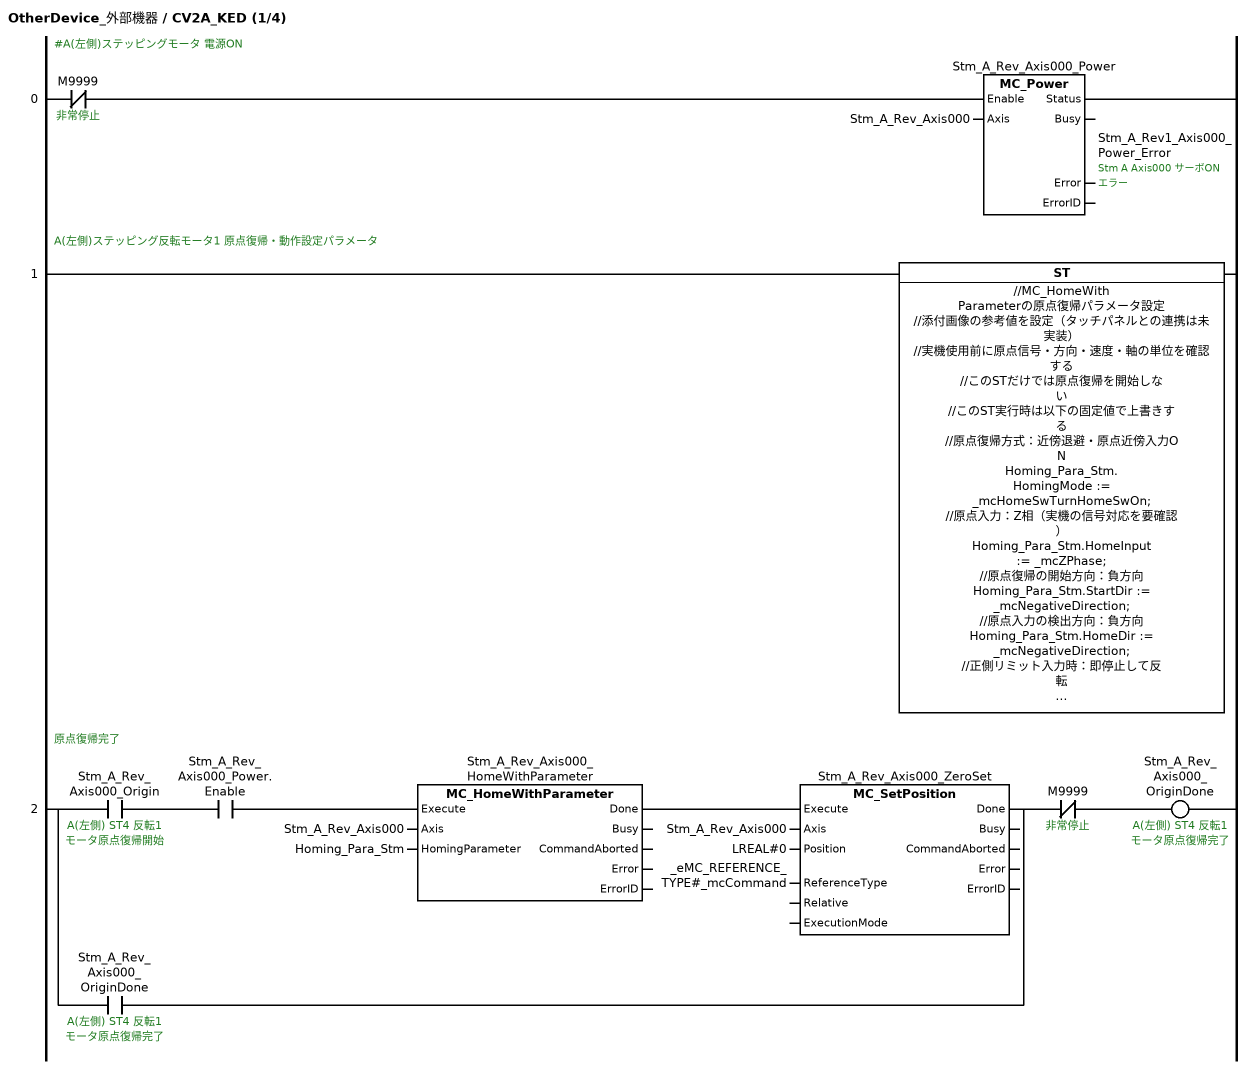
(* [picture p143: OtherDevice_外部機器 / CV2A_KED, rungs 0-2] *)
(* Rung 0: #A(左側)ステッピングモータ 電源ON *)
Stm_A_Rev_Axis000_Power(Enable := NOT M9999, Axis := Stm_A_Rev_Axis000, Error => Stm_A_Rev1_Axis000_Power_Error);
(* Rung 1: A(左側)ステッピング反転モータ1 原点復帰・動作設定パラメータ *)
//MC_HomeWithParameterの原点復帰パラメータ設定
//添付画像の参考値を設定（タッチパネルとの連携は未実装）
//実機使用前に原点信号・方向・速度・軸の単位を確認する
//このSTだけでは原点復帰を開始しない
//このST実行時は以下の固定値で上書きする

//原点復帰方式：近傍退避・原点近傍入力ON
Homing_Para_Stm.HomingMode := _mcHomeSwTurnHomeSwOn;
//原点入力：Z相（実機の信号対応を要確認）
Homing_Para_Stm.HomeInput := _mcZPhase;
//原点復帰の開始方向：負方向
Homing_Para_Stm.StartDir := _mcNegativeDirection;
//原点入力の検出方向：負方向
Homing_Para_Stm.HomeDir := _mcNegativeDirection;
//正側リミット入力時：即停止して反転
Homing_Para_Stm.PosiLmtMode := _mcRevImmediateStop;
//負側リミット入力時：即停止して反転
Homing_Para_Stm.NegaLmtMode := _mcRevImmediateStop;

//原点復帰速度 [指令単位/s]
Homing_Para_Stm.Vel := LREAL#40;
//原点近傍での接近速度 [指令単位/s]
Homing_Para_Stm.ApproachVel := LREAL#1;
//原点復帰の加速度 [指令単位/s^2]
Homing_Para_Stm.Acc := LREAL#100;
//原点復帰の減速度 [指令単位/s^2]
Homing_Para_Stm.Dec := LREAL#200;
//ジャーク [指令単位/s^3]：0はジャーク制御なし
Homing_Para_Stm.Jerk := LREAL#0;

//原点入力マスク距離 [指令単位]：今回の方式では未使用
Homing_Para_Stm.Mask := LREAL#0;
//原点確定後の現在位置 [指令単位]
Homing_Para_Stm.Offset := LREAL#0;
//押当て時間 [ms]：今回の方式では未使用
Homing_Para_Stm.PushTime := UINT#0;
//原点検出後の補正移動量 [指令単位]：0は補正移動なし
Homing_Para_Stm.Compensation := LREAL#0;
//原点補正移動時の速度 [指令単位/s]
Homing_Para_Stm.CompensationVel := LREAL#10;
(* Rung 2: 原点復帰完了 *)
Stm_A_Rev_Axis000_HomeWithParameter(Execute := Stm_A_Rev_Axis000_Origin AND Stm_A_Rev_Axis000_Power.Enable, Axis := Stm_A_Rev_Axis000, HomingParameter := Homing_Para_Stm);
Stm_A_Rev_Axis000_ZeroSet(Execute := Stm_A_Rev_Axis000_HomeWithParameter.Done, Axis := Stm_A_Rev_Axis000, Position := LREAL#0, ReferenceType := _eMC_REFERENCE_TYPE#_mcCommand);
Stm_A_Rev_Axis000_OriginDone := (Stm_A_Rev_Axis000_ZeroSet.Done OR Stm_A_Rev_Axis000_OriginDone) AND NOT M9999;

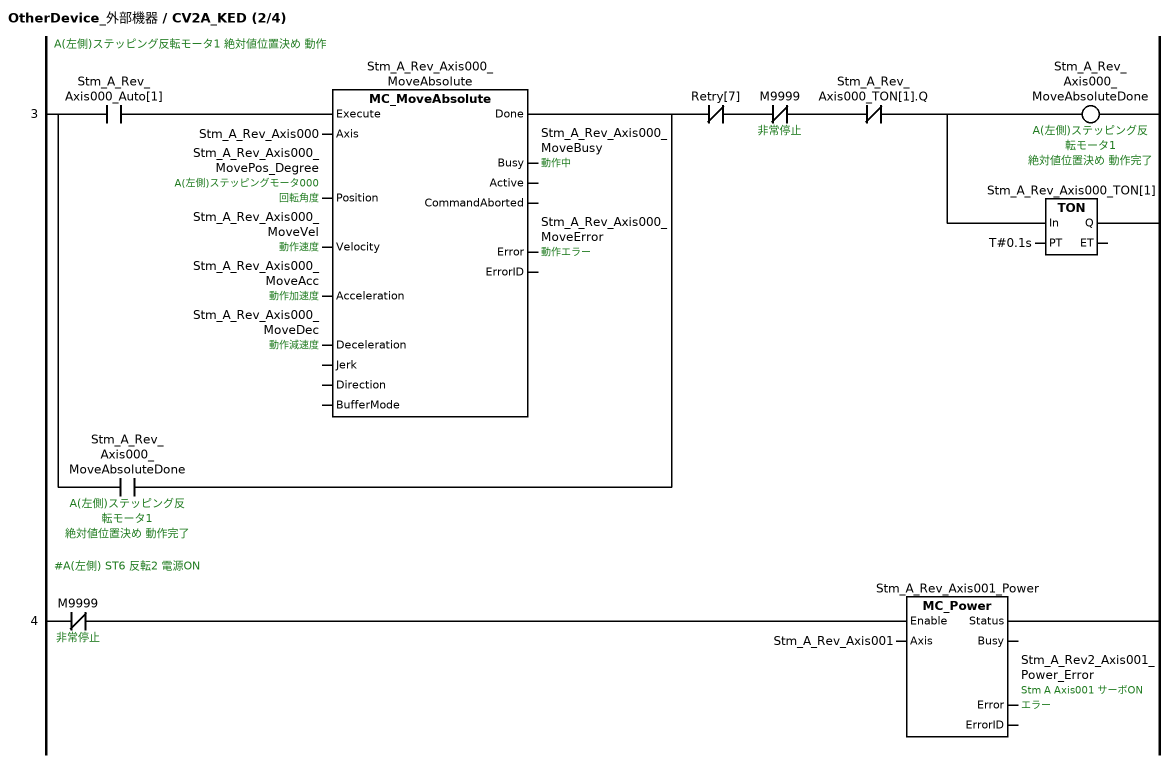
(* Rung 3: A(左側)ステッピング反転モータ1 絶対値位置決め 動作 *)
Stm_A_Rev_Axis000_MoveAbsolute(Execute := Stm_A_Rev_Axis000_Auto[1], Axis := Stm_A_Rev_Axis000, Position := Stm_A_Rev_Axis000_MovePos_Degree, Velocity := Stm_A_Rev_Axis000_MoveVel, Acceleration := Stm_A_Rev_Axis000_MoveAcc, Deceleration := Stm_A_Rev_Axis000_MoveDec, Busy => Stm_A_Rev_Axis000_MoveBusy, Error => Stm_A_Rev_Axis000_MoveError);
_p71 := (Stm_A_Rev_Axis000_MoveAbsolute.Done OR Stm_A_Rev_Axis000_MoveAbsoluteDone) AND NOT Retry[7] AND NOT M9999 AND NOT Stm_A_Rev_Axis000_TON[1].Q;
Stm_A_Rev_Axis000_MoveAbsoluteDone := _p71;
Stm_A_Rev_Axis000_TON[1](In := _p71, PT := T#0.1s);
(* Rung 4: #A(左側) ST6 反転2 電源ON *)
Stm_A_Rev_Axis001_Power(Enable := NOT M9999, Axis := Stm_A_Rev_Axis001, Error => Stm_A_Rev2_Axis001_Power_Error);

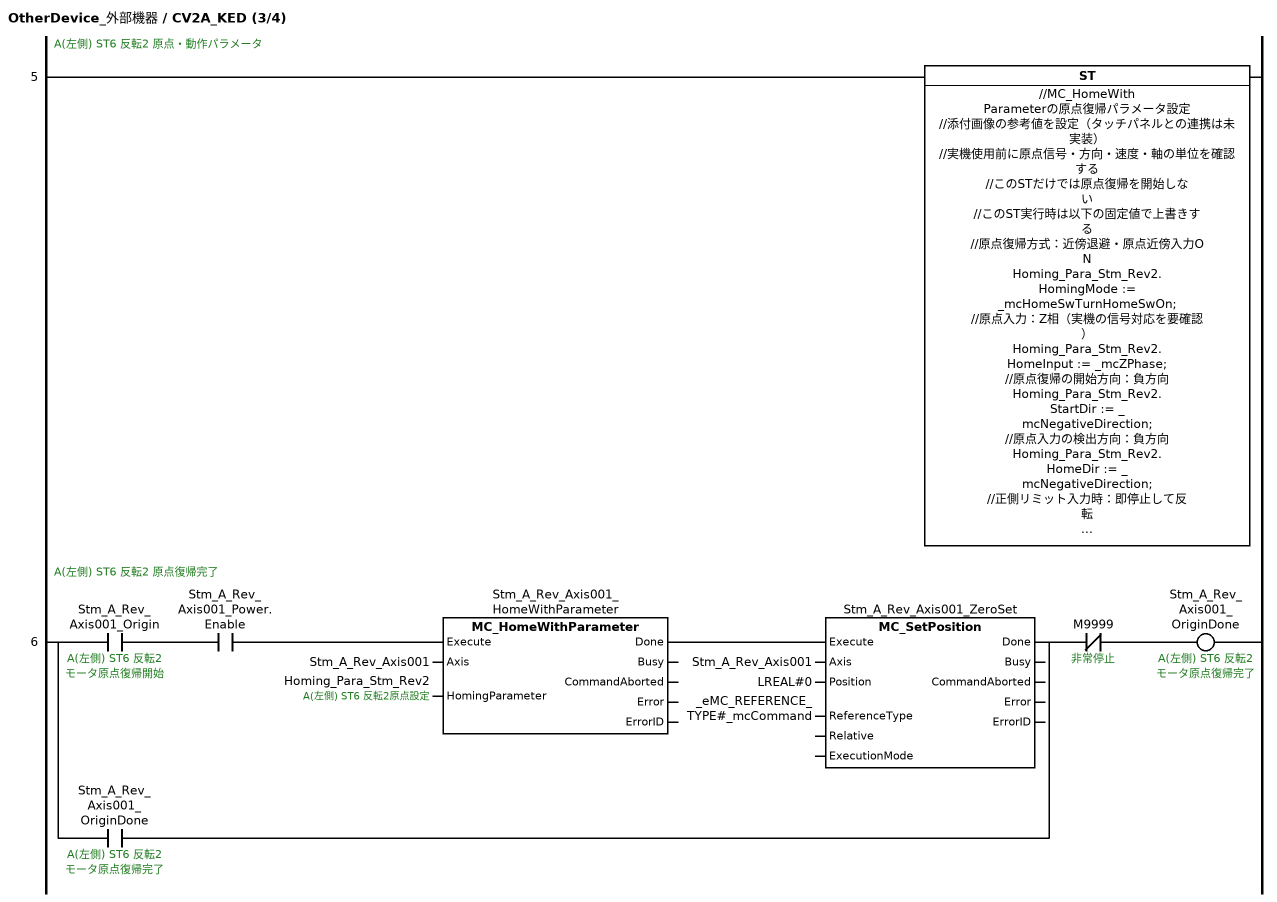
(* Rung 5: A(左側) ST6 反転2 原点・動作パラメータ *)
//MC_HomeWithParameterの原点復帰パラメータ設定
//添付画像の参考値を設定（タッチパネルとの連携は未実装）
//実機使用前に原点信号・方向・速度・軸の単位を確認する
//このSTだけでは原点復帰を開始しない
//このST実行時は以下の固定値で上書きする

//原点復帰方式：近傍退避・原点近傍入力ON
Homing_Para_Stm_Rev2.HomingMode := _mcHomeSwTurnHomeSwOn;
//原点入力：Z相（実機の信号対応を要確認）
Homing_Para_Stm_Rev2.HomeInput := _mcZPhase;
//原点復帰の開始方向：負方向
Homing_Para_Stm_Rev2.StartDir := _mcNegativeDirection;
//原点入力の検出方向：負方向
Homing_Para_Stm_Rev2.HomeDir := _mcNegativeDirection;
//正側リミット入力時：即停止して反転
Homing_Para_Stm_Rev2.PosiLmtMode := _mcRevImmediateStop;
//負側リミット入力時：即停止して反転
Homing_Para_Stm_Rev2.NegaLmtMode := _mcRevImmediateStop;

//原点復帰速度 [指令単位/s]
Homing_Para_Stm_Rev2.Vel := LREAL#40;
//原点近傍での接近速度 [指令単位/s]
Homing_Para_Stm_Rev2.ApproachVel := LREAL#1;
//原点復帰の加速度 [指令単位/s^2]
Homing_Para_Stm_Rev2.Acc := LREAL#100;
//原点復帰の減速度 [指令単位/s^2]
Homing_Para_Stm_Rev2.Dec := LREAL#200;
//ジャーク [指令単位/s^3]：0はジャーク制御なし
Homing_Para_Stm_Rev2.Jerk := LREAL#0;

//原点入力マスク距離 [指令単位]：今回の方式では未使用
Homing_Para_Stm_Rev2.Mask := LREAL#0;
//原点確定後の現在位置 [指令単位]
Homing_Para_Stm_Rev2.Offset := LREAL#0;
//押当て時間 [ms]：今回の方式では未使用
Homing_Para_Stm_Rev2.PushTime := UINT#0;
//原点検出後の補正移動量 [指令単位]：0は補正移動なし
Homing_Para_Stm_Rev2.Compensation := LREAL#0;
//原点補正移動時の速度 [指令単位/s]
Homing_Para_Stm_Rev2.CompensationVel := LREAL#10;
(* Rung 6: A(左側) ST6 反転2 原点復帰完了 *)
Stm_A_Rev_Axis001_HomeWithParameter(Execute := Stm_A_Rev_Axis001_Origin AND Stm_A_Rev_Axis001_Power.Enable, Axis := Stm_A_Rev_Axis001, HomingParameter := Homing_Para_Stm_Rev2);
Stm_A_Rev_Axis001_ZeroSet(Execute := Stm_A_Rev_Axis001_HomeWithParameter.Done, Axis := Stm_A_Rev_Axis001, Position := LREAL#0, ReferenceType := _eMC_REFERENCE_TYPE#_mcCommand);
Stm_A_Rev_Axis001_OriginDone := (Stm_A_Rev_Axis001_ZeroSet.Done OR Stm_A_Rev_Axis001_OriginDone) AND NOT M9999;

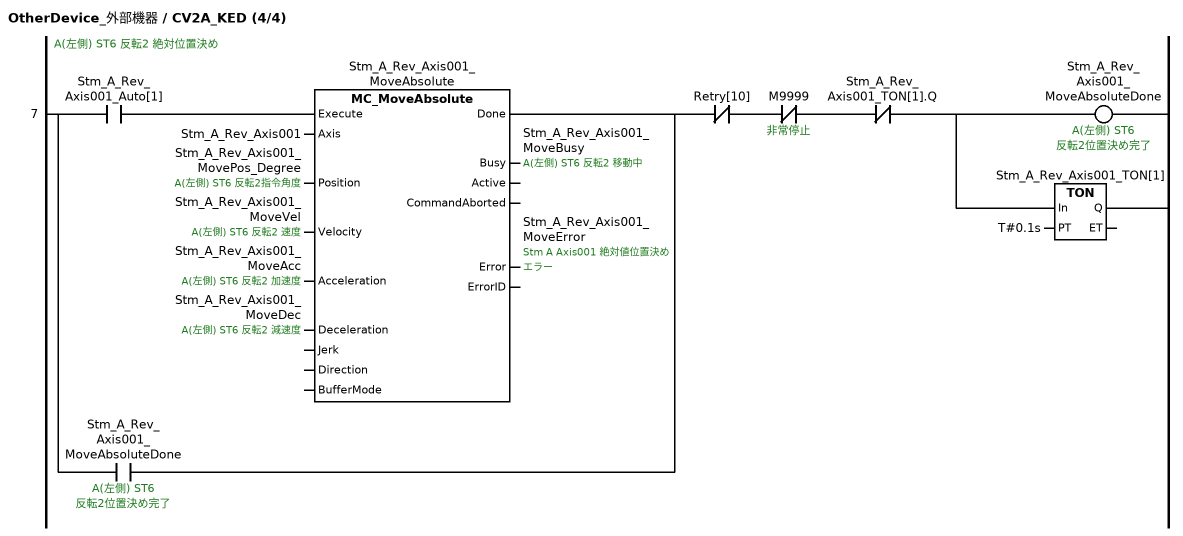
(* Rung 7: A(左側) ST6 反転2 絶対位置決め *)
Stm_A_Rev_Axis001_MoveAbsolute(Execute := Stm_A_Rev_Axis001_Auto[1], Axis := Stm_A_Rev_Axis001, Position := Stm_A_Rev_Axis001_MovePos_Degree, Velocity := Stm_A_Rev_Axis001_MoveVel, Acceleration := Stm_A_Rev_Axis001_MoveAcc, Deceleration := Stm_A_Rev_Axis001_MoveDec, Busy => Stm_A_Rev_Axis001_MoveBusy, Error => Stm_A_Rev_Axis001_MoveError);
_p72 := (Stm_A_Rev_Axis001_MoveAbsolute.Done OR Stm_A_Rev_Axis001_MoveAbsoluteDone) AND NOT Retry[10] AND NOT M9999 AND NOT Stm_A_Rev_Axis001_TON[1].Q;
Stm_A_Rev_Axis001_MoveAbsoluteDone := _p72;
Stm_A_Rev_Axis001_TON[1](In := _p72, PT := T#0.1s);

(* Section HMI: ladder, written here as Structured Text *)

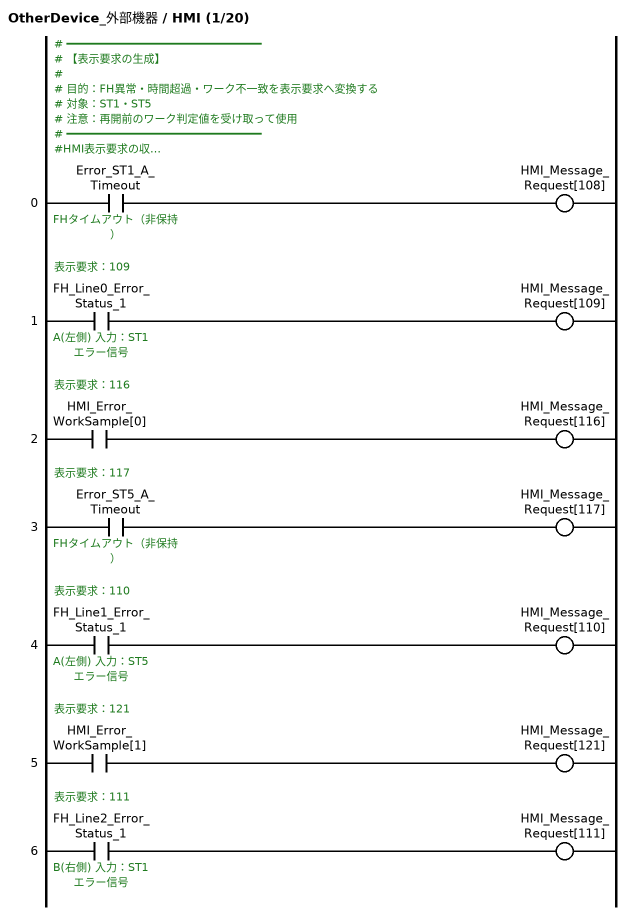
(* Rung 0: # ━━━━━━━━━━━━━━━━━━━━━━━━━━━━━━ / # 【表示要求の生成】 / # / # 目的：FH異常・時間超過・ワーク不一致を表示要求へ変換する / # 対象：ST1・ST5 / # 注意：再開前のワーク判定値を受け取って使用 / # ━━━━━━━━━━━━━━━━━━━━━━━━━━━━━━ / #HMI表示要求の収集 / 実行順維持のため、異常判定後・再開処理前 / 表示要求：108 *)
HMI_Message_Request[108] := Error_ST1_A_Timeout;
(* Rung 1: 表示要求：109 *)
HMI_Message_Request[109] := FH_Line0_Error_Status_1;
(* Rung 2: 表示要求：116 *)
HMI_Message_Request[116] := HMI_Error_WorkSample[0];
(* Rung 3: 表示要求：117 *)
HMI_Message_Request[117] := Error_ST5_A_Timeout;
(* Rung 4: 表示要求：110 *)
HMI_Message_Request[110] := FH_Line1_Error_Status_1;
(* Rung 5: 表示要求：121 *)
HMI_Message_Request[121] := HMI_Error_WorkSample[1];
(* Rung 6: 表示要求：111 *)
HMI_Message_Request[111] := FH_Line2_Error_Status_1;

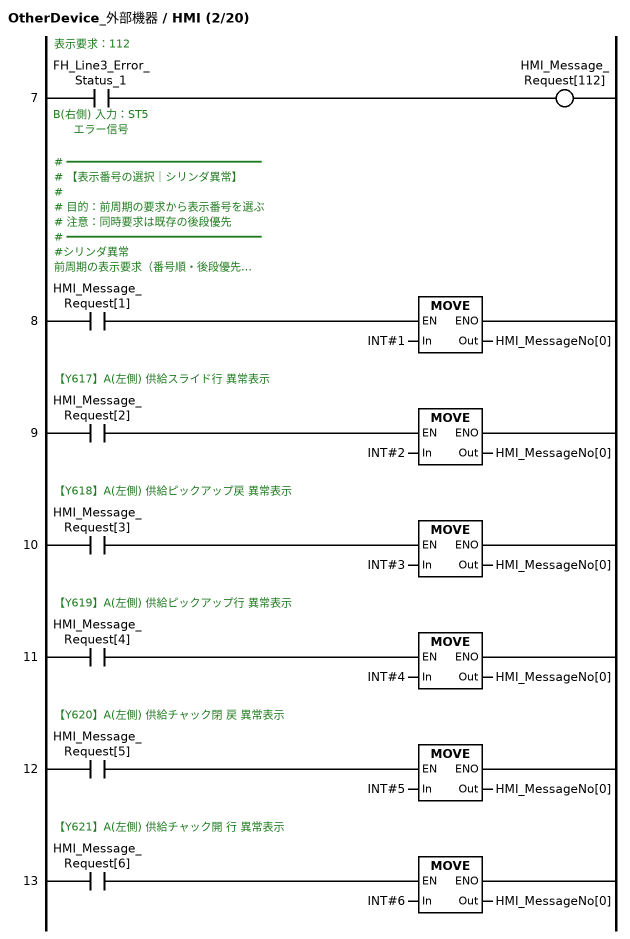
(* Rung 7: 表示要求：112 *)
HMI_Message_Request[112] := FH_Line3_Error_Status_1;
(* Rung 8: # ━━━━━━━━━━━━━━━━━━━━━━━━━━━━━━ / # 【表示番号の選択｜シリンダ異常】 / # / # 目的：前周期の要求から表示番号を選ぶ / # 注意：同時要求は既存の後段優先 / # ━━━━━━━━━━━━━━━━━━━━━━━━━━━━━━ / #シリンダ異常 / 前周期の表示要求（番号順・後段優先） / 【Y616】A(左側) 供給スライド戻 異常表示 *)
IF HMI_Message_Request[1] THEN HMI_MessageNo[0] := INT#1; END_IF;
(* Rung 9: 【Y617】A(左側) 供給スライド行 異常表示 *)
IF HMI_Message_Request[2] THEN HMI_MessageNo[0] := INT#2; END_IF;
(* Rung 10: 【Y618】A(左側) 供給ピックアップ戻 異常表示 *)
IF HMI_Message_Request[3] THEN HMI_MessageNo[0] := INT#3; END_IF;
(* Rung 11: 【Y619】A(左側) 供給ピックアップ行 異常表示 *)
IF HMI_Message_Request[4] THEN HMI_MessageNo[0] := INT#4; END_IF;
(* Rung 12: 【Y620】A(左側) 供給チャック閉 戻 異常表示 *)
IF HMI_Message_Request[5] THEN HMI_MessageNo[0] := INT#5; END_IF;
(* Rung 13: 【Y621】A(左側) 供給チャック開 行 異常表示 *)
IF HMI_Message_Request[6] THEN HMI_MessageNo[0] := INT#6; END_IF;

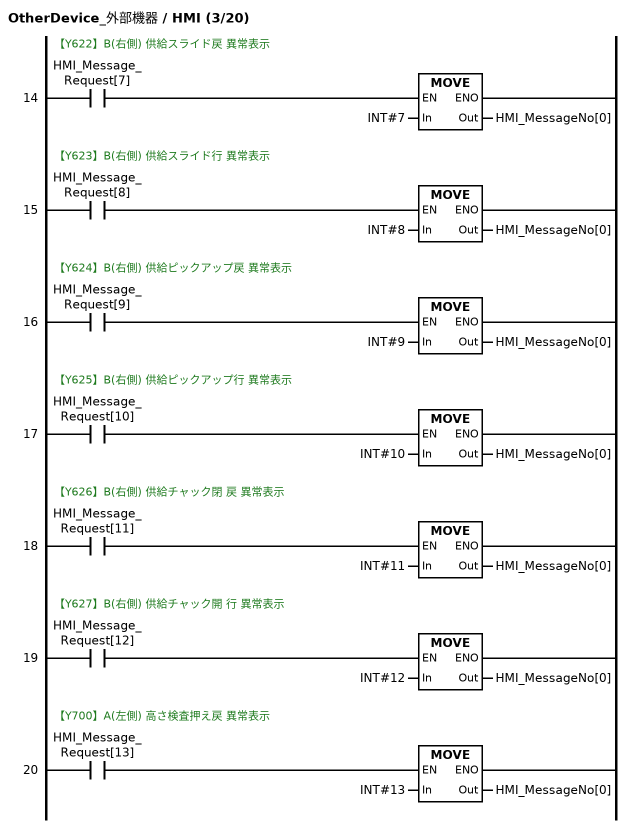
(* Rung 14: 【Y622】B(右側) 供給スライド戻 異常表示 *)
IF HMI_Message_Request[7] THEN HMI_MessageNo[0] := INT#7; END_IF;
(* Rung 15: 【Y623】B(右側) 供給スライド行 異常表示 *)
IF HMI_Message_Request[8] THEN HMI_MessageNo[0] := INT#8; END_IF;
(* Rung 16: 【Y624】B(右側) 供給ピックアップ戻 異常表示 *)
IF HMI_Message_Request[9] THEN HMI_MessageNo[0] := INT#9; END_IF;
(* Rung 17: 【Y625】B(右側) 供給ピックアップ行 異常表示 *)
IF HMI_Message_Request[10] THEN HMI_MessageNo[0] := INT#10; END_IF;
(* Rung 18: 【Y626】B(右側) 供給チャック閉 戻 異常表示 *)
IF HMI_Message_Request[11] THEN HMI_MessageNo[0] := INT#11; END_IF;
(* Rung 19: 【Y627】B(右側) 供給チャック開 行 異常表示 *)
IF HMI_Message_Request[12] THEN HMI_MessageNo[0] := INT#12; END_IF;
(* Rung 20: 【Y700】A(左側) 高さ検査押え戻 異常表示 *)
IF HMI_Message_Request[13] THEN HMI_MessageNo[0] := INT#13; END_IF;

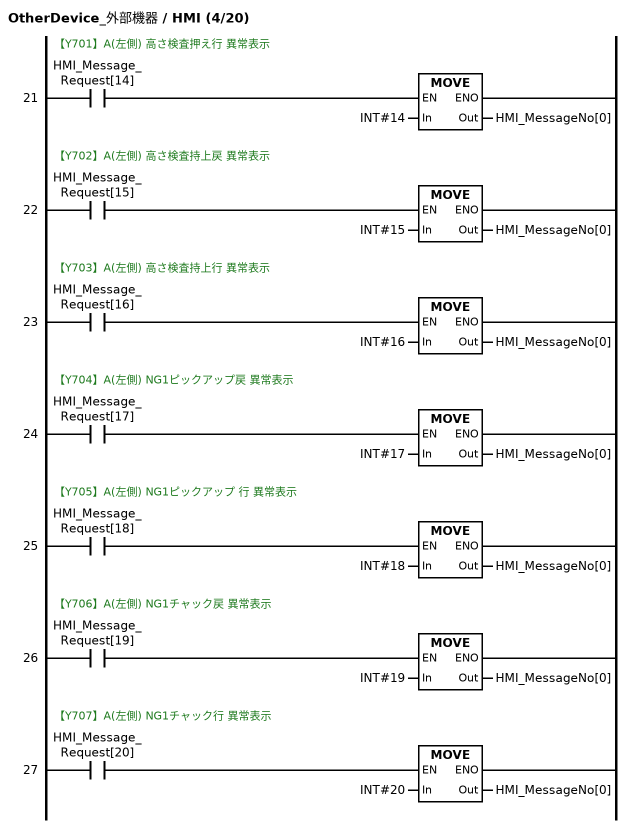
(* Rung 21: 【Y701】A(左側) 高さ検査押え行 異常表示 *)
IF HMI_Message_Request[14] THEN HMI_MessageNo[0] := INT#14; END_IF;
(* Rung 22: 【Y702】A(左側) 高さ検査持上戻 異常表示 *)
IF HMI_Message_Request[15] THEN HMI_MessageNo[0] := INT#15; END_IF;
(* Rung 23: 【Y703】A(左側) 高さ検査持上行 異常表示 *)
IF HMI_Message_Request[16] THEN HMI_MessageNo[0] := INT#16; END_IF;
(* Rung 24: 【Y704】A(左側) NG1ピックアップ戻 異常表示 *)
IF HMI_Message_Request[17] THEN HMI_MessageNo[0] := INT#17; END_IF;
(* Rung 25: 【Y705】A(左側) NG1ピックアップ 行 異常表示 *)
IF HMI_Message_Request[18] THEN HMI_MessageNo[0] := INT#18; END_IF;
(* Rung 26: 【Y706】A(左側) NG1チャック戻 異常表示 *)
IF HMI_Message_Request[19] THEN HMI_MessageNo[0] := INT#19; END_IF;
(* Rung 27: 【Y707】A(左側) NG1チャック行 異常表示 *)
IF HMI_Message_Request[20] THEN HMI_MessageNo[0] := INT#20; END_IF;

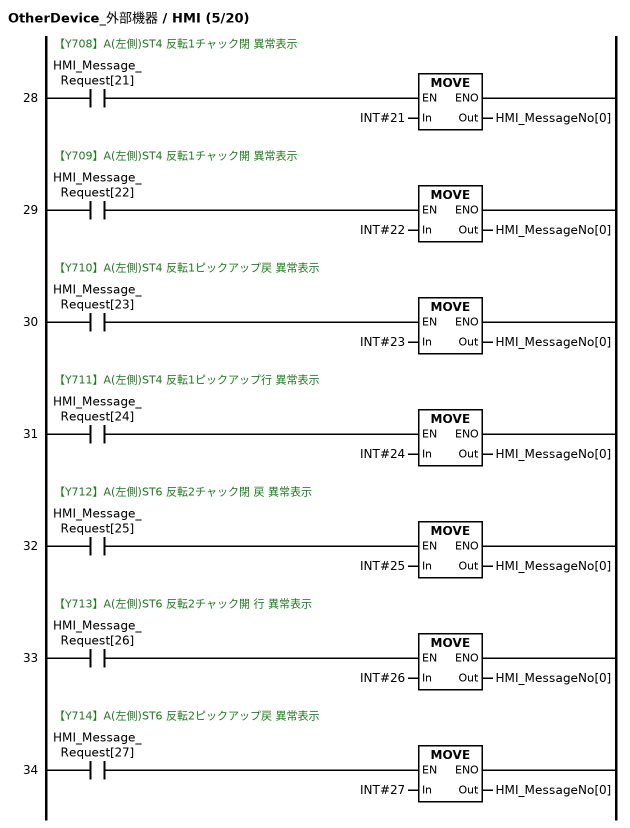
(* Rung 28: 【Y708】A(左側)ST4 反転1チャック閉 異常表示 *)
IF HMI_Message_Request[21] THEN HMI_MessageNo[0] := INT#21; END_IF;
(* Rung 29: 【Y709】A(左側)ST4 反転1チャック開 異常表示 *)
IF HMI_Message_Request[22] THEN HMI_MessageNo[0] := INT#22; END_IF;
(* Rung 30: 【Y710】A(左側)ST4 反転1ピックアップ戻 異常表示 *)
IF HMI_Message_Request[23] THEN HMI_MessageNo[0] := INT#23; END_IF;
(* Rung 31: 【Y711】A(左側)ST4 反転1ピックアップ行 異常表示 *)
IF HMI_Message_Request[24] THEN HMI_MessageNo[0] := INT#24; END_IF;
(* Rung 32: 【Y712】A(左側)ST6 反転2チャック閉 戻 異常表示 *)
IF HMI_Message_Request[25] THEN HMI_MessageNo[0] := INT#25; END_IF;
(* Rung 33: 【Y713】A(左側)ST6 反転2チャック開 行 異常表示 *)
IF HMI_Message_Request[26] THEN HMI_MessageNo[0] := INT#26; END_IF;
(* Rung 34: 【Y714】A(左側)ST6 反転2ピックアップ戻 異常表示 *)
IF HMI_Message_Request[27] THEN HMI_MessageNo[0] := INT#27; END_IF;

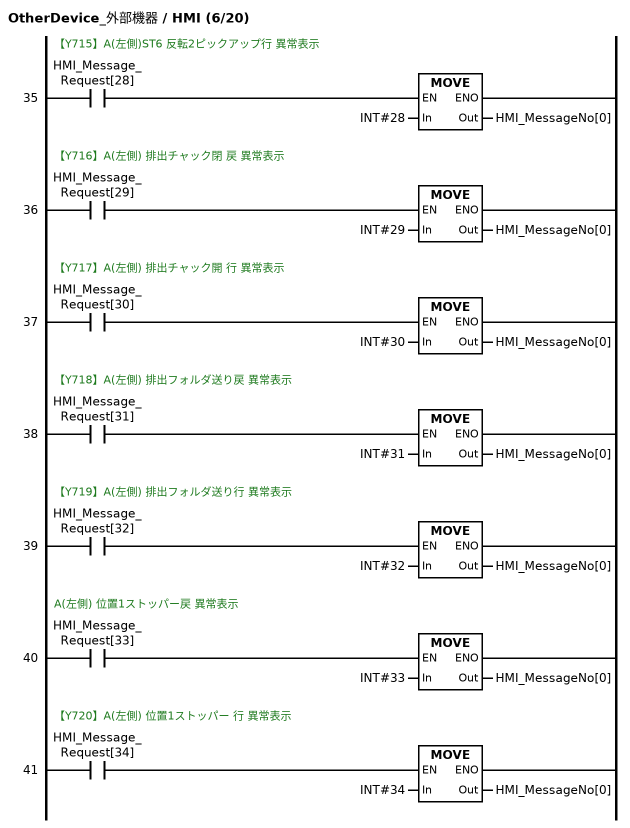
(* Rung 35: 【Y715】A(左側)ST6 反転2ピックアップ行 異常表示 *)
IF HMI_Message_Request[28] THEN HMI_MessageNo[0] := INT#28; END_IF;
(* Rung 36: 【Y716】A(左側) 排出チャック閉 戻 異常表示 *)
IF HMI_Message_Request[29] THEN HMI_MessageNo[0] := INT#29; END_IF;
(* Rung 37: 【Y717】A(左側) 排出チャック開 行 異常表示 *)
IF HMI_Message_Request[30] THEN HMI_MessageNo[0] := INT#30; END_IF;
(* Rung 38: 【Y718】A(左側) 排出フォルダ送り戻 異常表示 *)
IF HMI_Message_Request[31] THEN HMI_MessageNo[0] := INT#31; END_IF;
(* Rung 39: 【Y719】A(左側) 排出フォルダ送り行 異常表示 *)
IF HMI_Message_Request[32] THEN HMI_MessageNo[0] := INT#32; END_IF;
(* Rung 40: A(左側) 位置1ストッパー戻 異常表示 *)
IF HMI_Message_Request[33] THEN HMI_MessageNo[0] := INT#33; END_IF;
(* Rung 41: 【Y720】A(左側) 位置1ストッパー 行 異常表示 *)
IF HMI_Message_Request[34] THEN HMI_MessageNo[0] := INT#34; END_IF;

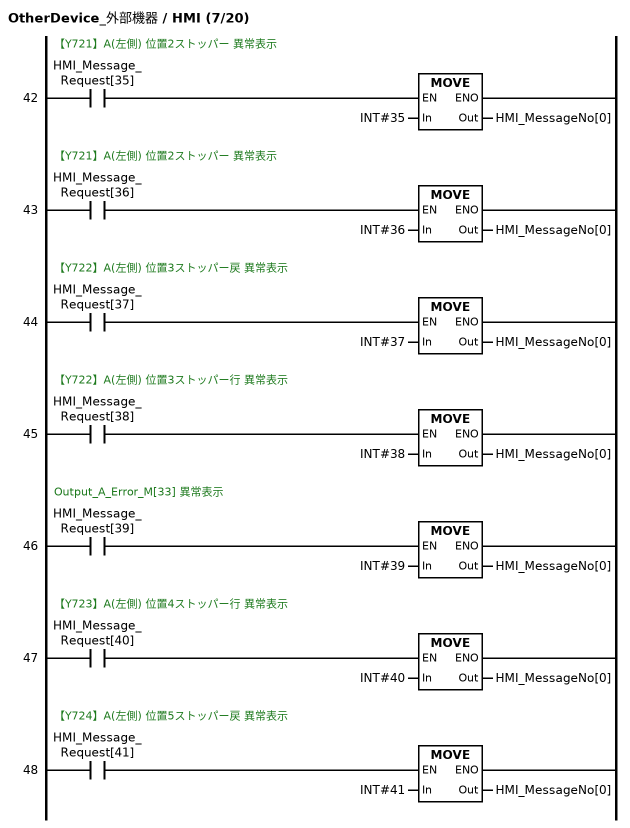
(* Rung 42: 【Y721】A(左側) 位置2ストッパー 異常表示 *)
IF HMI_Message_Request[35] THEN HMI_MessageNo[0] := INT#35; END_IF;
(* Rung 43: 【Y721】A(左側) 位置2ストッパー 異常表示 *)
IF HMI_Message_Request[36] THEN HMI_MessageNo[0] := INT#36; END_IF;
(* Rung 44: 【Y722】A(左側) 位置3ストッパー戻 異常表示 *)
IF HMI_Message_Request[37] THEN HMI_MessageNo[0] := INT#37; END_IF;
(* Rung 45: 【Y722】A(左側) 位置3ストッパー行 異常表示 *)
IF HMI_Message_Request[38] THEN HMI_MessageNo[0] := INT#38; END_IF;
(* Rung 46: Output_A_Error_M[33] 異常表示 *)
IF HMI_Message_Request[39] THEN HMI_MessageNo[0] := INT#39; END_IF;
(* Rung 47: 【Y723】A(左側) 位置4ストッパー行 異常表示 *)
IF HMI_Message_Request[40] THEN HMI_MessageNo[0] := INT#40; END_IF;
(* Rung 48: 【Y724】A(左側) 位置5ストッパー戻 異常表示 *)
IF HMI_Message_Request[41] THEN HMI_MessageNo[0] := INT#41; END_IF;

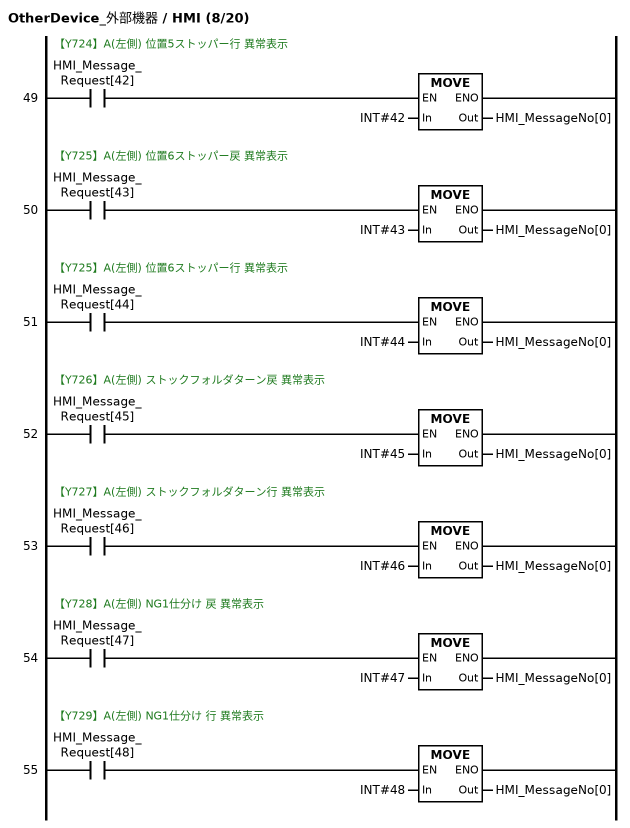
(* Rung 49: 【Y724】A(左側) 位置5ストッパー行 異常表示 *)
IF HMI_Message_Request[42] THEN HMI_MessageNo[0] := INT#42; END_IF;
(* Rung 50: 【Y725】A(左側) 位置6ストッパー戻 異常表示 *)
IF HMI_Message_Request[43] THEN HMI_MessageNo[0] := INT#43; END_IF;
(* Rung 51: 【Y725】A(左側) 位置6ストッパー行 異常表示 *)
IF HMI_Message_Request[44] THEN HMI_MessageNo[0] := INT#44; END_IF;
(* Rung 52: 【Y726】A(左側) ストックフォルダターン戻 異常表示 *)
IF HMI_Message_Request[45] THEN HMI_MessageNo[0] := INT#45; END_IF;
(* Rung 53: 【Y727】A(左側) ストックフォルダターン行 異常表示 *)
IF HMI_Message_Request[46] THEN HMI_MessageNo[0] := INT#46; END_IF;
(* Rung 54: 【Y728】A(左側) NG1仕分け 戻 異常表示 *)
IF HMI_Message_Request[47] THEN HMI_MessageNo[0] := INT#47; END_IF;
(* Rung 55: 【Y729】A(左側) NG1仕分け 行 異常表示 *)
IF HMI_Message_Request[48] THEN HMI_MessageNo[0] := INT#48; END_IF;

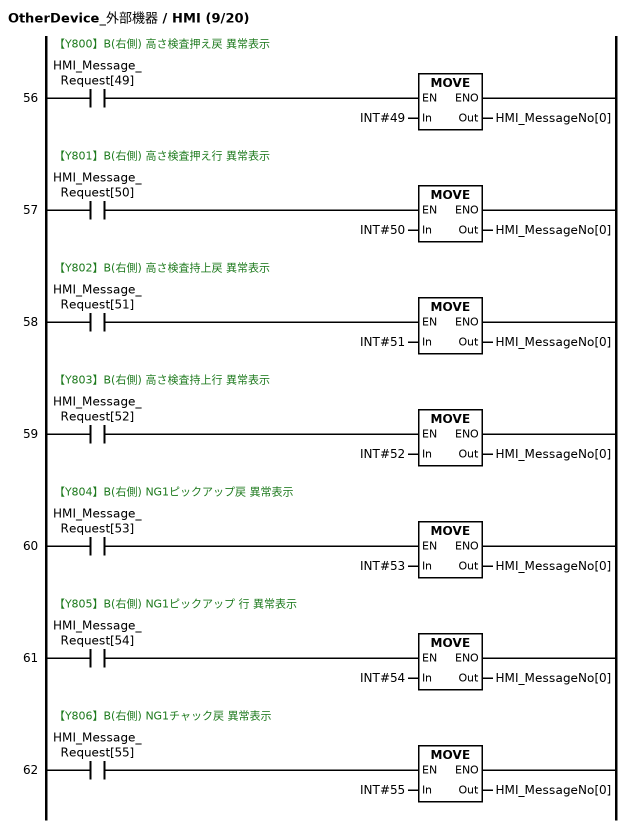
(* Rung 56: 【Y800】B(右側) 高さ検査押え戻 異常表示 *)
IF HMI_Message_Request[49] THEN HMI_MessageNo[0] := INT#49; END_IF;
(* Rung 57: 【Y801】B(右側) 高さ検査押え行 異常表示 *)
IF HMI_Message_Request[50] THEN HMI_MessageNo[0] := INT#50; END_IF;
(* Rung 58: 【Y802】B(右側) 高さ検査持上戻 異常表示 *)
IF HMI_Message_Request[51] THEN HMI_MessageNo[0] := INT#51; END_IF;
(* Rung 59: 【Y803】B(右側) 高さ検査持上行 異常表示 *)
IF HMI_Message_Request[52] THEN HMI_MessageNo[0] := INT#52; END_IF;
(* Rung 60: 【Y804】B(右側) NG1ピックアップ戻 異常表示 *)
IF HMI_Message_Request[53] THEN HMI_MessageNo[0] := INT#53; END_IF;
(* Rung 61: 【Y805】B(右側) NG1ピックアップ 行 異常表示 *)
IF HMI_Message_Request[54] THEN HMI_MessageNo[0] := INT#54; END_IF;
(* Rung 62: 【Y806】B(右側) NG1チャック戻 異常表示 *)
IF HMI_Message_Request[55] THEN HMI_MessageNo[0] := INT#55; END_IF;

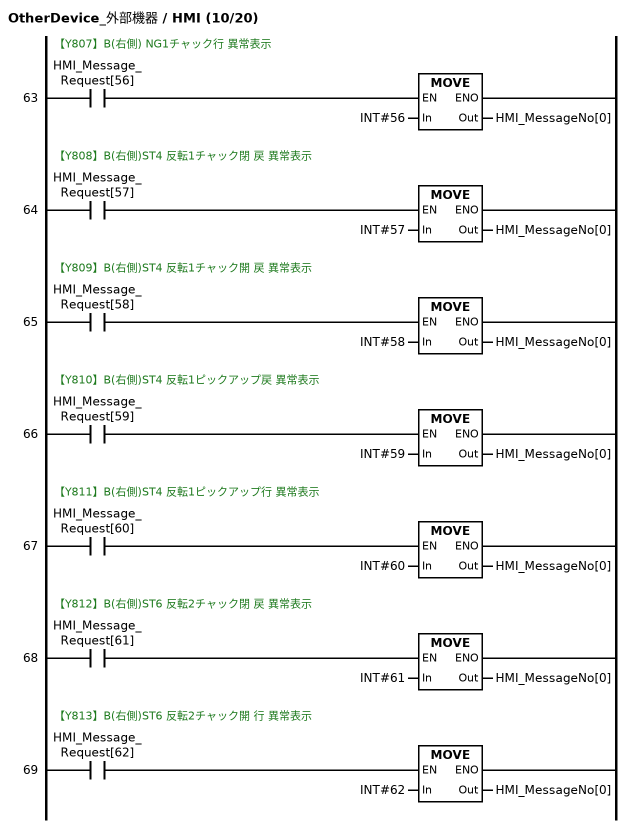
(* Rung 63: 【Y807】B(右側) NG1チャック行 異常表示 *)
IF HMI_Message_Request[56] THEN HMI_MessageNo[0] := INT#56; END_IF;
(* Rung 64: 【Y808】B(右側)ST4 反転1チャック閉 戻 異常表示 *)
IF HMI_Message_Request[57] THEN HMI_MessageNo[0] := INT#57; END_IF;
(* Rung 65: 【Y809】B(右側)ST4 反転1チャック開 戻 異常表示 *)
IF HMI_Message_Request[58] THEN HMI_MessageNo[0] := INT#58; END_IF;
(* Rung 66: 【Y810】B(右側)ST4 反転1ピックアップ戻 異常表示 *)
IF HMI_Message_Request[59] THEN HMI_MessageNo[0] := INT#59; END_IF;
(* Rung 67: 【Y811】B(右側)ST4 反転1ピックアップ行 異常表示 *)
IF HMI_Message_Request[60] THEN HMI_MessageNo[0] := INT#60; END_IF;
(* Rung 68: 【Y812】B(右側)ST6 反転2チャック閉 戻 異常表示 *)
IF HMI_Message_Request[61] THEN HMI_MessageNo[0] := INT#61; END_IF;
(* Rung 69: 【Y813】B(右側)ST6 反転2チャック開 行 異常表示 *)
IF HMI_Message_Request[62] THEN HMI_MessageNo[0] := INT#62; END_IF;

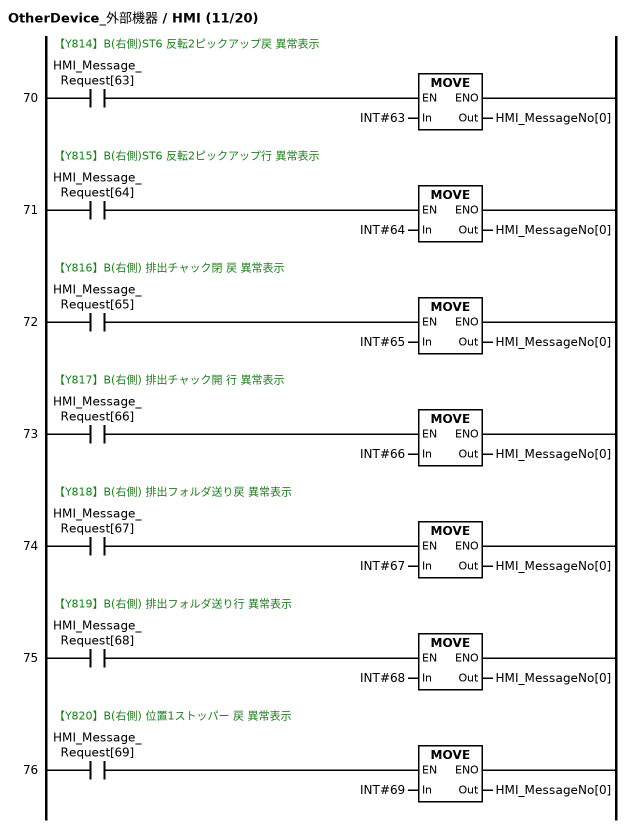
(* Rung 70: 【Y814】B(右側)ST6 反転2ピックアップ戻 異常表示 *)
IF HMI_Message_Request[63] THEN HMI_MessageNo[0] := INT#63; END_IF;
(* Rung 71: 【Y815】B(右側)ST6 反転2ピックアップ行 異常表示 *)
IF HMI_Message_Request[64] THEN HMI_MessageNo[0] := INT#64; END_IF;
(* Rung 72: 【Y816】B(右側) 排出チャック閉 戻 異常表示 *)
IF HMI_Message_Request[65] THEN HMI_MessageNo[0] := INT#65; END_IF;
(* Rung 73: 【Y817】B(右側) 排出チャック開 行 異常表示 *)
IF HMI_Message_Request[66] THEN HMI_MessageNo[0] := INT#66; END_IF;
(* Rung 74: 【Y818】B(右側) 排出フォルダ送り戻 異常表示 *)
IF HMI_Message_Request[67] THEN HMI_MessageNo[0] := INT#67; END_IF;
(* Rung 75: 【Y819】B(右側) 排出フォルダ送り行 異常表示 *)
IF HMI_Message_Request[68] THEN HMI_MessageNo[0] := INT#68; END_IF;
(* Rung 76: 【Y820】B(右側) 位置1ストッパー 戻 異常表示 *)
IF HMI_Message_Request[69] THEN HMI_MessageNo[0] := INT#69; END_IF;

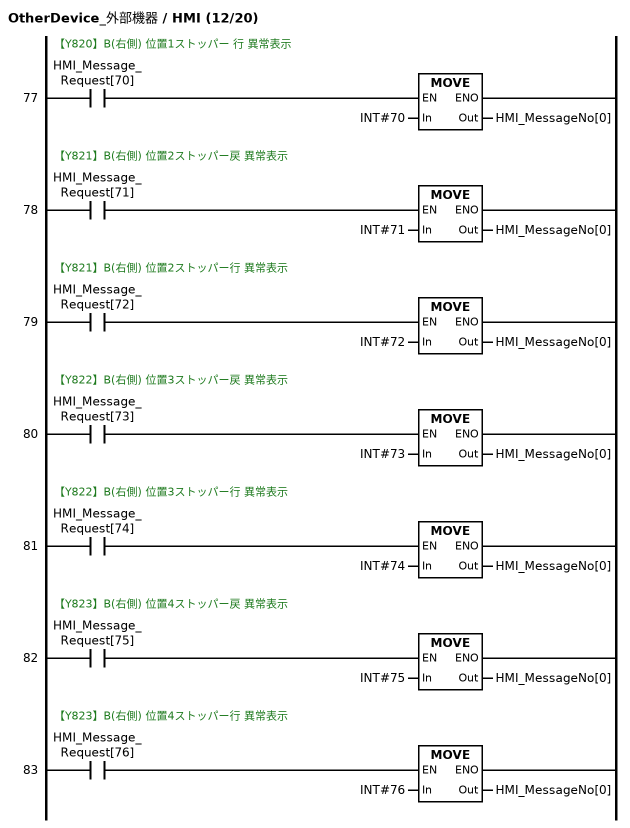
(* Rung 77: 【Y820】B(右側) 位置1ストッパー 行 異常表示 *)
IF HMI_Message_Request[70] THEN HMI_MessageNo[0] := INT#70; END_IF;
(* Rung 78: 【Y821】B(右側) 位置2ストッパー戻 異常表示 *)
IF HMI_Message_Request[71] THEN HMI_MessageNo[0] := INT#71; END_IF;
(* Rung 79: 【Y821】B(右側) 位置2ストッパー行 異常表示 *)
IF HMI_Message_Request[72] THEN HMI_MessageNo[0] := INT#72; END_IF;
(* Rung 80: 【Y822】B(右側) 位置3ストッパー戻 異常表示 *)
IF HMI_Message_Request[73] THEN HMI_MessageNo[0] := INT#73; END_IF;
(* Rung 81: 【Y822】B(右側) 位置3ストッパー行 異常表示 *)
IF HMI_Message_Request[74] THEN HMI_MessageNo[0] := INT#74; END_IF;
(* Rung 82: 【Y823】B(右側) 位置4ストッパー戻 異常表示 *)
IF HMI_Message_Request[75] THEN HMI_MessageNo[0] := INT#75; END_IF;
(* Rung 83: 【Y823】B(右側) 位置4ストッパー行 異常表示 *)
IF HMI_Message_Request[76] THEN HMI_MessageNo[0] := INT#76; END_IF;

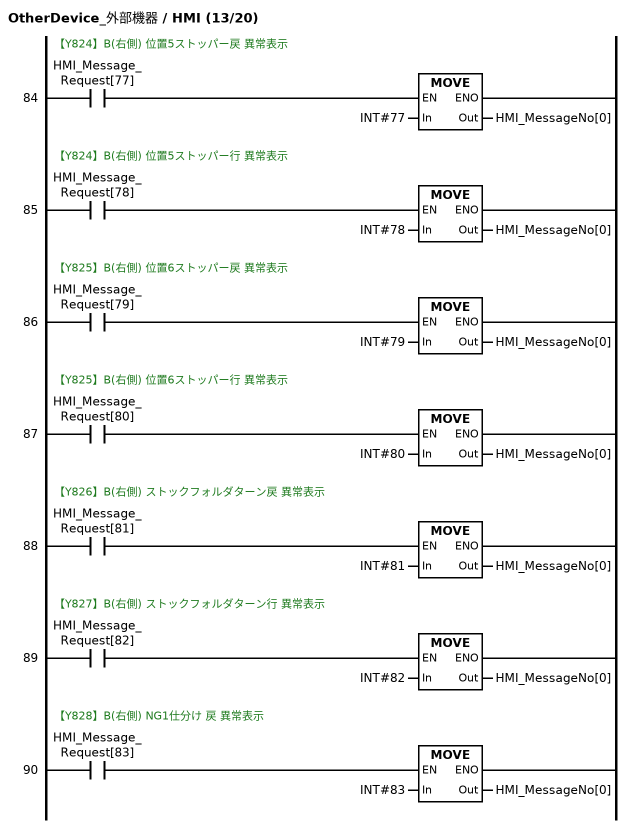
(* Rung 84: 【Y824】B(右側) 位置5ストッパー戻 異常表示 *)
IF HMI_Message_Request[77] THEN HMI_MessageNo[0] := INT#77; END_IF;
(* Rung 85: 【Y824】B(右側) 位置5ストッパー行 異常表示 *)
IF HMI_Message_Request[78] THEN HMI_MessageNo[0] := INT#78; END_IF;
(* Rung 86: 【Y825】B(右側) 位置6ストッパー戻 異常表示 *)
IF HMI_Message_Request[79] THEN HMI_MessageNo[0] := INT#79; END_IF;
(* Rung 87: 【Y825】B(右側) 位置6ストッパー行 異常表示 *)
IF HMI_Message_Request[80] THEN HMI_MessageNo[0] := INT#80; END_IF;
(* Rung 88: 【Y826】B(右側) ストックフォルダターン戻 異常表示 *)
IF HMI_Message_Request[81] THEN HMI_MessageNo[0] := INT#81; END_IF;
(* Rung 89: 【Y827】B(右側) ストックフォルダターン行 異常表示 *)
IF HMI_Message_Request[82] THEN HMI_MessageNo[0] := INT#82; END_IF;
(* Rung 90: 【Y828】B(右側) NG1仕分け 戻 異常表示 *)
IF HMI_Message_Request[83] THEN HMI_MessageNo[0] := INT#83; END_IF;

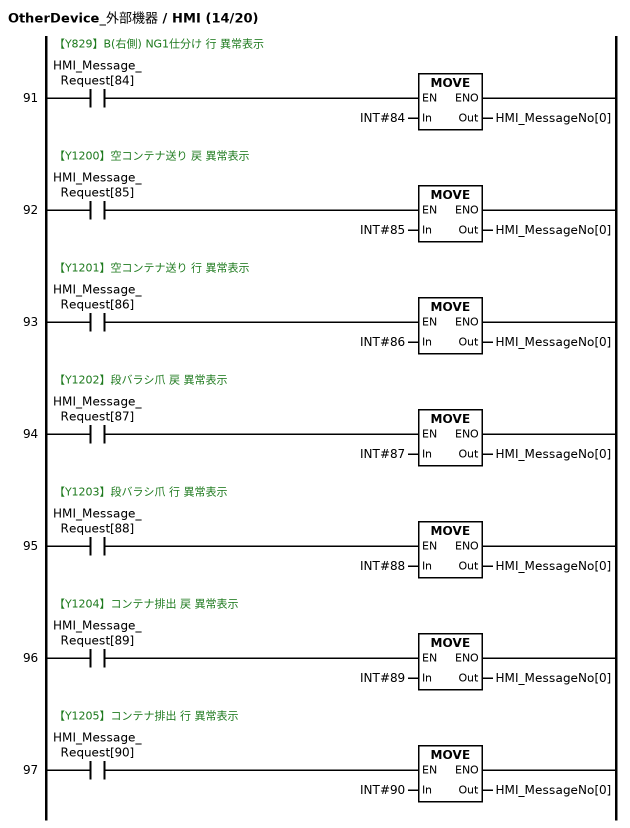
(* Rung 91: 【Y829】B(右側) NG1仕分け 行 異常表示 *)
IF HMI_Message_Request[84] THEN HMI_MessageNo[0] := INT#84; END_IF;
(* Rung 92: 【Y1200】空コンテナ送り 戻 異常表示 *)
IF HMI_Message_Request[85] THEN HMI_MessageNo[0] := INT#85; END_IF;
(* Rung 93: 【Y1201】空コンテナ送り 行 異常表示 *)
IF HMI_Message_Request[86] THEN HMI_MessageNo[0] := INT#86; END_IF;
(* Rung 94: 【Y1202】段バラシ爪 戻 異常表示 *)
IF HMI_Message_Request[87] THEN HMI_MessageNo[0] := INT#87; END_IF;
(* Rung 95: 【Y1203】段バラシ爪 行 異常表示 *)
IF HMI_Message_Request[88] THEN HMI_MessageNo[0] := INT#88; END_IF;
(* Rung 96: 【Y1204】コンテナ排出 戻 異常表示 *)
IF HMI_Message_Request[89] THEN HMI_MessageNo[0] := INT#89; END_IF;
(* Rung 97: 【Y1205】コンテナ排出 行 異常表示 *)
IF HMI_Message_Request[90] THEN HMI_MessageNo[0] := INT#90; END_IF;

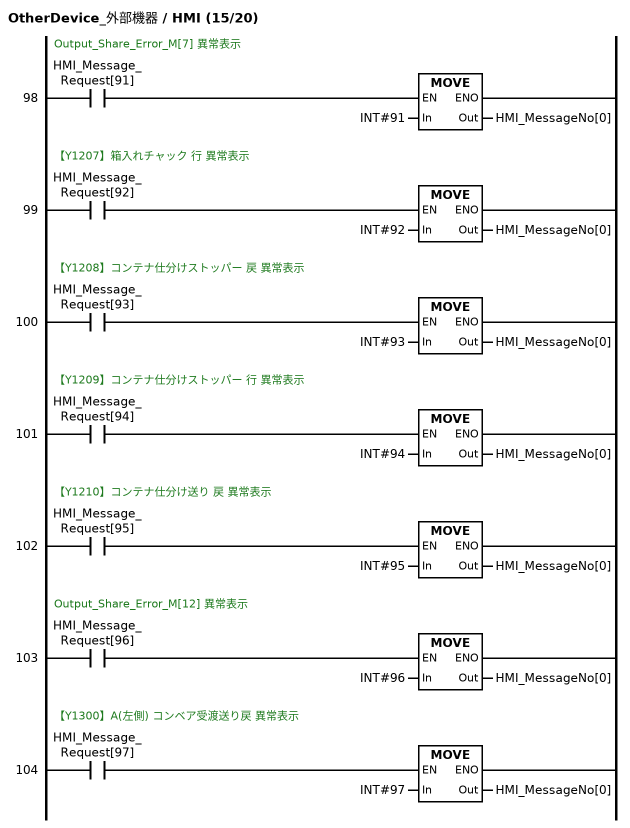
(* Rung 98: Output_Share_Error_M[7] 異常表示 *)
IF HMI_Message_Request[91] THEN HMI_MessageNo[0] := INT#91; END_IF;
(* Rung 99: 【Y1207】箱入れチャック 行 異常表示 *)
IF HMI_Message_Request[92] THEN HMI_MessageNo[0] := INT#92; END_IF;
(* Rung 100: 【Y1208】コンテナ仕分けストッパー 戻 異常表示 *)
IF HMI_Message_Request[93] THEN HMI_MessageNo[0] := INT#93; END_IF;
(* Rung 101: 【Y1209】コンテナ仕分けストッパー 行 異常表示 *)
IF HMI_Message_Request[94] THEN HMI_MessageNo[0] := INT#94; END_IF;
(* Rung 102: 【Y1210】コンテナ仕分け送り 戻 異常表示 *)
IF HMI_Message_Request[95] THEN HMI_MessageNo[0] := INT#95; END_IF;
(* Rung 103: Output_Share_Error_M[12] 異常表示 *)
IF HMI_Message_Request[96] THEN HMI_MessageNo[0] := INT#96; END_IF;
(* Rung 104: 【Y1300】A(左側) コンベア受渡送り戻 異常表示 *)
IF HMI_Message_Request[97] THEN HMI_MessageNo[0] := INT#97; END_IF;

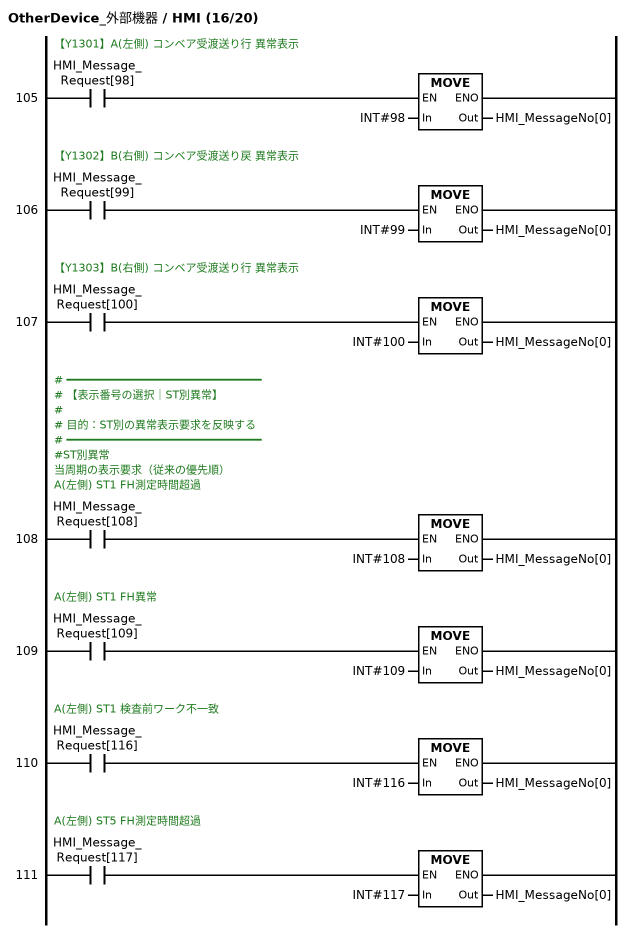
(* Rung 105: 【Y1301】A(左側) コンベア受渡送り行 異常表示 *)
IF HMI_Message_Request[98] THEN HMI_MessageNo[0] := INT#98; END_IF;
(* Rung 106: 【Y1302】B(右側) コンベア受渡送り戻 異常表示 *)
IF HMI_Message_Request[99] THEN HMI_MessageNo[0] := INT#99; END_IF;
(* Rung 107: 【Y1303】B(右側) コンベア受渡送り行 異常表示 *)
IF HMI_Message_Request[100] THEN HMI_MessageNo[0] := INT#100; END_IF;
(* Rung 108: # ━━━━━━━━━━━━━━━━━━━━━━━━━━━━━━ / # 【表示番号の選択｜ST別異常】 / # / # 目的：ST別の異常表示要求を反映する / # ━━━━━━━━━━━━━━━━━━━━━━━━━━━━━━ / #ST別異常 / 当周期の表示要求（従来の優先順） / A(左側) ST1 FH測定時間超過 *)
IF HMI_Message_Request[108] THEN HMI_MessageNo[0] := INT#108; END_IF;
(* Rung 109: A(左側) ST1 FH異常 *)
IF HMI_Message_Request[109] THEN HMI_MessageNo[0] := INT#109; END_IF;
(* Rung 110: A(左側) ST1 検査前ワーク不一致 *)
IF HMI_Message_Request[116] THEN HMI_MessageNo[0] := INT#116; END_IF;
(* Rung 111: A(左側) ST5 FH測定時間超過 *)
IF HMI_Message_Request[117] THEN HMI_MessageNo[0] := INT#117; END_IF;

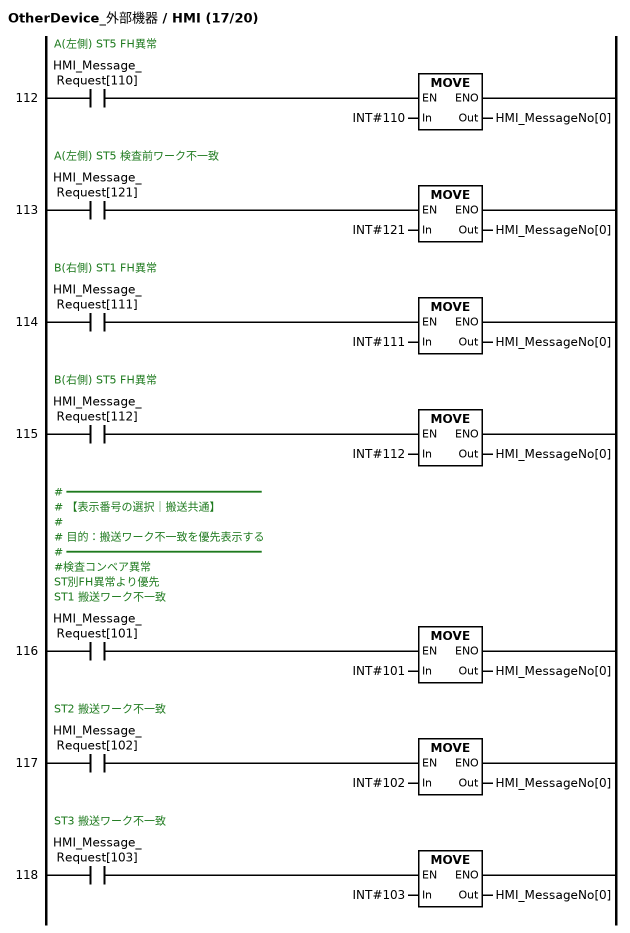
(* Rung 112: A(左側) ST5 FH異常 *)
IF HMI_Message_Request[110] THEN HMI_MessageNo[0] := INT#110; END_IF;
(* Rung 113: A(左側) ST5 検査前ワーク不一致 *)
IF HMI_Message_Request[121] THEN HMI_MessageNo[0] := INT#121; END_IF;
(* Rung 114: B(右側) ST1 FH異常 *)
IF HMI_Message_Request[111] THEN HMI_MessageNo[0] := INT#111; END_IF;
(* Rung 115: B(右側) ST5 FH異常 *)
IF HMI_Message_Request[112] THEN HMI_MessageNo[0] := INT#112; END_IF;
(* Rung 116: # ━━━━━━━━━━━━━━━━━━━━━━━━━━━━━━ / # 【表示番号の選択｜搬送共通】 / # / # 目的：搬送ワーク不一致を優先表示する / # ━━━━━━━━━━━━━━━━━━━━━━━━━━━━━━ / #検査コンベア異常 / ST別FH異常より優先 / ST1 搬送ワーク不一致 *)
IF HMI_Message_Request[101] THEN HMI_MessageNo[0] := INT#101; END_IF;
(* Rung 117: ST2 搬送ワーク不一致 *)
IF HMI_Message_Request[102] THEN HMI_MessageNo[0] := INT#102; END_IF;
(* Rung 118: ST3 搬送ワーク不一致 *)
IF HMI_Message_Request[103] THEN HMI_MessageNo[0] := INT#103; END_IF;

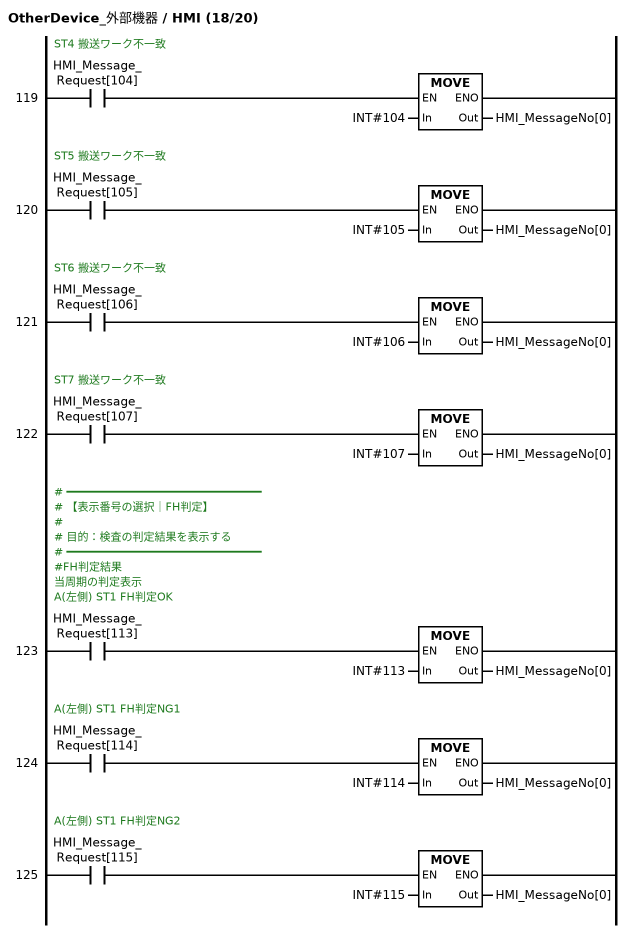
(* Rung 119: ST4 搬送ワーク不一致 *)
IF HMI_Message_Request[104] THEN HMI_MessageNo[0] := INT#104; END_IF;
(* Rung 120: ST5 搬送ワーク不一致 *)
IF HMI_Message_Request[105] THEN HMI_MessageNo[0] := INT#105; END_IF;
(* Rung 121: ST6 搬送ワーク不一致 *)
IF HMI_Message_Request[106] THEN HMI_MessageNo[0] := INT#106; END_IF;
(* Rung 122: ST7 搬送ワーク不一致 *)
IF HMI_Message_Request[107] THEN HMI_MessageNo[0] := INT#107; END_IF;
(* Rung 123: # ━━━━━━━━━━━━━━━━━━━━━━━━━━━━━━ / # 【表示番号の選択｜FH判定】 / # / # 目的：検査の判定結果を表示する / # ━━━━━━━━━━━━━━━━━━━━━━━━━━━━━━ / #FH判定結果 / 当周期の判定表示 / A(左側) ST1 FH判定OK *)
IF HMI_Message_Request[113] THEN HMI_MessageNo[0] := INT#113; END_IF;
(* Rung 124: A(左側) ST1 FH判定NG1 *)
IF HMI_Message_Request[114] THEN HMI_MessageNo[0] := INT#114; END_IF;
(* Rung 125: A(左側) ST1 FH判定NG2 *)
IF HMI_Message_Request[115] THEN HMI_MessageNo[0] := INT#115; END_IF;

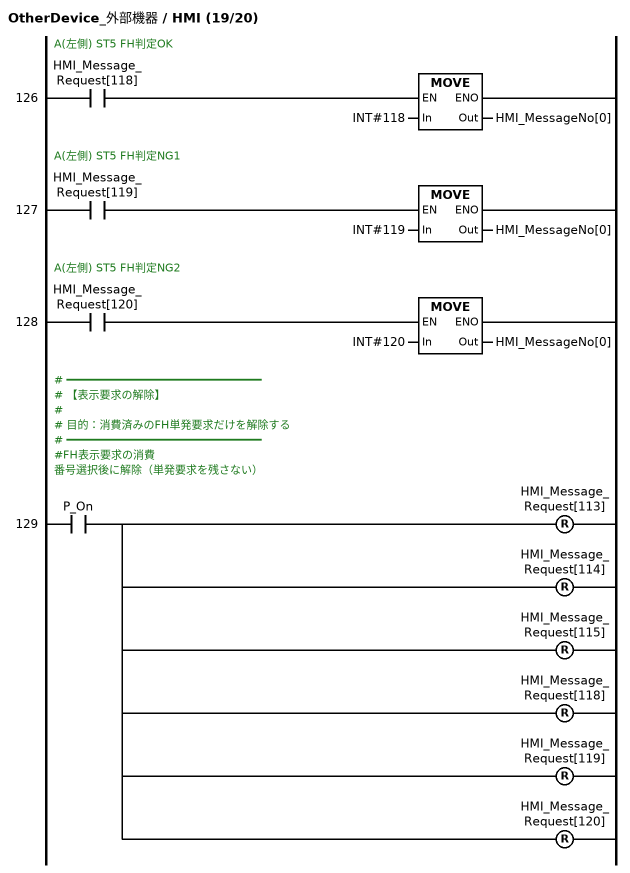
(* Rung 126: A(左側) ST5 FH判定OK *)
IF HMI_Message_Request[118] THEN HMI_MessageNo[0] := INT#118; END_IF;
(* Rung 127: A(左側) ST5 FH判定NG1 *)
IF HMI_Message_Request[119] THEN HMI_MessageNo[0] := INT#119; END_IF;
(* Rung 128: A(左側) ST5 FH判定NG2 *)
IF HMI_Message_Request[120] THEN HMI_MessageNo[0] := INT#120; END_IF;
(* Rung 129: # ━━━━━━━━━━━━━━━━━━━━━━━━━━━━━━ / # 【表示要求の解除】 / # / # 目的：消費済みのFH単発要求だけを解除する / # ━━━━━━━━━━━━━━━━━━━━━━━━━━━━━━ / #FH表示要求の消費 / 番号選択後に解除（単発要求を残さない） *)
IF P_On THEN
    HMI_Message_Request[113] := FALSE;
    HMI_Message_Request[114] := FALSE;
    HMI_Message_Request[115] := FALSE;
    HMI_Message_Request[118] := FALSE;
    HMI_Message_Request[119] := FALSE;
    HMI_Message_Request[120] := FALSE;
END_IF;

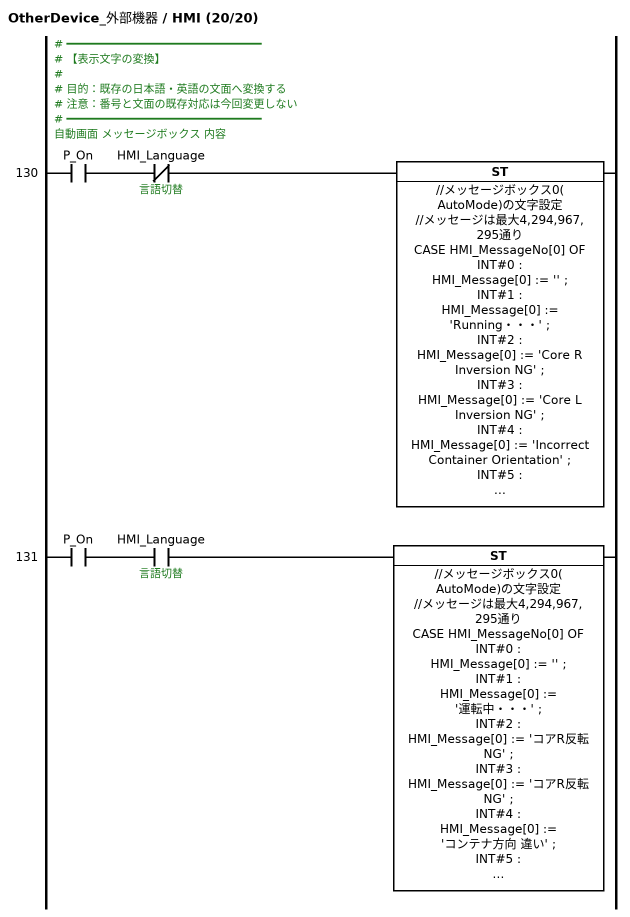
(* Rung 130: # ━━━━━━━━━━━━━━━━━━━━━━━━━━━━━━ / # 【表示文字の変換】 / # / # 目的：既存の日本語・英語の文面へ変換する / # 注意：番号と文面の既存対応は今回変更しない / # ━━━━━━━━━━━━━━━━━━━━━━━━━━━━━━ / 自動画面 メッセージボックス 内容 *)
IF P_On AND NOT HMI_Language THEN
    //メッセージボックス0(AutoMode)の文字設定
    //メッセージは最大4,294,967,295通り
    	
    	CASE HMI_MessageNo[0] OF
    	
    	INT#0 :
    	HMI_Message[0] := '' ;
        INT#1 :
    	HMI_Message[0] := 'Running・・・' ;
    	INT#2 :
    	HMI_Message[0] := 'Core R Inversion NG' ;
    	INT#3 :
    	HMI_Message[0] := 'Core L Inversion NG' ;
    	INT#4 :
    	HMI_Message[0] := 'Incorrect Container Orientation' ;
    	INT#5 :
    	HMI_Message[0] := 'Packed Container Full' ;
         INT#6 :
    	HMI_Message[0] := 'No Container Added' ;
    	INT#7 :
    	HMI_Message[0] := 'Paused・・・' ;
        INT#8 :
    	HMI_Message[0] := 'R Stock Holder Qty Error' ;
    	INT#9 :
    	HMI_Message[0] := 'L Stock Holder Qty Error' ;
        INT#10 :
    	HMI_Message[0] := 'Step Running・・・' ;
    	INT#11 :
    	HMI_Message[0] := 'Work Discharge Complete' ;
    	INT#12 :
    	HMI_Message[0] := 'SD Error' ;
    	END_CASE;		
    	
END_IF;
(* Rung 131 *)
IF P_On AND HMI_Language THEN
    //メッセージボックス0(AutoMode)の文字設定
    //メッセージは最大4,294,967,295通り
    	
    	CASE HMI_MessageNo[0] OF
    	
    	INT#0 :
    	HMI_Message[0] := '' ;
    	INT#1 :
    	HMI_Message[0] := '運転中・・・' ;	
    	INT#2 :
    	HMI_Message[0] := 'コアR反転 NG' ;	
        INT#3 :
    	HMI_Message[0] := 'コアR反転 NG' ;
    	INT#4 :
    	HMI_Message[0] := 'コンテナ方向 違い' ;
    	INT#5 :
    	HMI_Message[0] := '梱包済みコンテナ 満杯 or 排出詰まり' ;
        INT#6 :
    	HMI_Message[0] := 'コンテナ 無 追加してください' ;
        INT#7 :
    	HMI_Message[0] := '一時停止中・・・' ;
        INT#8 :
    	HMI_Message[0] := '右ストックフォルダ 入数ミス 取り除いて 再スタート' ;
        INT#9 :
    	HMI_Message[0] := '左ストックフォルダ 入数ミス 取り除いて 再スタート' ;
    	INT#10 :
    	HMI_Message[0] := 'ステップ運転中・・・' ;
    	INT#11 :
    	HMI_Message[0] := 'ワーク排出完了' ;
    	INT#12 :
    	HMI_Message[0] := 'SDカードエラー' ;
    	END_CASE;		
    	
END_IF;
END_PROGRAM

PROGRAM IO_入出力
VAR
    Timer_In_Sen_Accum_CV_A_Full : TON;
    Timer_In_Sen_Accum_CV_A_Arrival : TON;
    Timer_In_Sen_Work_A_Pos_00 : TON;
    Timer_In_Sen_Work_A_Pos_01 : TON;
    Timer_In_Sen_Work_A_Pos_02 : TON;
    Timer_In_Sen_Work_A_Pos_03 : TON;
    Timer_In_Sen_Work_A_Pos_04 : TON;
    Timer_In_Sen_Work_A_Pos_05 : TON;
    Timer_In_Sen_Work_A_Pos_06 : TON;
    Timer_In_Sen_Work_A_Pos_07 : TON;
    Timer_In_Sen_NG1_Tray_A_Full : TON;
    Timer_In_Sen_NG1_Tray_A_Full_Warn : TON;
    Timer_In_Sen_NG2_Tray_A_Full : TON;
    Timer_In_Sen_NG2_Tray_A_Full_Warn : TON;
    Timer_In_Sen_SH_A_Ent : TON;
    Timer_In_Sen_SH_A_Ext : TON;
    Timer_In_Sen_SH_A_Type_Ent : TON;
    Timer_In_Sen_SH_A_Type_Ext : TON;
    Timer_In_SenCY_Sply_Slide_A_H : TON;
    Timer_In_SenCY_Sply_Slide_A_F : TON;
    Timer_In_SenCY_Sply_Pick_A_H : TON;
    Timer_In_SenCY_Sply_Pick_A_F : TON;
    Timer_In_SenCY_Sply_Chk_A_H : TON;
    Timer_In_SenCY_Sply_Chk_A_F : TON;
    Timer_In_SenCY_HgtInsp_Clp_A_H : TON;
    Timer_In_SenCY_HgtInsp_Clp_A_F : TON;
    Timer_In_SenCY_HgtInsp_Lf_A_H : TON;
    Timer_In_SenCY_HgtInsp_Lf_A_F : TON;
    Timer_In_SenCY_NG1_Pick_A_H : TON;
    Timer_In_SenCY_NG1_Pick_A_F : TON;
    Timer_In_SenCY_NG1_Chk_A_H : TON;
    Timer_In_SenCY_NG1_Chk_A_F : TON;
    Timer_In_SenCY_Rev_01_Chk_A_H : TON;
    Timer_In_SenCY_Rev_01_Chk_A_F : TON;
    Timer_In_SenCY_Rev_01_Pick_A_H : TON;
    Timer_In_SenCY_Rev_01_Pick_A_F : TON;
    Timer_In_SenCY_Rev_02_Chk_A_H : TON;
    Timer_In_SenCY_Rev_02_Chk_A_F : TON;
    Timer_In_SenCY_Rev_02_Pick_A_H : TON;
    Timer_In_SenCY_Rev_02_Pick_A_F : TON;
    Timer_In_SenCY_Disc_Chk_A_H : TON;
    Timer_In_SenCY_Disc_Chk_A_F : TON;
    Timer_In_SenCY_Ejc_SH_Feed_A_F : TON;
    Timer_In_SenCY_Ejc_SH_Feed_A_H : TON;
    Timer_In_SenCY_Pos_01_Stopper_A_H : TON;
    Timer_In_SenCY_Pos_01_Stopper_A_F : TON;
    Timer_In_SenCY_Pos_02_Stopper_A_H : TON;
    Timer_In_SenCY_Pos_02_Stopper_A_F : TON;
    Timer_In_SenCY_Pos_03_Stopper_A_H : TON;
    Timer_In_SenCY_Pos_03_Stopper_A_F : TON;
    Timer_In_SenCY_Pos_04_Stopper_A_H : TON;
    Timer_In_SenCY_Pos_04_Stopper_A_F : TON;
    Timer_In_SenCY_Pos_05_Stopper_A_H : TON;
    Timer_In_SenCY_Pos_05_Stopper_A_F : TON;
    Timer_In_SenCY_Pos_06_Stopper_A_H : TON;
    Timer_In_SenCY_Pos_06_Stopper_A_F : TON;
    Timer_In_SenCY_SH_A_Turn_H : TON;
    Timer_In_SenCY_SH_A_Turn_F : TON;
    Timer_In_SenCY_NG1_Srt_A_H : TON;
    Timer_In_SenCY_NG1_Srt_A_F : TON;
    Timer_In_Sen_Accum_CV_B_Full : TON;
    Timer_In_Sen_Accum_CV_B_Arrival : TON;
    Timer_In_Sen_Work_B_Pos_00 : TON;
    Timer_In_Sen_Work_B_Pos_01 : TON;
    Timer_In_Sen_Work_B_Pos_02 : TON;
    Timer_In_Sen_Work_B_Pos_03 : TON;
    Timer_In_Sen_Work_B_Pos_04 : TON;
    Timer_In_Sen_Work_B_Pos_05 : TON;
    Timer_In_Sen_Work_B_Pos_06 : TON;
    Timer_In_Sen_Work_B_Pos_07 : TON;
    Timer_In_Sen_NG1_Tray_B_Full : TON;
    Timer_In_Sen_NG1_Tray_B_Full_Warn : TON;
    Timer_In_Sen_NG2_Tray_B_Full : TON;
    Timer_In_Sen_NG2_Tray_B_Full_Warn : TON;
    Timer_In_Sen_SH_B_Ent : TON;
    Timer_In_Sen_SH_B_Ext : TON;
    Timer_In_Sen_SH_B_Type_Ent : TON;
    Timer_In_Sen_SH_B_Type_Ext : TON;
    Timer_In_SenCY_Sply_Slide_B_H : TON;
    Timer_In_SenCY_Sply_Slide_B_F : TON;
    Timer_In_SenCY_Sply_Pick_B_H : TON;
    Timer_In_SenCY_Sply_Pick_B_F : TON;
    Timer_In_SenCY_Sply_Chk_B_H : TON;
    Timer_In_SenCY_HgtInsp_Clp_B_H : TON;
    Timer_In_SenCY_Sply_Chk_B_F : TON;
    Timer_In_SenCY_HgtInsp_Clp_B_F : TON;
    Timer_In_SenCY_HgtInsp_Lf_B_H : TON;
    Timer_In_SenCY_HgtInsp_Lf_B_F : TON;
    Timer_In_SenCY_NG1_Pick_B_H : TON;
    Timer_In_SenCY_NG1_Pick_B_F : TON;
    Timer_In_SenCY_NG1_Chk_B_H : TON;
    Timer_In_SenCY_NG1_Chk_B_F : TON;
    Timer_In_SenCY_Rev_01_Chk_B_H : TON;
    Timer_In_SenCY_Rev_01_Chk_B_F : TON;
    Timer_In_SenCY_Rev_01_Pick_B_H : TON;
    Timer_In_SenCY_Rev_01_Pick_B_F : TON;
    Timer_In_SenCY_Rev_02_Chk_B_H : TON;
    Timer_In_SenCY_Rev_02_Chk_B_F : TON;
    Timer_In_SenCY_Rev_02_Pick_B_H : TON;
    Timer_In_SenCY_Rev_02_Pick_B_F : TON;
    Timer_In_SenCY_Disc_Chk_B_H : TON;
    Timer_In_SenCY_Disc_Chk_B_F : TON;
    Timer_In_SenCY_Ejc_SH_Feed_B_F : TON;
    Timer_In_SenCY_Ejc_SH_Feed_B_H : TON;
    Timer_In_SenCY_Pos_01_Stopper_B_H : TON;
    Timer_In_SenCY_Pos_01_Stopper_B_F : TON;
    Timer_In_SenCY_Pos_02_Stopper_B_H : TON;
    Timer_In_SenCY_Pos_02_Stopper_B_F : TON;
    Timer_In_SenCY_Pos_03_Stopper_B_H : TON;
    Timer_In_SenCY_Pos_03_Stopper_B_F : TON;
    Timer_In_SenCY_Pos_04_Stopper_B_H : TON;
    Timer_In_SenCY_Pos_04_Stopper_B_F : TON;
    Timer_In_SenCY_Pos_05_Stopper_B_H : TON;
    Timer_In_SenCY_Pos_05_Stopper_B_F : TON;
    Timer_In_SenCY_Pos_06_Stopper_B_H : TON;
    Timer_In_SenCY_Pos_06_Stopper_B_F : TON;
    Timer_In_SenCY_SH_B_Turn_H : TON;
    Timer_In_SenCY_SH_B_Turn_F : TON;
    Timer_In_SenCY_NG1_Srt_B_H : TON;
    Timer_In_SenCY_NG1_Srt_B_F : TON;
    Timer_In_Sen_Supply_Container_Exist : TON;
    Timer_In_Sen_Destacker_Stage_01_Exist : TON;
    Timer_In_Sen_Destacker_Stage_02_Exist : TON;
    Timer_In_Sen_Container_Arrival : TON;
    Timer_In_Sen_Container_Direction_Check : TON;
    Timer_In_Sen_Container_Pass : TON;
    Timer_In_Sen_Container_Full : TON;
    Timer_In_Sen_Container_Sorting : TON;
    Timer_In_SenCY_Empty_Container_CY_H : TON;
    Timer_In_SenCY_Empty_Container_CY_F : TON;
    Timer_In_SenCY_Sep_Claw1_H : TON;
    Timer_In_SenCY_Sep_Claw1_F : TON;
    Timer_In_SenCY_Sep_Claw2_F : TON;
    Timer_In_SenCY_Sep_Claw2_H : TON;
    Timer_In_SenCY_Ejc_Cont1_H : TON;
    Timer_In_SenCY_Ejc_Cont1_F : TON;
    Timer_In_SenCY_Ejc_Cont2_H : TON;
    Timer_In_SenCY_Ejc_Cont2_F : TON;
    Timer_In_SenCY_Box_Chk_H : TON;
    Timer_In_SenCY_Box_Chk_F : TON;
    Timer_In_SenCY_Srt_Stopper_H : TON;
    Timer_In_SenCY_Srt_Stopper_F : TON;
    Timer_In_SenCY_Srt_Feed_H : TON;
    Timer_In_SenCY_Srt_Feed_F : TON;
    Timer_In_Sen_Unl_Conv_A_Pass : TON;
    Timer_In_Sen_Unl_Conv_B_Pass : TON;
    Timer_In_Sen_Trs_Conv_A_Arv : TON;
    Timer_In_Sen_Trs_Conv_A_Arrival : TON;
    Timer_In_Sen_Trs_Conv_B_Arrival : TON;
    Timer_In_SenCY_Hnd_Feed_A_H : TON;
    Timer_In_SenCY_Hnd_Feed_A_F : TON;
    Timer_In_SenCY_Hnd_Feed_B_H : TON;
    Timer_In_SenCY_Hnd_Feed_B_F : TON;
    Output_A_Error_TON : ARRAY[0..999] OF TON;  (* A(左側)出力タイムオーバーエラー： *)
    Output_A_M : ARRAY[0..999] OF Bool;  (* A(左側)出力補助コイル：; [1] 【Y616】A(左側) 供給スライド戻; [2] 【Y617】A(左側) 供給スライド行; [3] 【Y618】A(左側) 供給ピックアップ戻; [4] 【Y619】A(左側) 供給ピックアップ行; [5] 【Y620】A(左側) 供給チャック閉 戻; [6] 【Y621】A(左側) 供給チャック開 行; [7] 【Y700】A(左側) 高さ検査押え戻; [8] 【Y701】A(左側) 高さ検査押え行; [9] 【Y702】A(左側) 高さ検査持上戻; [10] 【Y703】A(左側) 高さ検査持上行; [11] 【Y704】A(左側) NG1ピックアップ戻; [12] 【Y705】A(左側) NG1ピックアップ 行; [13] 【Y706】A(左側) NG1チャック戻; [14] 【Y707】A(左側) NG1チャック行; [15] 【Y708】A(左側)ST4 反転1チャック閉; [16] 【Y709】A(左側)ST4 反転1チャック開; [17] 【Y710】A(左側)ST4 反転1ピックアップ戻; [18] 【Y711】A(左側)ST4 反転1ピックアップ行; [19] 【Y712】A(左側)ST6 反転2チャック閉 戻; [20] 【Y713】A(左側)ST6 反転2チャック開 行; [21] 【Y714】A(左側)ST6 反転2ピックアップ戻; [22] 【Y715】A(左側)ST6 反転2ピックアップ行; [23] 【Y716】A(左側) 排出チャック閉 戻; [24] 【Y717】A(左側) 排出チャック開 行; [25] 【Y718】A(左側) 排出フォルダ送り戻; [26] 【Y719】A(左側) 排出フォルダ送り行; [27] 【Y720】A(左側) 位置1ストッパー 戻; [28] 【Y720】A(左側) 位置1ストッパー 行; [29] 【Y721】A(左側) 位置2ストッパー; [30] 【Y721】A(左側) 位置2ストッパー; [32] 【Y722】A(左側) 位置3ストッパー行; [34] 【Y723】A(左側) 位置4ストッパー行; [35] 【Y724】A(左側) 位置5ストッパー戻; [36] 【Y724】A(左側) 位置5ストッパー行; [37] 【Y725】A(左側) 位置6ストッパー戻; [38] 【Y725】A(左側) 位置6ストッパー行; [39] 【Y726】A(左側) ストックフォルダターン戻; [40] 【Y727】A(左側) ストックフォルダターン行; [41] 【Y728】A(左側) NG1仕分け 戻; [42] 【Y729】A(左側) NG1仕分け 行; [43] 【Y1300】A(左側) コンベア受渡送り戻; [44] 【Y1301】A(左側) コンベア受渡送り行 *)
    Output_B_Error_TON : ARRAY[0..999] OF TON;  (* B(右側)出力タイムオーバーエラー *)
    Output_B_M : ARRAY[0..999] OF Bool;  (* B(右側)出力補助コイル：; [1] 【Y622】B(右側) 供給スライド戻; [2] 【Y623】B(右側) 供給スライド行; [3] 【Y624】B(右側) 供給ピックアップ戻; [4] 【Y625】B(右側) 供給ピックアップ行; [5] 【Y626】B(右側) 供給チャック閉 戻; [6] 【Y627】B(右側) 供給チャック開 行; [7] 【Y800】B(右側) 高さ検査押え戻; [9] 【Y802】B(右側) 高さ検査持上戻; [11] 【Y804】B(右側) NG1ピックアップ戻; [14] 【Y807】B(右側) NG1チャック行; [18] 【Y811】B(右側)ST4 反転1ピックアップ行; [42] 【Y829】B(右側) NG1仕分け 行; [41] 【Y828】B(右側) NG1仕分け 戻; [40] 【Y827】B(右側) ストックフォルダターン行; [39] 【Y826】B(右側) ストックフォルダターン戻; [38] 【Y825】B(右側) 位置6ストッパー行; [37] 【Y825】B(右側) 位置6ストッパー戻; [36] 【Y824】B(右側) 位置5ストッパー行; [35] 【Y824】B(右側) 位置5ストッパー戻; [34] 【Y823】B(右側) 位置4ストッパー行; [33] 【Y823】B(右側) 位置4ストッパー戻; [32] 【Y822】B(右側) 位置3ストッパー行; [31] 【Y822】B(右側) 位置3ストッパー戻; [30] 【Y821】B(右側) 位置2ストッパー行; [29] 【Y821】B(右側) 位置2ストッパー戻; [28] 【Y820】B(右側) 位置1ストッパー 行; [27] 【Y820】B(右側) 位置1ストッパー 戻; [26] 【Y819】B(右側) 排出フォルダ送り行; [25] 【Y818】B(右側) 排出フォルダ送り戻; [24] 【Y817】B(右側) 排出チャック開 行; [23] 【Y816】B(右側) 排出チャック閉 戻; [22] 【Y815】B(右側)ST6 反転2ピックアップ行; [21] 【Y814】B(右側)ST6 反転2ピックアップ戻; [20] 【Y813】B(右側)ST6 反転2チャック開 行; [19] 【Y812】B(右側)ST6 反転2チャック閉 戻; [17] 【Y810】B(右側)ST4 反転1ピックアップ戻; [16] 【Y809】B(右側)ST4 反転1チャック開 戻; [15] 【Y808】B(右側)ST4 反転1チャック閉 戻; [13] 【Y806】B(右側) NG1チャック戻; [12] 【Y805】B(右側) NG1ピックアップ 行; [10] 【Y803】B(右側) 高さ検査持上行; [8] 【Y801】B(右側) 高さ検査押え行; [43] 【Y1302】B(右側) コンベア受渡送り戻; [44] 【Y1303】B(右側) コンベア受渡送り行 *)
    Mtr_Flip_02_Busy : BOOL;  (* A(左側)反転 オリエンタルモータ2 動作中 *)
    Output_A_Reset_TON : ARRAY[0..99] OF TON;  (* A(左側)出力リセット ：; [34] 【Y723】A(左側) 位置4ストッパー行 *)
    Output_B_Reset_TON : ARRAY[0..99] OF TON;  (* B(右側)出力リセット ： *)
    Output_Share_M : ARRAY[0..99] OF Bool;  (* 共有出力補助コイル：; [1] 【Y1200】空コンテナ送り 戻; [2] 【Y1201】空コンテナ送り 行; [3] 【Y1202】段バラシ爪 戻; [4] 【Y1203】段バラシ爪 行; [5] 【Y1204】コンテナ排出 戻; [6] 【Y1205】コンテナ排出 行; [7] 【Y1206】箱入れチャック 戻; [8] 【Y1207】箱入れチャック 行; [9] 【Y1208】コンテナ仕分けストッパー 戻; [10] 【Y1209】コンテナ仕分けストッパー 行; [11] 【Y1210】コンテナ仕分け送り 戻 *)
    Output_Share_Reset_TON : ARRAY[0..99] OF TON;  (* 共有出力リセット:; [7] 【Y1206】箱入れチャック 戻 *)
    Output_Share_Error_TON : ARRAY[0..99] OF TON;  (* 共有出力タイムオーバーエラー *)
    IAI_In_Sample_Busy_MOVE : BOOL;
    Input_T : ARRAY[0..99] OF TON;
    Timer_In_Sen_Tray_Direction_Check : TON;
END_VAR
VAR_EXTERNAL
    In_Sw_EMS1 : BOOL;
    In_Sen_Accum_CV_A_Full : BOOL;
    TimerQ_In_Sen_Accum_CV_A_Full : BOOL;  (* 【X200】A(左側) アキュームCV満 *)
    In_Sen_Accum_CV_A_Arrival : BOOL;
    TimerQ_In_Sen_Accum_CV_A_Arrival : BOOL;  (* 【X201】A(左側) アキュームCV着 *)
    In_Sen_Work_A_Pos_00 : BOOL;
    TimerQ_In_Sen_Work_A_Pos_00 : BOOL;  (* 【X202】A(左側)ワーク位置0 *)
    In_Sen_Work_A_Pos_01 : BOOL;
    TimerQ_In_Sen_Work_A_Pos_01 : BOOL;  (* 【X203】A(左側)ワーク位置1 *)
    In_Sen_Work_A_Pos_02 : BOOL;
    TimerQ_In_Sen_Work_A_Pos_02 : BOOL;  (* 【X204】A(左側)ワーク位置2 *)
    In_Sen_Work_A_Pos_03 : BOOL;
    TimerQ_In_Sen_Work_A_Pos_03 : BOOL;  (* 【X205】A(左側)ワーク位置3 *)
    In_Sen_Work_A_Pos_04 : BOOL;
    TimerQ_In_Sen_Work_A_Pos_04 : BOOL;  (* 【X206】A(左側)ワーク位置4 *)
    In_Sen_Work_A_Pos_05 : BOOL;
    TimerQ_In_Sen_Work_A_Pos_05 : BOOL;  (* 【X207】A(左側)ワーク位置5 *)
    In_Sen_Work_A_Pos_06 : BOOL;
    TimerQ_In_Sen_Work_A_Pos_06 : BOOL;  (* 【X208】A(左側)ワーク位置6 *)
    In_Sen_Work_A_Pos_07 : BOOL;
    TimerQ_In_Sen_Work_A_Pos_07 : BOOL;  (* 【X209】A(左側)ワーク位置7 *)
    In_Sen_NG1_Tray_A_Full : BOOL;
    TimerQ_In_Sen_NG1_Tray_A_Full : BOOL;  (* 【X210】A(左側) NG1トレイ満杯停止 *)
    In_Sen_NG1_Tray_A_Full_Warn : BOOL;
    TimerQ_In_Sen_NG1_Tray_A_Full_Warn : BOOL;  (* 【X211】A(左側) NG1トレイ満杯警告 *)
    In_Sen_NG2_Tray_A_Full : BOOL;
    TimerQ_In_Sen_NG2_Tray_A_Full : BOOL;  (* 【X212】A(左側) NG2トレイ満杯停止 *)
    In_Sen_NG2_Tray_A_Full_Warn : BOOL;
    TimerQ_In_Sen_NG2_Tray_A_Full_Warn : BOOL;  (* 【X213】A(左側) NG2トレイ満杯警告 *)
    In_Sen_SH_A_Ent : BOOL;
    TimerQ_In_Sen_SH_A_Ent : BOOL;  (* 【X214】A(左側) ストックフォルダIN *)
    In_Sen_SH_A_Ext : BOOL;
    TimerQ_In_Sen_SH_A_Ext : BOOL;  (* 【X215】A(左側) ストックフォルダOut *)
    In_Sen_SH_A_Type_Ent : BOOL;
    TimerQ_In_Sen_SH_A_Type_Ent : BOOL;  (* 【X216】A(左側) ストック機種判別IN *)
    In_Sen_SH_A_Type_Ext : BOOL;
    TimerQ_In_Sen_SH_A_Type_Ext : BOOL;  (* 【X217】A(左側) ストック機種判別OUT *)
    In_SenCY_Sply_Slide_A_H : BOOL;
    In_SenCY_Sply_Slide_A_F : BOOL;
    TimerQ_In_SenCY_Sply_Slide_A_H : BOOL;  (* 【X218】A(左側) 供給スライド戻 *)
    TimerQ_In_SenCY_Sply_Slide_A_F : BOOL;  (* 【X219】A(左側) 供給スライド行 *)
    In_SenCY_Sply_Pick_A_H : BOOL;
    TimerQ_In_SenCY_Sply_Pick_A_H : BOOL;  (* 【X220】A(左側) 供給ピックアップ戻 *)
    In_SenCY_Sply_Pick_A_F : BOOL;
    TimerQ_In_SenCY_Sply_Pick_A_F : BOOL;  (* 【X221】A(左側) 供給ピックアップ行 *)
    In_SenCY_Sply_Chk_A_H : BOOL;
    TimerQ_In_SenCY_Sply_Chk_A_H : BOOL;  (* 【X222】A(左側) 供給チャック戻 *)
    In_SenCY_Sply_Chk_A_F : BOOL;
    TimerQ_In_SenCY_Sply_Chk_A_F : BOOL;  (* 【X223】A(左側) 供給チャック行 *)
    In_SenCY_HgtInsp_Clp_A_H : BOOL;
    TimerQ_In_SenCY_HgtInsp_Clp_A_H : BOOL;  (* 【X224】A(左側) 高さ検査押え戻 *)
    In_SenCY_HgtInsp_Clp_A_F : BOOL;
    TimerQ_In_SenCY_HgtInsp_Clp_A_F : BOOL;  (* 【X225】A(左側) 高さ検査押え行 *)
    In_SenCY_HgtInsp_Lf_A_H : BOOL;
    TimerQ_In_SenCY_HgtInsp_Lf_A_H : BOOL;  (* 【X226】A(左側) 高さ検査持上戻 *)
    In_SenCY_HgtInsp_Lf_A_F : BOOL;
    TimerQ_In_SenCY_HgtInsp_Lf_A_F : BOOL;  (* 【X227】A(左側) 高さ検査持上行 *)
    In_SenCY_NG1_Pick_A_H : BOOL;
    In_SenCY_NG1_Pick_A_F : BOOL;
    In_SenCY_NG1_Chk_A_H : BOOL;
    TimerQ_In_SenCY_NG1_Pick_A_H : BOOL;  (* 【X228】A(左側) NG1ピックアップ戻 *)
    TimerQ_In_SenCY_NG1_Pick_A_F : BOOL;  (* 【X229】A(左側) NG1ピックアップ行 *)
    TimerQ_In_SenCY_NG1_Chk_A_H : BOOL;  (* 【X230】A(左側) NG1チャック戻 *)
    In_SenCY_NG1_Chk_A_F : BOOL;
    In_SenCY_Rev_01_Chk_A_H : BOOL;  (* 【X300】A(左側)ST4 反転1チャック戻 *)
    In_SenCY_Rev_01_Chk_A_F : BOOL;  (* 【X301】A(左側)ST4 反転1チャック行 *)
    In_SenCY_Rev_01_Pick_A_H : BOOL;  (* 【X302】A(左側)ST4 反転1ピックアップ戻 *)
    In_SenCY_Rev_01_Pick_A_F : BOOL;  (* 【X303】A(左側)ST4 反転1ピックアップ行 *)
    In_SenCY_Rev_02_Chk_A_H : BOOL;  (* 【X304】A(左側)ST6 反転2チャック戻 *)
    In_SenCY_Rev_02_Chk_A_F : BOOL;  (* 【X305】A(左側)ST6 反転2チャック行 *)
    In_SenCY_Rev_02_Pick_A_H : BOOL;  (* 【X306】A(左側)ST6 反転2ピックアップ戻 *)
    TimerQ_In_SenCY_NG1_Chk_A_F : BOOL;  (* 【X231】A(左側) NG1チャック行 *)
    TimerQ_In_SenCY_Rev_01_Chk_A_H : BOOL;  (* 【X300】A(左側)ST4 反転1チャック戻 *)
    TimerQ_In_SenCY_Rev_01_Chk_A_F : BOOL;  (* 【X301】A(左側)ST4 反転1チャック行 *)
    TimerQ_In_SenCY_Rev_01_Pick_A_H : BOOL;  (* 【X302】A(左側)ST4 反転1ピックアップ戻 *)
    TimerQ_In_SenCY_Rev_01_Pick_A_F : BOOL;  (* 【X303】A(左側)ST4 反転1ピックアップ行 *)
    TimerQ_In_SenCY_Rev_02_Chk_A_H : BOOL;  (* 【X304】A(左側)ST6 反転2チャック戻 *)
    TimerQ_In_SenCY_Rev_02_Chk_A_F : BOOL;  (* 【X305】A(左側)ST6 反転2チャック行 *)
    TimerQ_In_SenCY_Rev_02_Pick_A_H : BOOL;  (* 【X306】A(左側)ST6 反転2ピックアップ戻 *)
    In_SenCY_Rev_02_Pick_A_F : BOOL;  (* 【X307】A(左側)ST6 反転2ピックアップ行 *)
    TimerQ_In_SenCY_Rev_02_Pick_A_F : BOOL;  (* 【X307】A(左側)ST6 反転2ピックアップ行 *)
    In_SenCY_Disc_Chk_A_H : BOOL;
    TimerQ_In_SenCY_Disc_Chk_A_H : BOOL;  (* 【X308】A(左側) 排出チャック戻 *)
    In_SenCY_Disc_Chk_A_F : BOOL;
    TimerQ_In_SenCY_Disc_Chk_A_F : BOOL;  (* 【X309】A(左側) 排出チャック行 *)
    In_SenCY_Ejc_SH_Feed_A_H : BOOL;
    In_SenCY_Ejc_SH_Feed_A_F : BOOL;
    TimerQ_In_SenCY_Ejc_SH_Feed_A_H : BOOL;  (* 【X310】A(左側) 排出フォルダ送り戻 *)
    TimerQ_In_SenCY_Ejc_SH_Feed_A_F : BOOL;  (* 【X311】A(左側) 排出フォルダ送り行 *)
    In_SenCY_Pos_01_Stopper_A_H : BOOL;
    TimerQ_In_SenCY_Pos_01_Stopper_A_H : BOOL;  (* 【X312】A(左側) 位置1ストッパー戻 *)
    In_SenCY_Pos_01_Stopper_A_F : BOOL;
    TimerQ_In_SenCY_Pos_01_Stopper_A_F : BOOL;  (* 【X313】位置1ストッパー行 *)
    In_SenCY_Pos_02_Stopper_A_H : BOOL;
    TimerQ_In_SenCY_Pos_02_Stopper_A_H : BOOL;  (* 【X314】A(左側) 位置2ストッパー戻 *)
    In_SenCY_Pos_02_Stopper_A_F : BOOL;
    TimerQ_In_SenCY_Pos_02_Stopper_A_F : BOOL;  (* 【X315】A(左側) 位置2ストッパー行 *)
    In_SenCY_Pos_03_Stopper_A_H : BOOL;
    In_SenCY_Pos_03_Stopper_A_F : BOOL;
    TimerQ_In_SenCY_Pos_03_Stopper_A_H : BOOL;  (* 【X316】A(左側) 位置3ストッパー戻 *)
    TimerQ_In_SenCY_Pos_03_Stopper_A_F : BOOL;  (* 【X317】A(左側) 位置3ストッパー行 *)
    In_SenCY_Pos_04_Stopper_A_H : BOOL;
    In_SenCY_Pos_04_Stopper_A_F : BOOL;
    TimerQ_In_SenCY_Pos_04_Stopper_A_H : BOOL;  (* 【X318】A(左側) 位置4ストッパー戻 *)
    TimerQ_In_SenCY_Pos_04_Stopper_A_F : BOOL;  (* 【X319】A(左側) 位置4ストッパー行 *)
    In_SenCY_Pos_05_Stopper_A_H : BOOL;
    In_SenCY_Pos_05_Stopper_A_F : BOOL;
    TimerQ_In_SenCY_Pos_05_Stopper_A_H : BOOL;  (* 【X320】A(左側) 位置5ストッパー戻 *)
    TimerQ_In_SenCY_Pos_05_Stopper_A_F : BOOL;  (* 【X321】A(左側) 位置5ストッパー行 *)
    In_SenCY_Pos_06_Stopper_A_H : BOOL;
    In_SenCY_Pos_06_Stopper_A_F : BOOL;
    TimerQ_In_SenCY_Pos_06_Stopper_A_H : BOOL;  (* 【X322】A(左側) 位置6ストッパー戻 *)
    TimerQ_In_SenCY_Pos_06_Stopper_A_F : BOOL;  (* 【X323】A(左側) 位置6ストッパー行 *)
    In_SenCY_SH_A_Turn_H : BOOL;
    TimerQ_In_SenCY_SH_A_Turn_H : BOOL;  (* 【X324】A(左側) ストックフォルダターン戻 *)
    In_SenCY_SH_A_Turn_F : BOOL;
    TimerQ_In_SenCY_SH_A_Turn_F : BOOL;  (* 【X325】A(左側) ストックフォルダターン行 *)
    In_SenCY_NG1_Srt_A_H : BOOL;
    TimerQ_In_SenCY_NG1_Srt_A_H : BOOL;  (* 【X330】NG1仕分け 戻 *)
    In_SenCY_NG1_Srt_A_F : BOOL;
    TimerQ_In_SenCY_NG1_Srt_A_F : BOOL;  (* 【X331】NG1仕分け 行 *)
    TimerQ_In_Sen_Accum_CV_B_Full : BOOL;  (* 【X400】B(右側) アキュームCV満 *)
    In_Sen_Accum_CV_B_Arrival : BOOL;
    TimerQ_In_Sen_Accum_CV_B_Arrival : BOOL;  (* 【X401】B(右側) アキュームCV着 *)
    In_Sen_Work_B_Pos_00 : BOOL;
    TimerQ_In_Sen_Work_B_Pos_00 : BOOL;  (* 【X402】B(右側)ワーク位置0 *)
    In_Sen_Work_B_Pos_01 : BOOL;
    In_Sen_Work_B_Pos_02 : BOOL;
    In_Sen_Work_B_Pos_03 : BOOL;
    In_Sen_Work_B_Pos_04 : BOOL;
    In_Sen_Work_B_Pos_05 : BOOL;
    In_Sen_Work_B_Pos_06 : BOOL;
    In_Sen_Work_B_Pos_07 : BOOL;
    In_Sen_NG1_Tray_B_Full : BOOL;
    In_Sen_NG1_Tray_B_Full_Warn : BOOL;
    In_Sen_NG2_Tray_B_Full : BOOL;
    In_Sen_NG2_Tray_B_Full_Warn : BOOL;
    In_Sen_SH_B_Ent : BOOL;
    In_Sen_SH_B_Ext : BOOL;
    In_Sen_SH_B_Type_Ent : BOOL;
    In_Sen_SH_B_Type_Ext : BOOL;
    In_SenCY_Sply_Slide_B_H : BOOL;
    In_SenCY_Sply_Slide_B_F : BOOL;
    In_SenCY_Sply_Pick_B_H : BOOL;
    In_SenCY_Sply_Pick_B_F : BOOL;
    In_SenCY_Sply_Chk_B_H : BOOL;
    In_SenCY_HgtInsp_Clp_B_H : BOOL;
    In_SenCY_Sply_Chk_B_F : BOOL;
    In_SenCY_HgtInsp_Clp_B_F : BOOL;
    In_SenCY_HgtInsp_Lf_B_H : BOOL;
    In_SenCY_HgtInsp_Lf_B_F : BOOL;
    In_SenCY_NG1_Pick_B_H : BOOL;
    In_SenCY_NG1_Pick_B_F : BOOL;
    In_SenCY_NG1_Chk_B_H : BOOL;
    In_SenCY_NG1_Chk_B_F : BOOL;
    In_SenCY_Rev_01_Chk_B_H : BOOL;  (* 【X500】B(右側)ST4 反転1チャック閉 戻 *)
    In_SenCY_Rev_01_Chk_B_F : BOOL;  (* 【X501】B(右側)ST4 反転1チャック開 行 *)
    In_SenCY_Rev_01_Pick_B_H : BOOL;  (* 【X502】B(右側)ST4 反転1ピックアップ戻 *)
    In_SenCY_Rev_01_Pick_B_F : BOOL;  (* 【X503】B(右側)ST4 反転1ピックアップ行 *)
    In_SenCY_Rev_02_Chk_B_H : BOOL;  (* 【X504】B(右側)ST6 反転2チャック閉 戻 *)
    In_SenCY_Rev_02_Chk_B_F : BOOL;  (* 【X505】B(右側)ST6 反転2チャック開 行 *)
    In_SenCY_Rev_02_Pick_B_H : BOOL;  (* 【X506】B(右側)ST6 反転2ピックアップ戻 *)
    In_SenCY_Rev_02_Pick_B_F : BOOL;  (* 【X507】B(右側)ST6 反転2ピックアップ行 *)
    In_SenCY_Disc_Chk_B_H : BOOL;
    In_SenCY_Disc_Chk_B_F : BOOL;
    In_SenCY_Ejc_SH_Feed_B_H : BOOL;
    In_SenCY_Ejc_SH_Feed_B_F : BOOL;
    In_SenCY_Pos_01_Stopper_B_H : BOOL;
    In_SenCY_Pos_01_Stopper_B_F : BOOL;
    In_SenCY_Pos_02_Stopper_B_H : BOOL;
    In_SenCY_Pos_02_Stopper_B_F : BOOL;
    In_SenCY_Pos_03_Stopper_B_H : BOOL;
    In_SenCY_Pos_03_Stopper_B_F : BOOL;
    In_SenCY_Pos_04_Stopper_B_H : BOOL;
    In_SenCY_Pos_04_Stopper_B_F : BOOL;
    In_SenCY_Pos_05_Stopper_B_H : BOOL;
    In_SenCY_Pos_05_Stopper_B_F : BOOL;
    In_SenCY_Pos_06_Stopper_B_H : BOOL;
    In_SenCY_Pos_06_Stopper_B_F : BOOL;
    In_SenCY_SH_B_Turn_H : BOOL;
    In_SenCY_SH_B_Turn_F : BOOL;
    In_SenCY_NG1_Srt_B_H : BOOL;
    In_SenCY_NG1_Srt_B_F : BOOL;
    TimerQ_In_Sen_Work_B_Pos_01 : BOOL;  (* 【X403】B(右側)ワーク位置1 *)
    TimerQ_In_Sen_Work_B_Pos_02 : BOOL;  (* 【X404】B(右側)ワーク位置2 *)
    TimerQ_In_Sen_Work_B_Pos_03 : BOOL;  (* 【X405】B(右側)ワーク位置3 *)
    TimerQ_In_Sen_Work_B_Pos_04 : BOOL;  (* 【X406】B(右側)ワーク位置4 *)
    TimerQ_In_Sen_Work_B_Pos_05 : BOOL;  (* 【X407】B(右側)ワーク位置5 *)
    TimerQ_In_Sen_Work_B_Pos_06 : BOOL;  (* 【X408】B(右側)ワーク位置6 *)
    TimerQ_In_Sen_Work_B_Pos_07 : BOOL;  (* 【X409】B(右側)ワーク位置7 *)
    TimerQ_In_Sen_NG1_Tray_B_Full : BOOL;  (* 【X410】B(右側) NG1トレイ満杯停止 *)
    TimerQ_In_Sen_NG1_Tray_B_Full_Warn : BOOL;  (* 【X411】B(右側) NG1トレイ満杯警告 *)
    TimerQ_In_Sen_NG2_Tray_B_Full : BOOL;  (* 【X412】B(右側) NG2トレイ満杯停止 *)
    TimerQ_In_Sen_NG2_Tray_B_Full_Warn : BOOL;  (* 【X413】B(右側) NG2トレイ満杯警告 *)
    TimerQ_In_Sen_SH_B_Ent : BOOL;  (* 【X414】B(右側) ストックフォルダIN *)
    TimerQ_In_Sen_SH_B_Ext : BOOL;  (* 【X415】B(右側) ストックフォルダOut *)
    TimerQ_In_Sen_SH_B_Type_Ent : BOOL;  (* 【X416】B(右側) ストック機種判別IN *)
    TimerQ_In_Sen_SH_B_Type_Ext : BOOL;  (* 【X417】B(右側) ストック機種判別OUT *)
    TimerQ_In_SenCY_Sply_Slide_B_H : BOOL;  (* 【X418】B(右側) 供給スライド戻 *)
    TimerQ_In_SenCY_Sply_Slide_B_F : BOOL;  (* 【X419】B(右側) 供給スライド行 *)
    TimerQ_In_SenCY_Sply_Pick_B_H : BOOL;  (* 【X420】B(右側) 供給ピックアップ戻 *)
    TimerQ_In_SenCY_Sply_Pick_B_F : BOOL;  (* 【X421】B(右側) 供給ピックアップ行 *)
    TimerQ_In_SenCY_Sply_Chk_B_H : BOOL;  (* 【X422】B(右側) 供給チャック閉 戻 *)
    TimerQ_In_SenCY_HgtInsp_Clp_B_H : BOOL;  (* 【X424】B(右側) 高さ検査押え戻 *)
    TimerQ_In_SenCY_Sply_Chk_B_F : BOOL;  (* 【X423】B(右側) 供給チャック開 行 *)
    TimerQ_In_SenCY_HgtInsp_Clp_B_F : BOOL;  (* 【X425】B(右側) 高さ検査押え行 *)
    TimerQ_In_SenCY_HgtInsp_Lf_B_H : BOOL;  (* 【X426】B(右側) 高さ検査持上戻 *)
    TimerQ_In_SenCY_HgtInsp_Lf_B_F : BOOL;  (* 【X427】 B(右側) 高さ検査持上行 *)
    TimerQ_In_SenCY_NG1_Pick_B_H : BOOL;  (* 【X428】B(右側) NG1ピックアップ戻 *)
    TimerQ_In_SenCY_NG1_Pick_B_F : BOOL;  (* 【X429】B(右側) NG1ピックアップ行 *)
    TimerQ_In_SenCY_NG1_Chk_B_H : BOOL;  (* 【X430】 B(右側) NG1チャック閉 戻 *)
    TimerQ_In_SenCY_NG1_Chk_B_F : BOOL;  (* 【X431】B(右側) NG1チャック開 行 *)
    TimerQ_In_SenCY_Rev_01_Chk_B_H : BOOL;  (* 【X500】B(右側)ST4 反転1チャック閉 戻 *)
    TimerQ_In_SenCY_Rev_01_Pick_B_H : BOOL;  (* 【X502】B(右側)ST4 反転1ピックアップ戻 *)
    TimerQ_In_SenCY_Rev_01_Pick_B_F : BOOL;  (* 【X503】B(右側)ST4 反転1ピックアップ行 *)
    TimerQ_In_SenCY_Rev_02_Chk_B_H : BOOL;  (* 【X504】B(右側)ST6 反転2チャック閉 戻 *)
    TimerQ_In_SenCY_Rev_02_Chk_B_F : BOOL;  (* 【X505】B(右側)ST6 反転2チャック開 行 *)
    TimerQ_In_SenCY_Rev_02_Pick_B_H : BOOL;  (* 【X506】B(右側)ST6 反転2ピックアップ戻 *)
    TimerQ_In_SenCY_Rev_02_Pick_B_F : BOOL;  (* 【X507】B(右側)ST6 反転2ピックアップ行 *)
    TimerQ_In_SenCY_Disc_Chk_B_H : BOOL;  (* 【X508】B(右側) 排出チャック閉 戻 *)
    TimerQ_In_SenCY_Disc_Chk_B_F : BOOL;  (* 【X509】B(右側) 排出チャック開 行 *)
    TimerQ_In_SenCY_Ejc_SH_Feed_B_H : BOOL;  (* 【X511】B(右側) 排出フォルダ送り行 *)
    TimerQ_In_SenCY_Ejc_SH_Feed_B_F : BOOL;  (* 【X510】B(右側) 排出フォルダ送り戻 *)
    TimerQ_In_SenCY_Pos_01_Stopper_B_H : BOOL;  (* 【X512】B(右側) 位置1ストッパー戻 *)
    TimerQ_In_SenCY_Pos_01_Stopper_B_F : BOOL;  (* 【X513】B(右側) 位置1ストッパー行 *)
    TimerQ_In_SenCY_Pos_02_Stopper_B_H : BOOL;  (* 【X514】B(右側) 位置2ストッパー戻 *)
    TimerQ_In_SenCY_Pos_02_Stopper_B_F : BOOL;  (* 【X515】B(右側) 位置2ストッパー行 *)
    TimerQ_In_SenCY_Pos_03_Stopper_B_H : BOOL;  (* 【X516】B(右側) 位置3ストッパー戻 *)
    TimerQ_In_SenCY_Pos_03_Stopper_B_F : BOOL;  (* 【X517】B(右側) 位置3ストッパー行 *)
    TimerQ_In_SenCY_Pos_04_Stopper_B_H : BOOL;  (* 【X518】B(右側) 位置4ストッパー戻 *)
    TimerQ_In_SenCY_Pos_04_Stopper_B_F : BOOL;  (* 【X519】B(右側) 位置4ストッパー行 *)
    TimerQ_In_SenCY_Pos_05_Stopper_B_H : BOOL;  (* 【X520】B(右側) 位置5ストッパー戻 *)
    TimerQ_In_SenCY_Pos_05_Stopper_B_F : BOOL;  (* 【X521】B(右側) 位置5ストッパー行 *)
    TimerQ_In_SenCY_Pos_06_Stopper_B_H : BOOL;  (* 【X522】B(右側) 位置6ストッパー戻 *)
    TimerQ_In_SenCY_Pos_06_Stopper_B_F : BOOL;  (* 【X523】B(右側) 位置6ストッパー行 *)
    TimerQ_In_SenCY_SH_B_Turn_H : BOOL;  (* 【X524】B(右側) ストックフォルダターン戻 *)
    TimerQ_In_SenCY_SH_B_Turn_F : BOOL;  (* 【X525】B(右側) ストックフォルダターン行 *)
    TimerQ_In_SenCY_NG1_Srt_B_H : BOOL;  (* 【X530】B(右側) NG1仕分け 戻 *)
    TimerQ_In_SenCY_NG1_Srt_B_F : BOOL;  (* 【X531】B(右側) NG1仕分け 行 *)
    In_Sen_Supply_Container_Exist : BOOL;
    In_Sen_Destacker_Stage_01_Exist : BOOL;
    In_Sen_Destacker_Stage_02_Exist : BOOL;
    In_Sen_Container_Arrival : BOOL;
    In_Sen_Container_Direction_Check : BOOL;
    In_Sen_Container_Pass : BOOL;
    In_Sen_Container_Full : BOOL;
    In_SenCY_Empty_Container_CY_H : BOOL;
    In_SenCY_Empty_Container_CY_F : BOOL;
    In_SenCY_Sep_Claw1_H : BOOL;
    In_SenCY_Sep_Claw1_F : BOOL;
    In_SenCY_Sep_Claw2_F : BOOL;
    In_SenCY_Sep_Claw2_H : BOOL;
    In_SenCY_Ejc_Cont1_H : BOOL;
    In_SenCY_Ejc_Cont1_F : BOOL;
    In_SenCY_Ejc_Cont2_F : BOOL;
    In_SenCY_Ejc_Cont2_H : BOOL;
    In_SenCY_Box_Chk_H : BOOL;
    In_SenCY_Box_Chk_F : BOOL;
    In_SenCY_Srt_Stopper_H : BOOL;
    In_SenCY_Srt_Stopper_F : BOOL;
    In_SenCY_Srt_Feed_H : BOOL;
    In_SenCY_Srt_Feed_F : BOOL;
    In_Sen_Unl_Conv_A_Pass : BOOL;
    In_Sen_Unl_Conv_B_Pass : BOOL;
    In_Sen_Trs_Conv_A_Arrival : BOOL;
    In_Sen_Trs_Conv_B_Arrival : BOOL;
    In_SenCY_Hnd_Feed_A_H : BOOL;
    In_SenCY_Hnd_Feed_A_F : BOOL;
    In_SenCY_Hnd_Feed_B_H : BOOL;
    In_SenCY_Hnd_Feed_B_F : BOOL;
    TimerQ_In_Sen_Supply_Container_Exist : BOOL;  (* 【X1000】供給部コンテナ有 *)
    TimerQ_In_Sen_Destacker_Stage_01_Exist : BOOL;  (* 【X1001】段バラシ1段目有 *)
    TimerQ_In_Sen_Destacker_Stage_02_Exist : BOOL;  (* 【X1002】段バラシ2段目有 *)
    TimerQ_In_Sen_Container_Arrival : BOOL;  (* 【X1003】コンテナ到着 *)
    TimerQ_In_Sen_Container_Direction_Check : BOOL;  (* 【X1004】コンテナ方向確認 *)
    TimerQ_In_Sen_Container_Pass : BOOL;  (* 【X1005】コンテナ通過 *)
    TimerQ_In_Sen_Container_Full : BOOL;  (* 【X1006】コンテナ満杯 *)
    TimerQ_In_Sen_Container_Sorting : BOOL;  (* 【X1007】コンテナ仕分け *)
    TimerQ_In_SenCY_Empty_Container_CY_H : BOOL;  (* 【X1010】空コンテナ送り 戻 *)
    TimerQ_In_SenCY_Empty_Container_CY_F : BOOL;  (* 【X1011】空コンテナ送り 行 *)
    TimerQ_In_SenCY_Sep_Claw1_H : BOOL;  (* 【X1012】段バラシ爪1 戻 *)
    TimerQ_In_SenCY_Sep_Claw1_F : BOOL;  (* 【X1013】段バラシ爪1 行 *)
    TimerQ_In_SenCY_Sep_Claw2_F : BOOL;  (* 【X1015】段バラシ爪2 行 *)
    TimerQ_In_SenCY_Sep_Claw2_H : BOOL;  (* 【X1014】段バラシ爪2 戻 *)
    TimerQ_In_SenCY_Ejc_Cont1_H : BOOL;  (* 【X1016】コンテナ排出1 戻 *)
    TimerQ_In_SenCY_Ejc_Cont1_F : BOOL;  (* 【X1017】コンテナ排出1 行 *)
    TimerQ_In_SenCY_Ejc_Cont2_H : BOOL;  (* 【X1018】コンテナ排出2 戻 *)
    TimerQ_In_SenCY_Ejc_Cont2_F : BOOL;  (* 【X1019】コンテナ排出2 行 *)
    TimerQ_In_SenCY_Box_Chk_H : BOOL;  (* 【X1020】箱入れチャック 戻 *)
    TimerQ_In_SenCY_Box_Chk_F : BOOL;  (* 【X1021】箱入れチャック 行 *)
    TimerQ_In_SenCY_Srt_Stopper_H : BOOL;  (* 【X1022】コンテナ仕分けストッパー 戻 *)
    TimerQ_In_SenCY_Srt_Stopper_F : BOOL;  (* 【X1023】コンテナ仕分けストッパー 行 *)
    TimerQ_In_SenCY_Srt_Feed_H : BOOL;  (* 【X1024】コンテナ仕分け送り 戻 *)
    TimerQ_In_SenCY_Srt_Feed_F : BOOL;  (* 【X1025】コンテナ仕分け送り 行 *)
    TimerQ_In_Sen_Unl_Conv_A_Pass : BOOL;  (* 【X1100】A(左側) 取出しコンベア 通過 *)
    TimerQ_In_Sen_Unl_Conv_B_Pass : BOOL;  (* 【X1101】B(右側) 取出しコンベア 通過 *)
    TimerQ_In_Sen_Trs_Conv_B_Arrival : BOOL;  (* 【X1103】B(右側) 搬送コンベア到着 *)
    TimerQ_In_Sen_Trs_Conv_A_Arrival : BOOL;  (* 【X1102】A(左側) 搬送コンベア到着 *)
    TimerQ_In_SenCY_Hnd_Feed_A_H : BOOL;  (* 【X1104】A(左側) コンベア受渡送り戻 *)
    TimerQ_In_SenCY_Hnd_Feed_A_F : BOOL;  (* 【X1105】A(左側) コンベア受渡送り行 *)
    TimerQ_In_SenCY_Hnd_Feed_B_H : BOOL;  (* 【X1106】B(右側) コンベア受渡送り戻 *)
    TimerQ_In_SenCY_Hnd_Feed_B_F : BOOL;  (* 【X1107】B(右側) コンベア受渡送り行 *)
    TimerQ_In_SenCY_Rev_01_Chk_B_F : BOOL;  (* 【X501】B(右側)ST4 反転1チャック開 行 *)
    Out_SW_Start_LP_GREEN : BOOL;
    Out_SW_Stop_LP_RED : BOOL;
    Out_SW_Reset_LP_Orange : BOOL;
    Out_Sg_LP_GREEN : BOOL;
    Out_Sg_LP_RED : BOOL;
    Out_Sg_LP_ORANGE : BOOL;
    Out_Sg_BUZZER : BOOL;
    Out_Accum_Cv_RESET : BOOL;
    Out_Acc_Conv_Run : BOOL;
    Out_Accum_Cv_PowerOn : BOOL;
    Out_Insp_Cv_A_Run : BOOL;
    Out_Insp_Cv_A_RESET : BOOL;
    Out_Insp_Cv_A_PowerOn : BOOL;
    Out_Insp_Cv_B_Run : BOOL;
    Out_Insp_Cv_B_RESET : BOOL;
    Out_Insp_Cv_B_PowerOn : BOOL;
    Out_CYw_Sply_Slide_A_H : BOOL;
    AutoMode : BOOL;  (* 自動運転 *)
    ManualMode : BOOL;  (* 手動運転 *)
    M9999 : BOOL;  (* 非常停止 *)
    Out_CYw_Sply_Slide_A_H_Done : BOOL;  (* 【Y616】A(左側) 供給スライド戻 動作完了 *)
    Output_A_Error_M : ARRAY[0..99] OF Bool;  (* Output一時停止：; [1] 【Y616】A(左側) 供給スライド戻 *)
    Output_A_Restart_M : ARRAY[0..99] OF Bool;  (* Output再スタート： *)
    Out_SW_Start_LP_GREEN_Auto : ARRAY[0..10] OF Bool;  (* 自動 【Y600】SWスタートランプ緑：; [1] 1 *)
    Out_SW_Start_LP_GREEN_Manual : ARRAY[0..10] OF Bool;  (* 手動 【Y600】SWスタートランプ緑： *)
    Out_SW_Stop_LP_RED_Auto : ARRAY[0..10] OF Bool;  (* 【Y601】SWストップランプ赤： *)
    Out_SW_Stop_LP_RED_Manual : ARRAY[0..10] OF Bool;  (* 【Y601】SWストップランプ赤： *)
    Out_SW_Reset_LP_Orange_Auto : ARRAY[0..10] OF Bool;  (* 【Y602】SW リセットランプ橙： *)
    Out_SW_Reset_LP_Orange_Manual : ARRAY[0..10] OF Bool;  (* 【Y602】SW リセットランプ橙： *)
    Out_Sg_LP_GREEN_Auto : ARRAY[0..10] OF Bool;  (* 【Y603】シグナルタワー緑： *)
    Out_Sg_LP_GREEN_Manual : ARRAY[0..10] OF Bool;  (* 【Y603】シグナルタワー緑： *)
    Out_Sg_LP_RED_Auto : ARRAY[0..10] OF Bool;  (* 【Y604】シグナルタワー赤： *)
    Out_Sg_LP_RED_Manual : ARRAY[0..10] OF Bool;  (* 【Y604】シグナルタワー赤： *)
    Out_Sg_LP_ORANGE_Auto : ARRAY[0..10] OF Bool;  (* 【Y605】シグナルタワー橙： *)
    Out_Sg_LP_ORANGE_Manual : ARRAY[0..10] OF Bool;  (* 【Y605】シグナルタワー橙： *)
    Out_Sg_BUZZER_Auto : ARRAY[0..10] OF Bool;  (* 【Y606】シグナルタワーブザー： *)
    Out_Sg_BUZZER_Manual : ARRAY[0..10] OF Bool;  (* 【Y606】シグナルタワーブザー： *)
    Out_Accum_Cv_RESET_Manual : ARRAY[0..10] OF Bool;  (* 【Y608】アキューム コンベア リセット： *)
    Out_Accum_Cv_RESET_Auto : ARRAY[0..10] OF Bool;  (* 【Y608】アキューム コンベア リセット： *)
    Out_Acc_Conv_Run_Manual : ARRAY[0..10] OF Bool;  (* 【Y607】アキューム コンベア運転ON： *)
    Out_Acc_Conv_Run_Auto : ARRAY[0..10] OF Bool;  (* 【Y607】アキューム コンベア運転ON： *)
    Out_Accum_Cv_PowerOn_Auto : ARRAY[0..10] OF Bool;  (* 【Y609】アキューム コンベア電源ON： *)
    Out_Accum_Cv_PowerOn_Manual : ARRAY[0..10] OF Bool;  (* 【Y609】アキューム コンベア電源ON： *)
    Out_Insp_Cv_A_Run_Auto : ARRAY[0..10] OF Bool;  (* 【Y610】A(左側) 検査 コンベア運転ON： *)
    Out_Insp_Cv_A_Run_Manual : ARRAY[0..10] OF Bool;  (* 【Y610】A(左側) 検査 コンベア運転ON： *)
    Out_Insp_Cv_A_RESET_Auto : ARRAY[0..10] OF Bool;  (* 【Y611】A(左側) 検査 コンベア リセット： *)
    Out_Insp_Cv_A_RESET_Manual : ARRAY[0..10] OF Bool;  (* 【Y611】A(左側) 検査 コンベア リセット： *)
    Out_Insp_Cv_A_PowerOn_Auto : ARRAY[0..10] OF Bool;
    Out_Insp_Cv_A_PowerOn_Manual : ARRAY[0..10] OF Bool;
    Out_Insp_Cv_B_RESET_Auto : ARRAY[0..10] OF Bool;  (* 【Y614】B(右側) 検査 コンベア リセット： *)
    Out_Insp_Cv_B_RESET_Manual : ARRAY[0..10] OF Bool;  (* 【Y614】B(右側) 検査 コンベア リセット： *)
    Out_Insp_Cv_B_Run_Manual : ARRAY[0..10] OF Bool;  (* 【Y613】B(右側) 検査 コンベア運転ON： *)
    Out_Insp_Cv_B_Run_Auto : ARRAY[0..10] OF Bool;  (* 【Y613】B(右側) 検査 コンベア運転ON： *)
    Out_CYw_Sply_Slide_A_H_Manual : ARRAY[0..10] OF Bool;  (* 【Y616】A(左側) 供給スライド戻： *)
    Out_CYw_Sply_Slide_A_H_Auto : ARRAY[0..10] OF Bool;  (* 【Y616】A(左側) 供給スライド戻： *)
    HMI_MessageNo : ARRAY[0..9] OF UINT;
    Out_CYw_Sply_Slide_A_F : BOOL;
    Out_CYw_Sply_Pick_A_H : BOOL;
    Out_CYw_Sply_Slide_A_F_Done : BOOL;  (* 【Y617】A(左側) 供給スライド行動作完了 *)
    Pause : ARRAY[0..99] OF Bool;  (* 一時停止; [3] FH A(左側) ST1; [9] FH A(左側) ST5; [10] FH B(右側) ST1; [11] FH B(右側) ST5; [12] A(左側) ST6 反転2 ワーク不一致 *)
    Out_CYw_Sply_Pick_A_F : BOOL;
    Out_CYw_Sup_Chuck_A_Cl_H : BOOL;
    Out_CYw_Sup_Chuck_A_Op_F : BOOL;
    Out_CYw_Sply_Slide_B_H : BOOL;
    Output_B_Restart_M : ARRAY[0..99] OF Bool;
    Output_B_Error_M : ARRAY[0..99] OF Bool;
    Out_CYw_Sply_Slide_B_F : BOOL;
    Out_CYw_Sply_Pick_B_H : BOOL;
    Out_CYw_Sply_Pick_B_F : BOOL;
    Out_CYw_Sup_Chuck_B_Cl_H : BOOL;
    Out_CYw_Sup_Chuck_B_Op_F : BOOL;
    Out_CYw_HgtInsp_Clp_A_H : BOOL;
    Out_CYw_HgtInsp_Clp_A_F : BOOL;
    Out_CYw_HgtInsp_Lf_A_H : BOOL;
    Out_CYw_HgtInsp_Lf_A_F : BOOL;
    Out_CYw_NG1_Pick_A_H : BOOL;
    Out_CYw_NG1_Pick_A_F : BOOL;
    Out_CYw_NG1_Chk_A_H : BOOL;
    Out_CYw_NG1_Chk_A_F : BOOL;
    Out_CYw_Rev_01_Chk_A_H : BOOL;  (* 【Y708】A(左側)ST4 反転1チャック閉 *)
    Out_CYw_Rev_01_Chk_A_F : BOOL;  (* 【Y709】A(左側)ST4 反転1チャック開 *)
    Out_CYw_Rev_01_Pick_A_H : BOOL;  (* 【Y710】A(左側)ST4 反転1ピックアップ戻 *)
    Out_CYw_Rev_01_Pick_A_F : BOOL;  (* 【Y711】A(左側)ST4 反転1ピックアップ行 *)
    Out_CYw_Rev_02_Chk_A_H : BOOL;  (* 【Y712】A(左側)ST6 反転2チャック閉 戻 *)
    Out_CYw_Rev_02_Chk_A_F : BOOL;  (* 【Y713】A(左側)ST6 反転2チャック開 行 *)
    Out_CYw_Rev_02_Pick_A_H : BOOL;  (* 【Y714】A(左側)ST6 反転2ピックアップ戻 *)
    Out_CYw_Rev_02_Pick_A_F : BOOL;  (* 【Y715】A(左側)ST6 反転2ピックアップ行 *)
    Out_CYw_Disc_Chk_A_H : BOOL;
    Out_CYw_Disc_Chk_A_F : BOOL;
    Out_CYw_Ejc_Hldr_Feed_A_F : BOOL;
    Out_CYw_Ejc_Hldr_Feed_A_H : BOOL;
    Out_CYS_Pos_01_Stopper_A : BOOL;
    Out_CYS_Pos_02_Stopper_A : BOOL;
    Out_CYS_Pos_03_Stopper_A : BOOL;
    Out_CYS_Pos_04_Stopper_A : BOOL;
    Out_CYS_Pos_05_Stopper_A : BOOL;
    Out_CYS_Pos_06_Stopper_A : BOOL;
    Out_CYw_SH_A_Turn_H : BOOL;
    Out_CYw_SH_A_Turn_F : BOOL;
    Out_CYw_NG1_Srt_A_H : BOOL;
    Out_CYw_NG1_Srt_A_F : BOOL;
    Out_CYw_HgtInsp_Clp_B_H : BOOL;
    Out_CYw_HgtInsp_Clp_B_F : BOOL;
    Out_CYw_HgtInsp_Lf_B_H : BOOL;
    Out_CYw_HgtInsp_Lf_B_F : BOOL;
    Out_CYw_NG1_Pick_B_H : BOOL;
    Out_CYw_NG1_Pick_B_F : BOOL;
    Out_CYw_NG1_Chk_B_H : BOOL;
    Out_CYw_NG1_Chk_B_F : BOOL;
    Out_CYw_Rev_01_Chk_B_H : BOOL;  (* 【Y808】B(右側)ST4 反転1チャック閉 戻 *)
    Out_CYw_Rev_01_Chk_B_F : BOOL;  (* 【Y809】B(右側)ST4 反転1チャック開 戻 *)
    Out_CYw_Rev_01_Pick_B_H : BOOL;  (* 【Y810】B(右側)ST4 反転1ピックアップ戻 *)
    Out_CYw_Rev_01_Pick_B_F : BOOL;  (* 【Y811】B(右側)ST4 反転1ピックアップ行 *)
    Out_CYw_Rev_02_Chk_B_H : BOOL;  (* 【Y812】B(右側)ST6 反転2チャック閉 戻 *)
    Out_CYw_Rev_02_Chk_B_F : BOOL;  (* 【Y813】B(右側)ST6 反転2チャック開 行 *)
    Out_CYw_Rev_02_Pick_B_H : BOOL;  (* 【Y814】B(右側)ST6 反転2ピックアップ戻 *)
    Out_CYw_Rev_02_Pick_B_F : BOOL;  (* 【Y815】B(右側)ST6 反転2ピックアップ行 *)
    Out_CYw_Disc_Chk_B_H : BOOL;
    Out_CYw_Disc_Chk_B_F : BOOL;
    Out_CYw_Ejc_Hldr_Feed_B_H : BOOL;
    Out_CYw_Ejc_Hldr_Feed_B_F : BOOL;
    Out_CYS_Pos_01_Stopper_B : BOOL;
    Out_CYS_Pos_02_Stopper_B : BOOL;
    Out_CYS_Pos_03_Stopper_B : BOOL;
    Out_CYS_Pos_04_Stopper_B : BOOL;
    Out_CYS_Pos_05_Stopper_B : BOOL;
    Out_CYS_Pos_06_Stopper_B : BOOL;
    Out_CYw_SH_B_Turn_H : BOOL;
    Out_CYw_SH_B_Turn_F : BOOL;
    Out_CYw_NG1_Srt_B_H : BOOL;
    Out_CYw_NG1_Srt_B_F : BOOL;
    Output_Share_Restart_M : ARRAY[0..99] OF Bool;  (* 共有シリンダ再開： *)
    Output_Share_Error_M : ARRAY[0..99] OF Bool;  (* 共有シリンダエラー： *)
    Out_CYw_Empty_Container_CY_H : BOOL;
    Out_CYw_Empty_Container_CY_F : BOOL;
    Out_CYw_Sep_Claw_F : BOOL;
    Out_CYw_Sep_Claw_H : BOOL;
    Out_CYw_Ejc_Cont_H : BOOL;
    Out_CYw_Ejc_Cont_F : BOOL;
    Out_CYw_Box_Chuck_H : BOOL;
    Out_CYw_Box_Chuck_F : BOOL;
    Out_CYw_Srt_Stopper_H : BOOL;
    Out_CYw_Srt_Stopper_F : BOOL;
    Out_CYw_Srt_Feed_H : BOOL;
    Out_CYw_Srt_Feed_F : BOOL;
    Out_CYw_Hnd_Feed_A_H : BOOL;
    Out_CYw_Hnd_Feed_A_F : BOOL;
    Out_CYw_Hnd_Feed_B_H : BOOL;
    Out_CYw_Hnd_Feed_B_F : BOOL;
    Out_CYw_Hnd_Feed_B_F_Done : BOOL;  (* 【Y1303】B(右側) コンベア受渡送り行 動作完了 *)
    Out_CYw_Hnd_Feed_B_F_Manual : ARRAY[0..10] OF Bool;  (* 手動【Y1303】B(右側) コンベア受渡送り行： *)
    Out_CYw_Hnd_Feed_B_F_Auto : ARRAY[0..10] OF Bool;  (* 自動【Y1303】B(右側) コンベア受渡送り行： *)
    Out_CYw_Hnd_Feed_B_H_Done : BOOL;  (* 【Y1302】B(右側) コンベア受渡送り戻 動作完了 *)
    Out_CYw_Hnd_Feed_B_H_Manual : ARRAY[0..10] OF Bool;  (* 手動【Y1302】B(右側) コンベア受渡送り戻： *)
    Out_CYw_Hnd_Feed_B_H_Auto : ARRAY[0..10] OF Bool;  (* 自動【Y1302】B(右側) コンベア受渡送り戻： *)
    Out_CYw_Hnd_Feed_A_F_Done : BOOL;  (* 【Y1301】A(左側) コンベア受渡送り行 動作完了 *)
    Out_CYw_Hnd_Feed_A_F_Manual : ARRAY[0..10] OF Bool;  (* 手動【Y1301】A(左側) コンベア受渡送り行： *)
    Out_CYw_Srt_Feed_H_Manual : ARRAY[0..10] OF Bool;  (* 手動【Y1210】コンテナ仕分け送り 戻： *)
    Out_CYw_Srt_Feed_H_Done : BOOL;  (* 【Y1210】コンテナ仕分け送り 戻 動作完了 *)
    Out_CYw_Srt_Feed_F_Auto : ARRAY[0..10] OF Bool;  (* 自動【Y1211】コンテナ仕分け送り 行： *)
    Out_CYw_Srt_Feed_F_Manual : ARRAY[0..10] OF Bool;  (* 手動【Y1211】コンテナ仕分け送り 行： *)
    Out_CYw_Srt_Feed_F_Done : BOOL;  (* 【Y1211】コンテナ仕分け送り 行 動作完了 *)
    Out_CYw_Hnd_Feed_A_H_Auto : ARRAY[0..10] OF Bool;  (* 自動【Y1300】A(左側) コンベア受渡送り戻： *)
    Out_CYw_Hnd_Feed_A_H_Manual : ARRAY[0..10] OF Bool;  (* 手動【Y1300】A(左側) コンベア受渡送り戻： *)
    Out_CYw_Hnd_Feed_A_H_Done : BOOL;  (* 【Y1300】A(左側) コンベア受渡送り戻 動作完了 *)
    Out_CYw_Hnd_Feed_A_F_Auto : ARRAY[0..10] OF Bool;  (* 自動【Y1301】A(左側) コンベア受渡送り行： *)
    Out_CYw_Empty_Container_CY_F_Done : BOOL;  (* 【Y1201】空コンテナ送り 行 動作完了 *)
    Out_CYw_Sep_Claw_H_Auto : ARRAY[0..10] OF Bool;  (* 自動【Y1202】段バラシ爪 戻： *)
    Out_CYw_Sep_Claw_H_Manual : ARRAY[0..10] OF Bool;  (* 手動【Y1202】段バラシ爪 戻： *)
    Out_CYw_Sep_Claw_H_Done : BOOL;  (* 【Y1202】段バラシ爪 戻 動作完了 *)
    Out_CYw_Sep_Claw_F_Auto : ARRAY[0..10] OF Bool;  (* 自動【Y1203】段バラシ爪 行： *)
    Out_CYw_Sep_Claw_F_Manual : ARRAY[0..10] OF Bool;  (* 手動【Y1203】段バラシ爪 行： *)
    Out_CYw_Sep_Claw_F_Done : BOOL;  (* 【Y1203】段バラシ爪 行 動作完了 *)
    Out_CYw_Ejc_Cont_H_Auto : ARRAY[0..10] OF Bool;  (* 自動【Y1204】コンテナ排出 戻： *)
    Out_CYw_Ejc_Cont_H_Manual : ARRAY[0..10] OF Bool;  (* 手動【Y1204】コンテナ排出 戻： *)
    Out_CYw_Ejc_Cont_H_Done : BOOL;  (* 【Y1204】コンテナ排出 戻 動作完了 *)
    Out_CYw_Ejc_Cont_F_Auto : ARRAY[0..10] OF Bool;  (* 自動【Y1205】コンテナ排出 行： *)
    Out_CYw_Ejc_Cont_F_Manual : ARRAY[0..10] OF Bool;  (* 手動【Y1205】コンテナ排出 行： *)
    Out_CYw_Ejc_Cont_F_Done : BOOL;  (* 【Y1205】コンテナ排出 行 動作完了 *)
    Out_CYw_Box_Chuck_H_Auto : ARRAY[0..10] OF Bool;  (* 自動【Y1206】箱入れチャック 戻： *)
    Out_CYw_Box_Chuck_H_Manual : ARRAY[0..10] OF Bool;  (* 手動【Y1206】箱入れチャック 戻： *)
    Out_CYw_Box_Chuck_H_Done : BOOL;  (* 【Y1206】箱入れチャック 戻 動作完了 *)
    Out_CYw_Box_Chuck_F_Auto : ARRAY[0..10] OF Bool;  (* 自動【Y1207】箱入れチャック 行： *)
    Out_CYw_Box_Chuck_F_Manual : ARRAY[0..10] OF Bool;  (* 手動【Y1207】箱入れチャック 行： *)
    Out_CYw_Box_Chuck_F_Done : BOOL;  (* 【Y1207】箱入れチャック 行 動作完了 *)
    Out_CYw_Srt_Stopper_H_Auto : ARRAY[0..10] OF Bool;  (* 自動【Y1208】コンテナ仕分けストッパー 戻： *)
    Out_CYw_Srt_Stopper_H_Manual : ARRAY[0..10] OF Bool;  (* 手動【Y1208】コンテナ仕分けストッパー 戻 行： *)
    Out_CYw_Srt_Stopper_H_Done : BOOL;  (* 【Y1208】コンテナ仕分けストッパー 戻 動作完了 *)
    Out_CYw_Srt_Stopper_F_Auto : ARRAY[0..10] OF Bool;  (* 自動【Y1209】コンテナ仕分けストッパー 行： *)
    Out_CYw_Srt_Stopper_F_Manual : ARRAY[0..10] OF Bool;  (* 手動【Y1209】コンテナ仕分けストッパー 行： *)
    Out_CYw_Srt_Stopper_F_Done : BOOL;  (* 【Y1209】コンテナ仕分けストッパー 行 動作完了 *)
    Out_CYw_Srt_Feed_H_Auto : ARRAY[0..10] OF Bool;  (* 自動【Y1210】コンテナ仕分け送り 戻： *)
    Out_CYS_Pos_04_Stopper_B_H_Auto : ARRAY[0..10] OF Bool;  (* 自動【Y823】B(右側) 位置4ストッパー戻： *)
    Out_CYS_Pos_04_Stopper_B_H_Manual : ARRAY[0..10] OF Bool;  (* 手動【Y823】B(右側) 位置4ストッパー戻： *)
    Out_CYS_Pos_04_Stopper_B_H_Done : BOOL;  (* 【Y823】B(右側) 位置4ストッパー戻 動作完了 *)
    Out_CYS_Pos_04_Stopper_B_F_Auto : ARRAY[0..10] OF Bool;  (* 自動【Y823】B(右側) 位置4ストッパー行： *)
    Out_CYS_Pos_04_Stopper_B_F_Manual : ARRAY[0..10] OF Bool;  (* 手動【Y823】B(右側) 位置4ストッパー行： *)
    Out_CYS_Pos_04_Stopper_B_F_Done : BOOL;  (* 【Y823】B(右側) 位置4ストッパー行 動作完了 *)
    Out_CYS_Pos_05_Stopper_B_H_Auto : ARRAY[0..10] OF Bool;  (* 自動【Y824】B(右側) 位置5ストッパー戻： *)
    Out_CYS_Pos_05_Stopper_B_H_Manual : ARRAY[0..10] OF Bool;  (* 手動【Y824】B(右側) 位置5ストッパー戻： *)
    Out_CYS_Pos_05_Stopper_B_H_Done : BOOL;  (* 【Y824】B(右側) 位置5ストッパー戻 動作完了 *)
    Out_CYS_Pos_05_Stopper_B_F_Auto : ARRAY[0..10] OF Bool;  (* 自動【Y824】B(右側) 位置5ストッパー行： *)
    Out_CYS_Pos_05_Stopper_B_F_Manual : ARRAY[0..10] OF Bool;  (* 手動【Y824】B(右側) 位置5ストッパー行： *)
    Out_CYS_Pos_05_Stopper_B_F_Done : BOOL;  (* 【Y824】B(右側) 位置5ストッパー行 動作完了 *)
    Out_CYS_Pos_06_Stopper_B_H_Auto : ARRAY[0..10] OF Bool;  (* 自動【Y825】B(右側) 位置6ストッパー戻： *)
    Out_CYS_Pos_06_Stopper_B_H_Manual : ARRAY[0..10] OF Bool;  (* 手動【Y825】B(右側) 位置6ストッパー戻： *)
    Out_CYS_Pos_06_Stopper_B_H_Done : BOOL;  (* 【Y825】B(右側) 位置6ストッパー戻 動作完了 *)
    Out_CYS_Pos_06_Stopper_B_F_Auto : ARRAY[0..10] OF Bool;  (* 自動【Y825】B(右側) 位置6ストッパー行： *)
    Out_CYS_Pos_06_Stopper_B_F_Manual : ARRAY[0..10] OF Bool;  (* 手動【Y825】B(右側) 位置6ストッパー行： *)
    Out_CYS_Pos_06_Stopper_B_F_Done : BOOL;  (* 【Y825】B(右側) 位置6ストッパー行 動作完了 *)
    Out_CYw_SH_B_Turn_H_Auto : ARRAY[0..10] OF Bool;  (* 自動【Y826】B(右側) ストックフォルダターン戻： *)
    Out_CYw_SH_B_Turn_H_Manual : ARRAY[0..10] OF Bool;  (* 手動【Y826】B(右側) ストックフォルダターン戻： *)
    Out_CYw_SH_B_Turn_H_Done : BOOL;  (* 【Y826】B(右側) ストックフォルダターン戻 動作完了 *)
    Out_CYw_SH_B_Turn_F_Manual : ARRAY[0..10] OF Bool;  (* 自動【Y827】B(右側) ストックフォルダターン行： *)
    Out_CYw_SH_B_Turn_F_Auto : ARRAY[0..10] OF Bool;  (* 手動【Y827】B(右側) ストックフォルダターン行： *)
    Out_CYw_SH_B_Turn_F_Done : BOOL;  (* 【Y827】B(右側) ストックフォルダターン行 動作完了 *)
    Out_CYw_NG1_Srt_B_H_Auto : ARRAY[0..10] OF Bool;  (* 自動【Y828】B(右側) NG1仕分け 戻： *)
    Out_CYw_NG1_Srt_B_H_Manual : ARRAY[0..10] OF Bool;  (* 手動【Y828】B(右側) NG1仕分け 戻： *)
    Out_CYw_NG1_Srt_B_H_Done : BOOL;  (* 【Y828】B(右側) NG1仕分け 戻 動作完了 *)
    Out_CYw_NG1_Srt_B_F_Auto : ARRAY[0..10] OF Bool;  (* 自動【Y829】B(右側) NG1仕分け 行： *)
    Out_CYw_NG1_Srt_B_F_Manual : ARRAY[0..10] OF Bool;  (* 手動【Y829】B(右側) NG1仕分け 行： *)
    Out_CYw_NG1_Srt_B_F_Done : BOOL;  (* 【Y829】B(右側) NG1仕分け 行 動作完了 *)
    Out_CYw_Empty_Container_CY_H_Manual : ARRAY[0..10] OF Bool;  (* 手動【Y1200】空コンテナ送り 戻： *)
    Out_CYw_Empty_Container_CY_H_Auto : ARRAY[0..10] OF Bool;  (* 自動【Y1200】空コンテナ送り 戻： *)
    Out_CYw_Empty_Container_CY_H_Done : BOOL;  (* 【Y1200】空コンテナ送り 戻 動作完了 *)
    Out_CYw_Empty_Container_CY_F_Auto : ARRAY[0..10] OF Bool;  (* 自動【Y1201】空コンテナ送り 行： *)
    Out_CYw_Empty_Container_CY_F_Manual : ARRAY[0..10] OF Bool;  (* 手動【Y1201】空コンテナ送り 行： *)
    Out_CYw_Rev_02_Pick_B_H_Manual : ARRAY[0..10] OF Bool;  (* 手動【Y814】B(右側)ST6 反転2ピックアップ戻： *)
    Out_CYw_Rev_02_Pick_B_H_Done : BOOL;  (* 【Y814】B(右側)ST6 反転2ピックアップ戻 動作完了 *)
    Out_CYw_Rev_02_Pick_B_F_Auto : ARRAY[0..10] OF Bool;  (* 自動【Y815】B(右側)ST6 反転2ピックアップ行 ： *)
    Out_CYw_Rev_02_Pick_B_F_Manual : ARRAY[0..10] OF Bool;  (* 手動【Y815】B(右側)ST6 反転2ピックアップ行： *)
    Out_CYw_Rev_02_Pick_B_F_Done : BOOL;  (* 【Y815】B(右側)ST6 反転2ピックアップ行 動作完了 *)
    Out_CYw_Disc_Chk_B_H_Auto : ARRAY[0..10] OF Bool;  (* 自動【Y816】B(右側) 排出チャック閉 戻 ： *)
    Out_CYw_Disc_Chk_B_H_Manual : ARRAY[0..10] OF Bool;  (* 手動【Y816】B(右側) 排出チャック閉 戻： *)
    Out_CYw_Disc_Chk_B_H_Done : BOOL;  (* 【Y816】B(右側) 排出チャック閉 戻 動作完了 *)
    Out_CYw_Disc_Chk_B_F_Auto : ARRAY[0..10] OF Bool;  (* 自動【Y817】B(右側) 排出チャック開 行 ： *)
    Out_CYw_Disc_Chk_B_F_Manual : ARRAY[0..10] OF Bool;  (* 手動【Y817】B(右側) 排出チャック開 行： *)
    Out_CYw_Disc_Chk_B_F_Done : BOOL;  (* 【Y817】B(右側) 排出チャック開 行 動作完了 *)
    Out_CYw_Ejc_Hldr_Feed_B_H_Auto : ARRAY[0..10] OF Bool;  (* 自動【Y818】B(右側) 排出フォルダ送り戻： *)
    Out_CYw_Ejc_Hldr_Feed_B_H_Manual : ARRAY[0..10] OF Bool;  (* 手動【Y818】B(右側) 排出フォルダ送り戻： *)
    Out_CYw_Ejc_Hldr_Feed_B_H_Done : BOOL;  (* 【Y818】B(右側) 排出フォルダ送り戻 動作完了 *)
    Out_CYw_Ejc_Hldr_Feed_B_F_Auto : ARRAY[0..10] OF Bool;  (* 自動【Y819】B(右側) 排出フォルダ送り行： *)
    Out_CYw_Ejc_Hldr_Feed_B_F_Manual : ARRAY[0..10] OF Bool;  (* 手動【Y819】B(右側) 排出フォルダ送り行： *)
    Out_CYw_Ejc_Hldr_Feed_B_F_Done : BOOL;  (* 【Y819】B(右側) 排出フォルダ送り行 動作完了 *)
    Out_CYS_Pos_01_Stopper_B_H_Auto : ARRAY[0..10] OF Bool;  (* 自動【Y820】B(右側) 位置1ストッパー戻： *)
    Out_CYS_Pos_01_Stopper_B_H_Manual : ARRAY[0..10] OF Bool;  (* 手動【Y820】B(右側) 位置1ストッパー戻： *)
    Out_CYS_Pos_01_Stopper_B_H_Done : BOOL;  (* 【Y820】B(右側) 位置1ストッパー戻 動作完了 *)
    Out_CYS_Pos_01_Stopper_B_F_Auto : ARRAY[0..10] OF Bool;  (* 自動【Y820】B(右側) 位置1ストッパー 行： *)
    Out_CYS_Pos_01_Stopper_B_F_Manual : ARRAY[0..10] OF Bool;  (* 手動【Y820】B(右側) 位置1ストッパー 行： *)
    Out_CYS_Pos_01_Stopper_B_F_Done : BOOL;  (* 【Y820】B(右側) 位置1ストッパー 行 動作完了 *)
    Out_CYS_Pos_02_Stopper_B_H_Auto : ARRAY[0..10] OF Bool;  (* 自動【Y821】B(右側) 位置2ストッパー戻： *)
    Out_CYS_Pos_02_Stopper_B_H_Manual : ARRAY[0..10] OF Bool;  (* 手動【Y821】B(右側) 位置2ストッパー戻： *)
    Out_CYS_Pos_02_Stopper_B_H_Done : BOOL;  (* 【Y821】B(右側) 位置2ストッパー戻 動作完了 *)
    Out_CYS_Pos_02_Stopper_B_F_Auto : ARRAY[0..10] OF Bool;  (* 自動【Y821】B(右側) 位置2ストッパー行： *)
    Out_CYS_Pos_02_Stopper_B_F_Manual : ARRAY[0..10] OF Bool;  (* 手動【Y821】B(右側) 位置2ストッパー行： *)
    Out_CYS_Pos_02_Stopper_B_F_Done : BOOL;  (* 【Y821】B(右側) 位置2ストッパー行 動作完了 *)
    Out_CYS_Pos_03_Stopper_B_H_Auto : ARRAY[0..10] OF Bool;  (* 自動【Y822】B(右側) 位置3ストッパー戻： *)
    Out_CYS_Pos_03_Stopper_B_H_Manual : ARRAY[0..10] OF Bool;  (* 手動【Y822】B(右側) 位置3ストッパー戻： *)
    Out_CYS_Pos_03_Stopper_B_H_Done : BOOL;  (* 【Y822】B(右側) 位置3ストッパー戻 動作完了 *)
    Out_CYS_Pos_03_Stopper_B_F_Auto : ARRAY[0..10] OF Bool;  (* 自動【Y822】B(右側) 位置3ストッパー行： *)
    Out_CYS_Pos_03_Stopper_B_F_Manual : ARRAY[0..10] OF Bool;  (* 手動【Y822】B(右側) 位置3ストッパー行： *)
    Out_CYS_Pos_03_Stopper_B_F_Done : BOOL;  (* 【Y822】B(右側) 位置3ストッパー行 動作完了 *)
    Out_CYw_HgtInsp_Lf_B_H_Done : BOOL;  (* 【Y802】B(右側) 高さ検査持上戻 動作完了 *)
    Out_CYw_HgtInsp_Lf_B_F_Auto : ARRAY[0..10] OF Bool;  (* 自動【Y803】B(右側) 高さ検査持上行： *)
    Out_CYw_HgtInsp_Lf_B_F_Manual : ARRAY[0..10] OF Bool;  (* 手動【Y803】B(右側) 高さ検査持上行： *)
    Out_CYw_HgtInsp_Lf_B_F_Done : BOOL;  (* 【Y803】B(右側) 高さ検査持上行 動作完了 *)
    Out_CYw_NG1_Pick_B_H_Auto : ARRAY[0..10] OF Bool;  (* 自動【Y804】B(右側) NG1ピックアップ戻： *)
    Out_CYw_NG1_Pick_B_H_Manual : ARRAY[0..10] OF Bool;  (* 手動【Y804】B(右側) NG1ピックアップ戻： *)
    Out_CYw_NG1_Pick_B_H_Done : BOOL;  (* 【Y804】B(右側) NG1ピックアップ戻 動作完了 *)
    Out_CYw_NG1_Pick_B_F_Auto : ARRAY[0..10] OF Bool;  (* 自動【Y805】B(右側) NG1ピックアップ行： *)
    Out_CYw_NG1_Pick_B_F_Manual : ARRAY[0..10] OF Bool;  (* 手動【Y805】B(右側) NG1ピックアップ行： *)
    Out_CYw_NG1_Pick_B_F_Done : BOOL;  (* 【Y805】B(右側) NG1ピックアップ行 動作完了 *)
    Out_CYw_NG1_Chk_B_H_Auto : ARRAY[0..10] OF Bool;  (* 自動【Y806】B(右側) NG1チャック戻： *)
    Out_CYw_NG1_Chk_B_H_Manual : ARRAY[0..10] OF Bool;  (* 手動【Y806】B(右側) NG1チャック戻： *)
    Out_CYw_NG1_Chk_B_H_Done : BOOL;  (* 【Y806】B(右側) NG1チャック戻 動作完了 *)
    Out_CYw_NG1_Chk_B_F_Auto : ARRAY[0..10] OF Bool;  (* 自動【Y807】B(右側) NG1チャック行： *)
    Out_CYw_NG1_Chk_B_F_Manual : ARRAY[0..10] OF Bool;  (* 手動【Y807】B(右側) NG1チャック行： *)
    Out_CYw_NG1_Chk_B_F_Done : BOOL;  (* 【Y807】B(右側) NG1チャック行 動作完了 *)
    Out_CYw_Rev_01_Chk_B_H_Auto : ARRAY[0..10] OF Bool;  (* 自動【Y808】B(右側)ST4 反転1チャック閉 戻： *)
    Out_CYw_Rev_01_Chk_B_H_Manual : ARRAY[0..10] OF Bool;  (* 手動【Y808】B(右側)ST4 反転1チャック閉 戻： *)
    Out_CYw_Rev_01_Chk_B_H_Done : BOOL;  (* 【Y808】B(右側)ST4 反転1チャック閉 戻 動作完了 *)
    Out_CYw_Rev_01_Chk_B_F_Auto : ARRAY[0..10] OF Bool;  (* 自動【Y809】B(右側)ST4 反転1チャック開 戻： *)
    Out_CYw_Rev_01_Chk_B_F_Manual : ARRAY[0..10] OF Bool;  (* 手動【Y809】B(右側)ST4 反転1チャック開 戻： *)
    Out_CYw_Rev_01_Chk_B_F_Done : BOOL;  (* 【Y809】B(右側)ST4 反転1チャック開 戻 動作完了 *)
    Out_CYw_Rev_01_Pick_B_H_Auto : ARRAY[0..10] OF Bool;  (* 自動【Y810】B(右側)ST4 反転1ピックアップ戻： *)
    Out_CYw_Rev_01_Pick_B_H_Manual : ARRAY[0..10] OF Bool;  (* 手動【Y810】B(右側)ST4 反転1ピックアップ戻： *)
    Out_CYw_Rev_01_Pick_B_H_Done : BOOL;  (* 【Y810】B(右側)ST4 反転1ピックアップ戻 動作完了 *)
    Out_CYw_Rev_01_Pick_B_F_Auto : ARRAY[0..10] OF Bool;  (* 自動【Y811】B(右側)ST4 反転1ピックアップ行： *)
    Out_CYw_Rev_01_Pick_B_F_Manual : ARRAY[0..10] OF Bool;  (* 手動【Y811】B(右側)ST4 反転1ピックアップ行： *)
    Out_CYw_Rev_01_Pick_B_F_Done : BOOL;  (* 【Y811】B(右側)ST4 反転1ピックアップ行 動作完了 *)
    Out_CYw_Rev_02_Chk_B_H_Auto : ARRAY[0..10] OF Bool;  (* 自動【Y812】B(右側)ST6 反転2チャック閉 戻： *)
    Out_CYw_Rev_02_Chk_B_H_Manual : ARRAY[0..10] OF Bool;  (* 手動【Y812】B(右側)ST6 反転2チャック閉 戻： *)
    Out_CYw_Rev_02_Chk_B_H_Done : BOOL;  (* 【Y812】B(右側)ST6 反転2チャック閉 戻 動作完了 *)
    Out_CYw_Rev_02_Chk_B_F_Auto : ARRAY[0..10] OF Bool;  (* 自動【Y813】B(右側)ST6 反転2チャック開 行 ： *)
    Out_CYw_Rev_02_Chk_B_F_Manual : ARRAY[0..10] OF Bool;  (* 手動【Y813】B(右側)ST6 反転2チャック開 行： *)
    Out_CYw_Rev_02_Chk_B_F_Done : BOOL;  (* 【Y813】B(右側)ST6 反転2チャック開 行 動作完了 *)
    Out_CYw_Rev_02_Pick_B_H_Auto : ARRAY[0..10] OF Bool;  (* 自動【Y814】B(右側)ST6 反転2ピックアップ戻 ： *)
    Out_CYw_HgtInsp_Clp_B_H_Done : BOOL;  (* 【Y800】B(右側) 高さ検査押え戻 動作完了 *)
    Out_CYw_HgtInsp_Clp_B_H_Auto : ARRAY[0..10] OF Bool;  (* 自動【Y800】B(右側) 高さ検査押え戻： *)
    Out_CYw_HgtInsp_Clp_B_H_Manual : ARRAY[0..10] OF Bool;  (* 手動【Y800】B(右側) 高さ検査押え戻： *)
    Out_CYw_HgtInsp_Clp_B_F_Auto : ARRAY[0..10] OF Bool;  (* 自動【Y801】B(右側) 高さ検査押え行： *)
    Out_CYw_HgtInsp_Clp_B_F_Manual : ARRAY[0..10] OF Bool;  (* 手動【Y801】B(右側) 高さ検査押え行： *)
    Out_CYw_HgtInsp_Clp_B_F_Done : BOOL;  (* 【Y801】B(右側) 高さ検査押え行 動作完了 *)
    Out_CYw_HgtInsp_Lf_B_H_Auto : ARRAY[0..10] OF Bool;  (* 自動【Y802】B(右側) 高さ検査持上戻： *)
    Out_CYw_HgtInsp_Lf_B_H_Manual : ARRAY[0..10] OF Bool;  (* 手動【Y802】B(右側) 高さ検査持上戻： *)
    Out_CYS_Pos_03_Stopper_A_H_Manual : ARRAY[0..10] OF Bool;  (* 手動【Y722】A(左側) 位置3ストッパー戻： *)
    Out_CYS_Pos_03_Stopper_A_H_Done : BOOL;  (* 【Y722】A(左側) 位置3ストッパー戻 動作完了 *)
    Out_CYS_Pos_03_Stopper_A_F_Auto : ARRAY[0..10] OF Bool;  (* 自動【Y722】A(左側) 位置3ストッパー行： *)
    Out_CYS_Pos_03_Stopper_A_F_Manual : ARRAY[0..10] OF Bool;  (* 手動【Y722】A(左側) 位置3ストッパー行： *)
    Out_CYS_Pos_03_Stopper_A_F_Done : BOOL;  (* 【Y722】A(左側) 位置3ストッパー行 動作完了 *)
    Out_CYS_Pos_04_Stopper_A_H_Auto : ARRAY[0..10] OF Bool;  (* 自動【Y723】A(左側) 位置4ストッパー戻： *)
    Out_CYS_Pos_04_Stopper_A_H_Manual : ARRAY[0..10] OF Bool;  (* 手動【Y723】A(左側) 位置4ストッパー戻： *)
    Out_CYS_Pos_04_Stopper_A_H_Done : BOOL;  (* 【Y723】A(左側) 位置4ストッパー戻 動作完了 *)
    Out_CYS_Pos_04_Stopper_A_F_Auto : ARRAY[0..10] OF Bool;  (* 自動【Y723】A(左側) 位置4ストッパー行： *)
    Out_CYS_Pos_04_Stopper_A_F_Manual : ARRAY[0..10] OF Bool;  (* 手動【Y723】A(左側) 位置4ストッパー行： *)
    Out_CYS_Pos_04_Stopper_A_F_Done : BOOL;  (* 【Y723】A(左側) 位置4ストッパー行 動作完了 *)
    Out_CYS_Pos_05_Stopper_A_H_Auto : ARRAY[0..10] OF Bool;  (* 自動【Y724】A(左側) 位置5ストッパー戻：; [2] A(左側) ST5 カメラ2検査開始 *)
    Out_CYS_Pos_05_Stopper_A_H_Manual : ARRAY[0..10] OF Bool;  (* 手動【Y724】A(左側) 位置5ストッパー戻： *)
    Out_CYS_Pos_05_Stopper_A_H_Done : BOOL;  (* 【Y724】A(左側) 位置5ストッパー戻 動作完了 *)
    Out_CYS_Pos_05_Stopper_A_F_Auto : ARRAY[0..10] OF Bool;  (* 自動【Y724】A(左側) 位置5ストッパー行： *)
    Out_CYS_Pos_05_Stopper_A_F_Manual : ARRAY[0..10] OF Bool;  (* 手動【Y724】A(左側) 位置5ストッパー行： *)
    Out_CYS_Pos_05_Stopper_A_F_Done : BOOL;  (* 【Y724】A(左側) 位置5ストッパー行 動作完了 *)
    Out_CYS_Pos_06_Stopper_A_H_Auto : ARRAY[0..10] OF Bool;  (* 自動【Y725】A(左側) 位置6ストッパー戻：; [1] A(左側)検査完了後; [2] A(左側) ST6 原点位置移動 *)
    Out_CYS_Pos_06_Stopper_A_H_Manual : ARRAY[0..10] OF Bool;  (* 手動【Y725】A(左側) 位置6ストッパー戻： *)
    Out_CYS_Pos_06_Stopper_A_H_Done : BOOL;  (* 【Y725】A(左側) 位置6ストッパー戻 動作完了 *)
    Out_CYS_Pos_06_Stopper_A_F_Auto : ARRAY[0..10] OF Bool;  (* 自動【Y725】A(左側) 位置6ストッパー行： *)
    Out_CYS_Pos_06_Stopper_A_F_Manual : ARRAY[0..10] OF Bool;  (* 手動【Y725】A(左側) 位置6ストッパー行： *)
    Out_CYS_Pos_06_Stopper_A_F_Done : BOOL;  (* 【Y725】A(左側) 位置6ストッパー行 動作完了 *)
    Out_CYw_SH_A_Turn_H_Auto : ARRAY[0..10] OF Bool;  (* 自動【Y726】A(左側) ストックフォルダターン戻： *)
    Out_CYw_SH_A_Turn_H_Manual : ARRAY[0..10] OF Bool;  (* 手動【Y726】A(左側) ストックフォルダターン戻： *)
    Out_CYw_SH_A_Turn_H_Done : BOOL;  (* 【Y726】A(左側) ストックフォルダターン戻 動作完了 *)
    Out_CYw_SH_A_Turn_F_Auto : ARRAY[0..10] OF Bool;  (* 自動【Y727】A(左側) ストックフォルダターン行： *)
    Out_CYw_SH_A_Turn_F_Manual : ARRAY[0..10] OF Bool;  (* 手動【Y727】A(左側) ストックフォルダターン行： *)
    Out_CYw_SH_A_Turn_F_Done : BOOL;  (* 【Y727】A(左側) ストックフォルダターン行 動作完了 *)
    Out_CYw_NG1_Srt_A_H_Auto : ARRAY[0..10] OF Bool;  (* 自動【Y728】A(左側) NG1仕分け 戻： *)
    Out_CYw_NG1_Srt_A_H_Manual : ARRAY[0..10] OF Bool;  (* 手動【Y728】A(左側) NG1仕分け 戻： *)
    Out_CYw_NG1_Srt_A_H_Done : BOOL;  (* 【Y728】A(左側) NG1仕分け 戻 動作完了 *)
    Out_CYw_NG1_Srt_A_F_Auto : ARRAY[0..10] OF Bool;  (* 自動【Y729】A(左側) NG1仕分け行： *)
    Out_CYw_NG1_Srt_A_F_Manual : ARRAY[0..10] OF Bool;  (* 手動【Y729】A(左側) NG1仕分け行： *)
    Out_CYw_NG1_Srt_A_F_Done : BOOL;  (* 【Y729】A(左側) NG1仕分け行 動作完了 *)
    Out_CYS_Pos_01_Stopper_A_F_Auto : ARRAY[0..10] OF Bool;  (* 自動【Y720】A(左側) 位置1ストッパー行： *)
    Out_CYS_Pos_01_Stopper_A_F_Manual : ARRAY[0..10] OF Bool;  (* 手動【Y720】A(左側) 位置1ストッパー 行： *)
    Out_CYS_Pos_02_Stopper_A_H_Auto : ARRAY[0..10] OF Bool;  (* 自動【Y721】A(左側) 位置2ストッパー戻： *)
    Out_CYS_Pos_02_Stopper_A_H_Manual : ARRAY[0..10] OF Bool;  (* 手動【Y721】A(左側) 位置2ストッパー戻： *)
    Out_CYS_Pos_02_Stopper_A_H_Done : BOOL;  (* 【Y721】A(左側) 位置2ストッパー戻 動作完了 *)
    Out_CYS_Pos_02_Stopper_A_F_Auto : ARRAY[0..10] OF Bool;  (* 自動【Y721】A(左側) 位置2ストッパー行： *)
    Out_CYS_Pos_02_Stopper_A_F_Manual : ARRAY[0..10] OF Bool;  (* 手動【Y721】A(左側) 位置2ストッパー行： *)
    Out_CYS_Pos_02_Stopper_A_F_Done : BOOL;  (* 【Y721】A(左側) 位置2ストッパー行 動作完了 *)
    Out_CYS_Pos_03_Stopper_A_H_Auto : ARRAY[0..10] OF Bool;  (* 自動【Y722】A(左側) 位置3ストッパー戻： *)
    Out_CYw_Rev_02_Pick_A_H_Auto : ARRAY[0..10] OF Bool;  (* 自動【Y714】A(左側)ST6 反転2ピックアップ戻 ：; [1] A(左側) ST6 反転前戻; [2] A(左側) ST6 設置後戻 *)
    Out_CYw_Rev_02_Pick_A_H_Manual : ARRAY[0..10] OF Bool;  (* 手動【Y714】A(左側)ST6 反転2ピックアップ戻 ： *)
    Out_CYw_Rev_02_Pick_A_H_Done : BOOL;  (* 【Y714】A(左側)ST6 反転2ピックアップ戻 動作完了 *)
    Out_CYw_Rev_02_Pick_A_F_Auto : ARRAY[0..10] OF Bool;  (* 自動【Y715】A(左側)ST6 反転2ピックアップ行 ：; [1] A(左側) ST6 反転前行; [2] A(左側) ST6 設置行 *)
    Out_CYw_Rev_02_Pick_A_F_Manual : ARRAY[0..10] OF Bool;  (* 手動【Y715】A(左側)ST6 反転2ピックアップ行 ： *)
    Out_CYw_Rev_02_Pick_A_F_Done : BOOL;  (* 【Y715】A(左側)ST6 反転2ピックアップ行 動作完了 *)
    Out_CYw_Disc_Chk_A_H_Auto : ARRAY[0..10] OF Bool;  (* 自動【Y716】A(左側) 排出チャック閉 戻 ： *)
    Out_CYw_Disc_Chk_A_H_Manual : ARRAY[0..10] OF Bool;  (* 手動【Y716】A(左側) 排出チャック閉 戻 ： *)
    Out_CYw_Disc_Chk_A_H_Done : BOOL;  (* 【Y716】A(左側) 排出チャック閉 戻 動作完了 *)
    Out_CYw_Disc_Chk_A_F_Auto : ARRAY[0..10] OF Bool;  (* 自動【Y717】A(左側) 排出チャック開 行 ： *)
    Out_CYw_Disc_Chk_A_F_Manual : ARRAY[0..10] OF Bool;  (* 手動【Y717】A(左側) 排出チャック開 行 ： *)
    Out_CYw_Disc_Chk_A_F_Done : BOOL;  (* 【Y717】A(左側) 排出チャック開 行 動作完了 *)
    Out_CYw_Ejc_Hldr_Feed_A_F_Auto : ARRAY[0..10] OF Bool;  (* 自動【Y719】A(左側) 排出フォルダ送り行 ： *)
    Out_CYw_Ejc_Hldr_Feed_A_F_Manual : ARRAY[0..10] OF Bool;  (* 手動【Y719】A(左側) 排出フォルダ送り行 ： *)
    Out_CYw_Ejc_Hldr_Feed_A_F_Done : BOOL;  (* 【Y719】A(左側) 排出フォルダ送り行 動作完了 *)
    Out_CYw_Ejc_Hldr_Feed_A_H_Auto : ARRAY[0..10] OF Bool;  (* 自動【Y718】A(左側) 排出フォルダ送り戻 ： *)
    Out_CYw_Ejc_Hldr_Feed_A_H_Manual : ARRAY[0..10] OF Bool;  (* 手動【Y718】A(左側) 排出フォルダ送り戻 ： *)
    Out_CYw_Ejc_Hldr_Feed_A_H_Done : BOOL;  (* 【Y718】A(左側) 排出フォルダ送り戻 動作完了 *)
    Out_CYS_Pos_01_Stopper_A_H_Auto : ARRAY[0..10] OF Bool;  (* 自動【Y720】A(左側) 位置1ストッパー 戻： *)
    Out_CYS_Pos_01_Stopper_A_H_Manual : ARRAY[0..10] OF Bool;  (* 手動【Y720】A(左側) 位置1ストッパー 戻 ： *)
    Out_CYS_Pos_01_Stopper_A_F_Done : BOOL;  (* 【Y720】A(左側) 位置1ストッパー行 動作完了 *)
    Out_CYS_Pos_01_Stopper_A_H_Done : BOOL;  (* 【Y720】A(左側) 位置1ストッパー戻 動作完了 *)
    Out_CYw_HgtInsp_Lf_A_F_Done : BOOL;  (* 【Y703】A(左側) 高さ検査持上行 動作完了 *)
    Out_CYw_NG1_Pick_A_H_Auto : ARRAY[0..10] OF Bool;  (* 自動【Y704】A(左側) NG1ピックアップ戻： *)
    Out_CYw_NG1_Pick_A_H_Manual : ARRAY[0..10] OF Bool;  (* 手動【Y704】A(左側) NG1ピックアップ戻： *)
    Out_CYw_NG1_Pick_A_H_Done : BOOL;  (* 【Y704】A(左側) NG1ピックアップ戻 動作完了 *)
    Out_CYw_NG1_Pick_A_F_Auto : ARRAY[0..10] OF Bool;  (* 自動【Y705】A(左側) NG1ピックアップ 行： *)
    Out_CYw_NG1_Pick_A_F_Manual : ARRAY[0..10] OF Bool;  (* 手動【Y705】A(左側) NG1ピックアップ 行： *)
    Out_CYw_NG1_Pick_A_F_Done : BOOL;  (* 【Y705】A(左側) NG1ピックアップ 動作完了 *)
    Out_CYw_NG1_Chk_A_H_Auto : ARRAY[0..10] OF Bool;  (* 自動【Y706】A(左側) NG1チャック戻 ： *)
    Out_CYw_NG1_Chk_A_H_Manual : ARRAY[0..10] OF Bool;  (* 手動【Y706】A(左側) NG1チャック戻 ： *)
    Out_CYw_NG1_Chk_A_H_Done : BOOL;  (* 【Y706】A(左側) NG1チャック戻 動作完了 *)
    Out_CYw_NG1_Chk_A_F_Auto : ARRAY[0..10] OF Bool;  (* 自動【Y707】A(左側) NG1チャック行： *)
    Out_CYw_NG1_Chk_A_F_Manual : ARRAY[0..10] OF Bool;  (* 手動【Y707】A(左側) NG1チャック行： *)
    Out_CYw_NG1_Chk_A_F_Done : BOOL;  (* 【Y707】A(左側) NG1チャック行 動作完了 *)
    Out_CYw_Rev_01_Chk_A_H_Auto : ARRAY[0..10] OF Bool;  (* 自動【Y708】A(左側)ST4 反転1チャック閉： *)
    Out_CYw_Rev_01_Chk_A_H_Manual : ARRAY[0..10] OF Bool;  (* 手動【Y708】A(左側)ST4 反転1チャック閉： *)
    Out_CYw_Rev_01_Chk_A_H_Done : BOOL;  (* 【Y708】A(左側)ST4 反転1チャック閉 動作完了 *)
    Mtr_Flip_01_Busy : BOOL;  (* A(左側)反転 オリエンタルモータ1 動作中 *)
    Out_CYw_Rev_01_Chk_A_F_Auto : ARRAY[0..10] OF Bool;  (* 自動【Y709】A(左側)ST4 反転1チャック開： *)
    Out_CYw_Rev_01_Chk_A_F_Manual : ARRAY[0..10] OF Bool;  (* 手動【Y709】A(左側)ST4 反転1チャック開： *)
    Out_CYw_Rev_01_Chk_A_F_Done : BOOL;  (* 【Y709】A(左側)ST4 反転1チャック開 動作完了 *)
    Out_CYw_Rev_01_Pick_A_H_Auto : ARRAY[0..10] OF Bool;  (* 自動【Y710】A(左側)ST4 反転1ピックアップ戻： *)
    Out_CYw_Rev_01_Pick_A_H_Manual : ARRAY[0..10] OF Bool;  (* 手動【Y710】A(左側)ST4 反転1ピックアップ戻： *)
    Out_CYw_Rev_01_Pick_A_H_Done : BOOL;  (* 【Y710】A(左側)ST4 反転1ピックアップ戻 動作完了 *)
    Out_CYw_Rev_01_Pick_A_F_Auto : ARRAY[0..10] OF Bool;  (* 自動【Y711】A(左側)ST4 反転1ピックアップ行： *)
    Out_CYw_Rev_01_Pick_A_F_Manual : ARRAY[0..10] OF Bool;  (* 手動【Y711】A(左側)ST4 反転1ピックアップ行： *)
    Out_CYw_Rev_01_Pick_A_F_Done : BOOL;  (* 【Y711】A(左側)ST4 反転1ピックアップ行 動作完了 *)
    Out_CYw_Rev_02_Chk_A_H_Auto : ARRAY[0..10] OF Bool;  (* 自動【Y712】A(左側)ST6 反転2チャック閉 戻： *)
    Out_CYw_Rev_02_Chk_A_H_Manual : ARRAY[0..10] OF Bool;  (* 手動【Y712】A(左側)ST6 反転2チャック閉 戻： *)
    Out_CYw_Rev_02_Chk_A_H_Done : BOOL;  (* 【Y712】A(左側)ST6 反転2チャック閉 戻 動作完了 *)
    Out_CYw_Rev_02_Chk_A_F_Auto : ARRAY[0..10] OF Bool;  (* 自動【Y713】A(左側)ST6 反転2チャック開 行 戻： *)
    Out_CYw_Rev_02_Chk_A_F_Manual : ARRAY[0..10] OF Bool;  (* 手動【Y713】A(左側)ST6 反転2チャック開 行 戻： *)
    Out_CYw_Rev_02_Chk_A_F_Done : BOOL;  (* 【Y713】A(左側)ST6 反転2チャック開 行 動作完了 *)
    Out_CYw_Sply_Slide_B_F_Done : BOOL;  (* 【Y623】B(右側) 供給スライド行 動作完了 *)
    Out_CYw_Sply_Pick_B_H_Auto : ARRAY[0..10] OF Bool;  (* 自動【Y624】B(右側) 供給ピックアップ戻： *)
    Out_CYw_Sply_Pick_B_H_Manual : ARRAY[0..10] OF Bool;  (* 手動【Y624】B(右側) 供給ピックアップ戻： *)
    Out_CYw_Sply_Pick_B_H_Done : BOOL;  (* 【Y624】B(右側) 供給ピックアップ戻 動作完了 *)
    Out_CYw_Sply_Pick_B_F_Auto : ARRAY[0..10] OF Bool;  (* 自動【Y625】B(右側) 供給ピックアップ行： *)
    Out_CYw_Sply_Pick_B_F_Manual : ARRAY[0..10] OF Bool;  (* 手動【Y625】B(右側) 供給ピックアップ行： *)
    Out_CYw_Sply_Pick_B_F_Done : BOOL;  (* 【Y625】B(右側) 供給ピックアップ行 動作完了 *)
    Out_CYw_Sup_Chuck_B_Cl_H_Auto : ARRAY[0..10] OF Bool;  (* 自動【Y626】B(右側) 供給チャック閉 戻： *)
    Out_CYw_Sup_Chuck_B_Cl_H_Manual : ARRAY[0..10] OF Bool;  (* 手動【Y626】B(右側) 供給チャック閉 戻： *)
    Out_CYw_Sup_Chuck_B_Cl_H_Done : BOOL;  (* 【Y626】B(右側) 供給チャック閉 戻 動作完了 *)
    Out_CYw_Sup_Chuck_B_Cl_F_Auto : ARRAY[0..10] OF Bool;  (* 自動【Y627】B(右側) 供給チャック開 行： *)
    Out_CYw_Sup_Chuck_B_Cl_F_Manual : ARRAY[0..10] OF Bool;  (* 手動【Y627】B(右側) 供給チャック開 行： *)
    Out_CYw_Sup_Chuck_B_Cl_F_Done : BOOL;  (* 【Y627】B(右側) 供給チャック開 行 動作完了 *)
    Out_CYw_HgtInsp_Clp_A_H_Auto : ARRAY[0..10] OF Bool;  (* 自動【Y700】A(左側) 高さ検査押え戻： *)
    Out_CYw_HgtInsp_Clp_A_H_Manual : ARRAY[0..10] OF Bool;  (* 手動【Y700】A(左側) 高さ検査押え戻： *)
    Out_CYw_HgtInsp_Clp_A_H_Done : BOOL;  (* 【Y700】A(左側) 高さ検査押え戻 動作完了 *)
    Out_CYw_HgtInsp_Clp_A_F_Auto : ARRAY[0..10] OF Bool;  (* 自動【Y701】A(左側) 高さ検査押え行： *)
    Out_CYw_HgtInsp_Clp_A_F_Manual : ARRAY[0..10] OF Bool;  (* 手動【Y701】A(左側) 高さ検査押え行： *)
    Out_CYw_HgtInsp_Clp_A_F_Done : BOOL;  (* 【Y701】A(左側) 高さ検査押え行 動作完了 *)
    Out_CYw_HgtInsp_Lf_A_H_Auto : ARRAY[0..10] OF Bool;  (* 自動【Y702】A(左側) 高さ検査持上戻： *)
    Out_CYw_HgtInsp_Lf_A_H_Manual : ARRAY[0..10] OF Bool;  (* 手動【Y702】A(左側) 高さ検査持上戻： *)
    Out_CYw_HgtInsp_Lf_A_H_Done : BOOL;  (* 【Y702】A(左側) 高さ検査持上戻 動作完了 *)
    Out_CYw_HgtInsp_Lf_A_F_Auto : ARRAY[0..10] OF Bool;  (* 自動【Y703】A(左側) 高さ検査持上行： *)
    Out_CYw_HgtInsp_Lf_A_F_Manual : ARRAY[0..10] OF Bool;  (* 手動【Y703】A(左側) 高さ検査持上行： *)
    Out_CYw_Sply_Slide_A_F_Auto : ARRAY[0..10] OF Bool;  (* 自動【Y617】A(左側) 供給スライド行： *)
    Out_CYw_Sply_Slide_A_F_Manual : ARRAY[0..10] OF Bool;  (* 手動【Y617】A(左側) 供給スライド行： *)
    Out_CYw_Sply_Pick_A_H_Auto : ARRAY[0..10] OF Bool;  (* 自動【Y618】A(左側) 供給ピックアップ戻： *)
    Out_CYw_Sply_Pick_A_H_Manual : ARRAY[0..10] OF Bool;  (* 手動【Y618】A(左側) 供給ピックアップ戻： *)
    Out_CYw_Sply_Pick_A_H_Done : BOOL;  (* 【Y618】A(左側) 供給ピックアップ戻 動作完了 *)
    Out_CYw_Sply_Pick_A_F_Auto : ARRAY[0..10] OF Bool;  (* 自動【Y619】A(左側) 供給ピックアップ行： *)
    Out_CYw_Sply_Pick_A_F_Manual : ARRAY[0..10] OF Bool;  (* 自動【Y619】A(左側) 供給ピックアップ行： *)
    Out_CYw_Sply_Pick_A_F_Done : BOOL;  (* 【Y619】A(左側) 供給ピックアップ行 動作完了 *)
    Out_CYw_Sup_Chuck_A_Cl_H_Auto : ARRAY[0..10] OF Bool;  (* 自動【Y620】A(左側) 供給チャック閉 戻： *)
    Out_CYw_Sup_Chuck_A_Cl_H_Manual : ARRAY[0..10] OF Bool;  (* 手動【Y620】A(左側) 供給チャック閉 戻： *)
    Out_CYw_Sup_Chuck_A_Cl_H_Done : BOOL;  (* 【Y620】A(左側) 供給チャック閉 戻 動作完了 *)
    Out_CYw_Sup_Chuck_A_Cl_F_Auto : ARRAY[0..10] OF Bool;  (* 自動【Y621】A(左側) 供給チャック開 行： *)
    Out_CYw_Sup_Chuck_A_Cl_F_Manual : ARRAY[0..10] OF Bool;  (* 手動【Y621】A(左側) 供給チャック開 行： *)
    Out_CYw_Sup_Chuck_A_Cl_F_Done : BOOL;  (* 【Y621】A(左側) 供給チャック開 行 動作完了 *)
    Out_CYw_Sply_Slide_B_H_Auto : ARRAY[0..10] OF Bool;  (* 自動【Y622】B(右側) 供給スライド戻： *)
    Out_CYw_Sply_Slide_B_H_Manual : ARRAY[0..10] OF Bool;  (* 手動【Y622】B(右側) 供給スライド行： *)
    Out_CYw_Sply_Slide_B_Done : BOOL;  (* 【Y622】B(右側) 供給スライド戻 動作完了 *)
    Out_CYw_Sply_Slide_B_F_Auto : ARRAY[0..10] OF Bool;  (* 自動【Y623】B(右側) 供給スライド行： *)
    Out_CYw_Sply_Slide_B_F_Manual : ARRAY[0..10] OF Bool;  (* 手動【Y623】B(右側) 供給スライド行： *)
    In_Sen_Accum_CV_B_Full : BOOL;
    In_Sen_Tray_Direction_Check : BOOL;
    TimerQ_In_Sen_Tray_Direction_Check : BOOL;  (* 【X1007】コンテナトレイ方向 *)
    Out_CYw_Rev_01_Pick_A_H_Origin : ARRAY[0..10] OF Bool;  (* 原点復帰【Y710】A(左側)ST4 反転1ピックアップ戻： *)
    Out_CYw_Rev_01_Pick_A_F_Origin : ARRAY[0..99] OF Bool;  (* 原点復帰【Y711】A(左側)ST4 反転1ピックアップ行： *)
    Out_CYw_Rev_01_Chk_A_H_Origin : ARRAY[0..99] OF Bool;  (* 原点復帰【Y708】A(左側)ST4 反転1チャック閉： *)
    Out_CYw_Rev_02_Chk_A_H_Origin : ARRAY[0..99] OF Bool;  (* 原点復帰 【Y712】A(左側)ST6 反転2チャック閉 戻 *)
    Out_CYw_Rev_02_Pick_A_H_Origin : ARRAY[0..10] OF Bool;  (* 原点復帰 【Y714】A(左側)ST6 反転2ピックアップ戻 *)
    Out_CYw_Rev_02_Pick_A_F_Origin : ARRAY[0..99] OF Bool;  (* 原点復帰 【Y715】A(左側)ST6 反転2ピックアップ行 *)
    Out_CYw_Rev_01_Chk_B_H_Origin : ARRAY[0..99] OF Bool;  (* 原点復帰 【Y808】B(右側)ST4 反転1チャック閉 戻 *)
    Out_CYw_Rev_01_Pick_B_H_Origin : ARRAY[0..10] OF Bool;  (* 原点復帰 【Y810】B(右側)ST4 反転1ピックアップ戻 *)
    Out_CYw_Rev_01_Pick_B_F_Origin : ARRAY[0..99] OF Bool;  (* 原点復帰 【Y811】B(右側)ST4 反転1ピックアップ行 *)
    Out_CYw_Rev_02_Chk_B_H_Origin : ARRAY[0..99] OF Bool;  (* 原点復帰 【Y812】B(右側)ST6 反転2チャック閉 戻 *)
    Out_CYw_Rev_02_Pick_B_H_Origin : ARRAY[0..10] OF Bool;  (* 原点復帰 【Y814】B(右側)ST6 反転2ピックアップ戻 *)
    Out_CYw_Rev_02_Pick_B_F_Origin : ARRAY[0..99] OF Bool;  (* 原点復帰 【Y815】B(右側)ST6 反転2ピックアップ行 *)
    RCON1_5_ActualPos_mm : LREAL;
    RCON1_5_SafePos_mm : LREAL;  (* フォルダストック回転可能高さ *)
    HMI_Message_Request : ARRAY[0..121] OF BOOL;  (* #HMI メッセージ表示要求; [0] 未使用; [1] 【Y616】A(左側) 供給スライド戻 異常表示; [2] 【Y617】A(左側) 供給スライド行 異常表示; [3] 【Y618】A(左側) 供給ピックアップ戻 異常表示; [4] 【Y619】A(左側) 供給ピックアップ行 異常表示; [5] 【Y620】A(左側) 供給チャック閉 戻 異常表示; [6] 【Y621】A(左側) 供給チャック開 行 異常表示; [7] 【Y622】B(右側) 供給スライド戻 異常表示; [8] 【Y623】B(右側) 供給スライド行 異常表示; [9] 【Y624】B(右側) 供給ピックアップ戻 異常表示; [10] 【Y625】B(右側) 供給ピックアップ行 異常表示; [11] 【Y626】B(右側) 供給チャック閉 戻 異常表示; [12] 【Y627】B(右側) 供給チャック開 行 異常表示; [13] 【Y700】A(左側) 高さ検査押え戻 異常表示; [14] 【Y701】A(左側) 高さ検査押え行 異常表示; [15] 【Y702】A(左側) 高さ検査持上戻 異常表示; [16] 【Y703】A(左側) 高さ検査持上行 異常表示; [17] 【Y704】A(左側) NG1ピックアップ戻 異常表示; [18] 【Y705】A(左側) NG1ピックアップ 行 異常表示; [19] 【Y706】A(左側) NG1チャック戻 異常表示; [20] 【Y707】A(左側) NG1チャック行 異常表示; [21] 【Y708】A(左側)ST4 反転1チャック閉 異常表示; [22] 【Y709】A(左側)ST4 反転1チャック開 異常表示; [23] 【Y710】A(左側)ST4 反転1ピックアップ戻 異常表示; [24] 【Y711】A(左側)ST4 反転1ピックアップ行 異常表示; [25] 【Y712】A(左側)ST6 反転2チャック閉 戻 異常表示; [26] 【Y713】A(左側)ST6 反転2チャック開 行 異常表示; [27] 【Y714】A(左側)ST6 反転2ピックアップ戻 異常表示; [28] 【Y715】A(左側)ST6 反転2ピックアップ行 異常表示; [29] 【Y716】A(左側) 排出チャック閉 戻 異常表示; [30] 【Y717】A(左側) 排出チャック開 行 異常表示; [31] 【Y718】A(左側) 排出フォルダ送り戻 異常表示; [32] 【Y719】A(左側) 排出フォルダ送り行 異常表示; [33] A(左側) 位置1ストッパー戻 異常表示; [34] 【Y720】A(左側) 位置1ストッパー 行 異常表示; [35] 【Y721】A(左側) 位置2ストッパー 異常表示; [36] 【Y721】A(左側) 位置2ストッパー 異常表示; [37] 【Y722】A(左側) 位置3ストッパー戻 異常表示; [38] 【Y722】A(左側) 位置3ストッパー行 異常表示; [39] Output_A_Error_M[33] 異常表示; [40] 【Y723】A(左側) 位置4ストッパー行 異常表示; [41] 【Y724】A(左側) 位置5ストッパー戻 異常表示; [42] 【Y724】A(左側) 位置5ストッパー行 異常表示; [43] 【Y725】A(左側) 位置6ストッパー戻 異常表示; [44] 【Y725】A(左側) 位置6ストッパー行 異常表示; [45] 【Y726】A(左側) ストックフォルダターン戻 異常表示; [46] 【Y727】A(左側) ストックフォルダターン行 異常表示; [47] 【Y728】A(左側) NG1仕分け 戻 異常表示; [48] 【Y729】A(左側) NG1仕分け 行 異常表示; [49] 【Y800】B(右側) 高さ検査押え戻 異常表示; [50] 【Y801】B(右側) 高さ検査押え行 異常表示; [51] 【Y802】B(右側) 高さ検査持上戻 異常表示; [52] 【Y803】B(右側) 高さ検査持上行 異常表示; [53] 【Y804】B(右側) NG1ピックアップ戻 異常表示; [54] 【Y805】B(右側) NG1ピックアップ 行 異常表示; [55] 【Y806】B(右側) NG1チャック戻 異常表示; [56] 【Y807】B(右側) NG1チャック行 異常表示; [57] 【Y808】B(右側)ST4 反転1チャック閉 戻 異常表示; [58] 【Y809】B(右側)ST4 反転1チャック開 戻 異常表示; [59] 【Y810】B(右側)ST4 反転1ピックアップ戻 異常表示; [60] 【Y811】B(右側)ST4 反転1ピックアップ行 異常表示; [61] 【Y812】B(右側)ST6 反転2チャック閉 戻 異常表示; [62] 【Y813】B(右側)ST6 反転2チャック開 行 異常表示; [63] 【Y814】B(右側)ST6 反転2ピックアップ戻 異常表示; [64] 【Y815】B(右側)ST6 反転2ピックアップ行 異常表示; [65] 【Y816】B(右側) 排出チャック閉 戻 異常表示; [66] 【Y817】B(右側) 排出チャック開 行 異常表示; [67] 【Y818】B(右側) 排出フォルダ送り戻 異常表示; [68] 【Y819】B(右側) 排出フォルダ送り行 異常表示; [69] 【Y820】B(右側) 位置1ストッパー 戻 異常表示; [70] 【Y820】B(右側) 位置1ストッパー 行 異常表示; [71] 【Y821】B(右側) 位置2ストッパー戻 異常表示; [72] 【Y821】B(右側) 位置2ストッパー行 異常表示; [73] 【Y822】B(右側) 位置3ストッパー戻 異常表示; [74] 【Y822】B(右側) 位置3ストッパー行 異常表示; [75] 【Y823】B(右側) 位置4ストッパー戻 異常表示; [76] 【Y823】B(右側) 位置4ストッパー行 異常表示; [77] 【Y824】B(右側) 位置5ストッパー戻 異常表示; [78] 【Y824】B(右側) 位置5ストッパー行 異常表示; [79] 【Y825】B(右側) 位置6ストッパー戻 異常表示; [80] 【Y825】B(右側) 位置6ストッパー行 異常表示; [81] 【Y826】B(右側) ストックフォルダターン戻 異常表示; [82] 【Y827】B(右側) ストックフォルダターン行 異常表示; [83] 【Y828】B(右側) NG1仕分け 戻 異常表示; [84] 【Y829】B(右側) NG1仕分け 行 異常表示; [85] 【Y1200】空コンテナ送り 戻 異常表示; [86] 【Y1201】空コンテナ送り 行 異常表示; [87] 【Y1202】段バラシ爪 戻 異常表示; [88] 【Y1203】段バラシ爪 行 異常表示; [89] 【Y1204】コンテナ排出 戻 異常表示; [90] 【Y1205】コンテナ排出 行 異常表示; [91] Output_Share_Error_M[7] 異常表示; [92] 【Y1207】箱入れチャック 行 異常表示; [93] 【Y1208】コンテナ仕分けストッパー 戻 異常表示; [94] 【Y1209】コンテナ仕分けストッパー 行 異常表示; [95] 【Y1210】コンテナ仕分け送り 戻 異常表示; [96] Output_Share_Error_M[12] 異常表示; [97] 【Y1300】A(左側) コンベア受渡送り戻 異常表示; [98] 【Y1301】A(左側) コンベア受渡送り行 異常表示; [99] 【Y1302】B(右側) コンベア受渡送り戻 異常表示; [100] 【Y1303】B(右側) コンベア受渡送り行 異常表示; [101] ST1 搬送ワーク不一致; [102] ST2 搬送ワーク不一致; [103] ST3 搬送ワーク不一致; [104] ST4 搬送ワーク不一致; [105] ST5 搬送ワーク不一致; [106] ST6 搬送ワーク不一致; [107] ST7 搬送ワーク不一致; [108] A(左側) ST1 FH測定時間超過; [109] A(左側) ST1 FH異常; [110] A(左側) ST5 FH異常; [111] B(右側) ST1 FH異常; [112] B(右側) ST5 FH異常; [113] A(左側) ST1 FH判定OK; [114] A(左側) ST1 FH判定NG1; [115] A(左側) ST1 FH判定NG2; [116] A(左側) ST1 検査前ワーク不一致; [117] A(左側) ST5 FH測定時間超過; [118] A(左側) ST5 FH判定OK; [119] A(左側) ST5 FH判定NG1; [120] A(左側) ST5 FH判定NG2; [121] A(左側) ST5 検査前ワーク不一致 *)
END_VAR
VAR
    _e1 : R_TRIG;
    _e2 : R_TRIG;
    _p3 : BOOL;
    _e4 : R_TRIG;
    _e5 : R_TRIG;
    _e6 : R_TRIG;
    _p7 : BOOL;
    _e8 : R_TRIG;
    _e9 : R_TRIG;
    _e10 : R_TRIG;
    _p11 : BOOL;
    _e12 : R_TRIG;
    _e13 : R_TRIG;
    _e14 : R_TRIG;
    _p15 : BOOL;
    _e16 : R_TRIG;
    _e17 : R_TRIG;
    _e18 : R_TRIG;
    _p19 : BOOL;
    _e20 : R_TRIG;
    _e21 : R_TRIG;
    _e22 : R_TRIG;
    _p23 : BOOL;
    _e24 : R_TRIG;
    _e25 : R_TRIG;
    _e26 : R_TRIG;
    _p27 : BOOL;
    _e28 : R_TRIG;
    _e29 : R_TRIG;
    _e30 : R_TRIG;
    _p31 : BOOL;
    _e32 : R_TRIG;
    _e33 : R_TRIG;
    _e34 : R_TRIG;
    _p35 : BOOL;
    _e36 : R_TRIG;
    _e37 : R_TRIG;
    _e38 : R_TRIG;
    _p39 : BOOL;
    _e40 : R_TRIG;
    _e41 : R_TRIG;
    _e42 : R_TRIG;
    _p43 : BOOL;
    _e44 : R_TRIG;
    _e45 : R_TRIG;
    _e46 : R_TRIG;
    _p47 : BOOL;
    _e48 : R_TRIG;
    _e49 : R_TRIG;
    _e50 : R_TRIG;
    _p51 : BOOL;
    _p52 : BOOL;
    _e53 : R_TRIG;
    _e54 : R_TRIG;
    _e55 : R_TRIG;
    _p56 : BOOL;
    _p57 : BOOL;
    _e58 : R_TRIG;
    _e59 : R_TRIG;
    _e60 : R_TRIG;
    _p61 : BOOL;
    _e62 : R_TRIG;
    _e63 : R_TRIG;
    _e64 : R_TRIG;
    _p65 : BOOL;
    _p66 : BOOL;
    _e67 : R_TRIG;
    _e68 : R_TRIG;
    _e69 : R_TRIG;
    _p70 : BOOL;
    _e71 : R_TRIG;
    _e72 : R_TRIG;
    _e73 : R_TRIG;
    _p74 : BOOL;
    _e75 : R_TRIG;
    _e76 : R_TRIG;
    _e77 : R_TRIG;
    _p78 : BOOL;
    _e79 : R_TRIG;
    _e80 : R_TRIG;
    _e81 : R_TRIG;
    _p82 : BOOL;
    _e83 : R_TRIG;
    _e84 : R_TRIG;
    _e85 : R_TRIG;
    _e86 : R_TRIG;
    _p87 : BOOL;
    _p88 : BOOL;
    _e89 : R_TRIG;
    _e90 : R_TRIG;
    _e91 : R_TRIG;
    _p92 : BOOL;
    _p93 : BOOL;
    _e94 : R_TRIG;
    _e95 : R_TRIG;
    _e96 : R_TRIG;
    _e97 : R_TRIG;
    _p98 : BOOL;
    _p99 : BOOL;
    _e100 : R_TRIG;
    _e101 : R_TRIG;
    _e102 : R_TRIG;
    _e103 : R_TRIG;
    _p104 : BOOL;
    _p105 : BOOL;
    _e106 : R_TRIG;
    _e107 : R_TRIG;
    _e108 : R_TRIG;
    _e109 : R_TRIG;
    _p110 : BOOL;
    _p111 : BOOL;
    _e112 : R_TRIG;
    _e113 : R_TRIG;
    _e114 : R_TRIG;
    _p115 : BOOL;
    _p116 : BOOL;
    _e117 : R_TRIG;
    _e118 : R_TRIG;
    _e119 : R_TRIG;
    _e120 : R_TRIG;
    _p121 : BOOL;
    _p122 : BOOL;
    _e123 : R_TRIG;
    _e124 : R_TRIG;
    _e125 : R_TRIG;
    _e126 : R_TRIG;
    _p127 : BOOL;
    _p128 : BOOL;
    _e129 : R_TRIG;
    _e130 : R_TRIG;
    _e131 : R_TRIG;
    _p132 : BOOL;
    _e133 : R_TRIG;
    _e134 : R_TRIG;
    _e135 : R_TRIG;
    _p136 : BOOL;
    _e137 : R_TRIG;
    _e138 : R_TRIG;
    _e139 : R_TRIG;
    _p140 : BOOL;
    _p141 : BOOL;
    _e142 : R_TRIG;
    _e143 : R_TRIG;
    _e144 : R_TRIG;
    _p145 : BOOL;
    _p146 : BOOL;
    _e147 : R_TRIG;
    _e148 : R_TRIG;
    _e149 : R_TRIG;
    _p150 : BOOL;
    _p151 : BOOL;
    _e152 : R_TRIG;
    _e153 : R_TRIG;
    _e154 : R_TRIG;
    _p155 : BOOL;
    _p156 : BOOL;
    _e157 : R_TRIG;
    _e158 : R_TRIG;
    _e159 : R_TRIG;
    _p160 : BOOL;
    _p161 : BOOL;
    _e162 : R_TRIG;
    _e163 : R_TRIG;
    _e164 : R_TRIG;
    _p165 : BOOL;
    _p166 : BOOL;
    _e167 : R_TRIG;
    _e168 : R_TRIG;
    _e169 : R_TRIG;
    _p170 : BOOL;
    _p171 : BOOL;
    _e172 : R_TRIG;
    _e173 : R_TRIG;
    _e174 : R_TRIG;
    _p175 : BOOL;
    _p176 : BOOL;
    _e177 : R_TRIG;
    _e178 : R_TRIG;
    _e179 : R_TRIG;
    _p180 : BOOL;
    _p181 : BOOL;
    _e182 : R_TRIG;
    _e183 : R_TRIG;
    _e184 : R_TRIG;
    _p185 : BOOL;
    _p186 : BOOL;
    _e187 : R_TRIG;
    _e188 : R_TRIG;
    _e189 : R_TRIG;
    _p190 : BOOL;
    _p191 : BOOL;
    _e192 : R_TRIG;
    _e193 : R_TRIG;
    _e194 : R_TRIG;
    _p195 : BOOL;
    _p196 : BOOL;
    _e197 : R_TRIG;
    _e198 : R_TRIG;
    _e199 : R_TRIG;
    _p200 : BOOL;
    _p201 : BOOL;
    _e202 : R_TRIG;
    _e203 : R_TRIG;
    _e204 : R_TRIG;
    _p205 : BOOL;
    _p206 : BOOL;
    _e207 : R_TRIG;
    _e208 : R_TRIG;
    _e209 : R_TRIG;
    _p210 : BOOL;
    _e211 : R_TRIG;
    _e212 : R_TRIG;
    _e213 : R_TRIG;
    _p214 : BOOL;
    _e215 : R_TRIG;
    _e216 : R_TRIG;
    _e217 : R_TRIG;
    _p218 : BOOL;
    _e219 : R_TRIG;
    _e220 : R_TRIG;
    _e221 : R_TRIG;
    _p222 : BOOL;
    _e223 : R_TRIG;
    _e224 : R_TRIG;
    _e225 : R_TRIG;
    _p226 : BOOL;
    _p227 : BOOL;
    _e228 : R_TRIG;
    _e229 : R_TRIG;
    _e230 : R_TRIG;
    _p231 : BOOL;
    _p232 : BOOL;
    _e233 : R_TRIG;
    _e234 : R_TRIG;
    _e235 : R_TRIG;
    _p236 : BOOL;
    _e237 : R_TRIG;
    _e238 : R_TRIG;
    _e239 : R_TRIG;
    _p240 : BOOL;
    _p241 : BOOL;
    _e242 : R_TRIG;
    _e243 : R_TRIG;
    _e244 : R_TRIG;
    _p245 : BOOL;
    _e246 : R_TRIG;
    _e247 : R_TRIG;
    _e248 : R_TRIG;
    _p249 : BOOL;
    _e250 : R_TRIG;
    _e251 : R_TRIG;
    _e252 : R_TRIG;
    _p253 : BOOL;
    _e254 : R_TRIG;
    _e255 : R_TRIG;
    _e256 : R_TRIG;
    _p257 : BOOL;
    _e258 : R_TRIG;
    _e259 : R_TRIG;
    _e260 : R_TRIG;
    _e261 : R_TRIG;
    _p262 : BOOL;
    _p263 : BOOL;
    _e264 : R_TRIG;
    _e265 : R_TRIG;
    _e266 : R_TRIG;
    _p267 : BOOL;
    _p268 : BOOL;
    _e269 : R_TRIG;
    _e270 : R_TRIG;
    _e271 : R_TRIG;
    _e272 : R_TRIG;
    _p273 : BOOL;
    _p274 : BOOL;
    _e275 : R_TRIG;
    _e276 : R_TRIG;
    _e277 : R_TRIG;
    _e278 : R_TRIG;
    _p279 : BOOL;
    _p280 : BOOL;
    _e281 : R_TRIG;
    _e282 : R_TRIG;
    _e283 : R_TRIG;
    _e284 : R_TRIG;
    _p285 : BOOL;
    _p286 : BOOL;
    _e287 : R_TRIG;
    _e288 : R_TRIG;
    _e289 : R_TRIG;
    _p290 : BOOL;
    _p291 : BOOL;
    _e292 : R_TRIG;
    _e293 : R_TRIG;
    _e294 : R_TRIG;
    _e295 : R_TRIG;
    _p296 : BOOL;
    _p297 : BOOL;
    _e298 : R_TRIG;
    _e299 : R_TRIG;
    _e300 : R_TRIG;
    _e301 : R_TRIG;
    _p302 : BOOL;
    _p303 : BOOL;
    _e304 : R_TRIG;
    _e305 : R_TRIG;
    _e306 : R_TRIG;
    _p307 : BOOL;
    _e308 : R_TRIG;
    _e309 : R_TRIG;
    _e310 : R_TRIG;
    _p311 : BOOL;
    _e312 : R_TRIG;
    _e313 : R_TRIG;
    _e314 : R_TRIG;
    _p315 : BOOL;
    _p316 : BOOL;
    _e317 : R_TRIG;
    _e318 : R_TRIG;
    _e319 : R_TRIG;
    _p320 : BOOL;
    _p321 : BOOL;
    _e322 : R_TRIG;
    _e323 : R_TRIG;
    _e324 : R_TRIG;
    _p325 : BOOL;
    _p326 : BOOL;
    _e327 : R_TRIG;
    _e328 : R_TRIG;
    _e329 : R_TRIG;
    _p330 : BOOL;
    _p331 : BOOL;
    _e332 : R_TRIG;
    _e333 : R_TRIG;
    _e334 : R_TRIG;
    _p335 : BOOL;
    _p336 : BOOL;
    _e337 : R_TRIG;
    _e338 : R_TRIG;
    _e339 : R_TRIG;
    _p340 : BOOL;
    _p341 : BOOL;
    _e342 : R_TRIG;
    _e343 : R_TRIG;
    _e344 : R_TRIG;
    _p345 : BOOL;
    _p346 : BOOL;
    _e347 : R_TRIG;
    _e348 : R_TRIG;
    _e349 : R_TRIG;
    _p350 : BOOL;
    _p351 : BOOL;
    _e352 : R_TRIG;
    _e353 : R_TRIG;
    _e354 : R_TRIG;
    _p355 : BOOL;
    _p356 : BOOL;
    _e357 : R_TRIG;
    _e358 : R_TRIG;
    _e359 : R_TRIG;
    _p360 : BOOL;
    _p361 : BOOL;
    _e362 : R_TRIG;
    _e363 : R_TRIG;
    _e364 : R_TRIG;
    _p365 : BOOL;
    _p366 : BOOL;
    _e367 : R_TRIG;
    _e368 : R_TRIG;
    _e369 : R_TRIG;
    _p370 : BOOL;
    _p371 : BOOL;
    _e372 : R_TRIG;
    _e373 : R_TRIG;
    _e374 : R_TRIG;
    _p375 : BOOL;
    _p376 : BOOL;
    _e377 : R_TRIG;
    _e378 : R_TRIG;
    _e379 : R_TRIG;
    _p380 : BOOL;
    _p381 : BOOL;
    _e382 : R_TRIG;
    _e383 : R_TRIG;
    _e384 : R_TRIG;
    _p385 : BOOL;
    _e386 : R_TRIG;
    _e387 : R_TRIG;
    _e388 : R_TRIG;
    _p389 : BOOL;
    _e390 : R_TRIG;
    _e391 : R_TRIG;
    _e392 : R_TRIG;
    _p393 : BOOL;
    _e394 : R_TRIG;
    _e395 : R_TRIG;
    _e396 : R_TRIG;
    _p397 : BOOL;
    _e398 : R_TRIG;
    _e399 : R_TRIG;
    _e400 : R_TRIG;
    _p401 : BOOL;
    _p402 : BOOL;
    _e403 : R_TRIG;
    _e404 : R_TRIG;
    _e405 : R_TRIG;
    _p406 : BOOL;
    _p407 : BOOL;
    _e408 : R_TRIG;
    _e409 : R_TRIG;
    _e410 : R_TRIG;
    _p411 : BOOL;
    _p412 : BOOL;
    _e413 : R_TRIG;
    _e414 : R_TRIG;
    _e415 : R_TRIG;
    _p416 : BOOL;
    _p417 : BOOL;
    _e418 : R_TRIG;
    _e419 : R_TRIG;
    _e420 : R_TRIG;
    _p421 : BOOL;
    _p422 : BOOL;
    _e423 : R_TRIG;
    _e424 : R_TRIG;
    _e425 : R_TRIG;
    _p426 : BOOL;
    _p427 : BOOL;
    _e428 : R_TRIG;
    _e429 : R_TRIG;
    _e430 : R_TRIG;
    _p431 : BOOL;
    _e432 : R_TRIG;
    _e433 : R_TRIG;
    _e434 : R_TRIG;
    _p435 : BOOL;
    _e436 : R_TRIG;
    _e437 : R_TRIG;
    _e438 : R_TRIG;
    _p439 : BOOL;
    _p440 : BOOL;
    _e441 : R_TRIG;
    _e442 : R_TRIG;
    _e443 : R_TRIG;
    _p444 : BOOL;
    _p445 : BOOL;
    _e446 : R_TRIG;
    _e447 : R_TRIG;
    _e448 : R_TRIG;
    _p449 : BOOL;
    _p450 : BOOL;
    _e451 : R_TRIG;
    _e452 : R_TRIG;
    _e453 : R_TRIG;
    _p454 : BOOL;
    _p455 : BOOL;
    _e456 : R_TRIG;
    _e457 : R_TRIG;
    _e458 : R_TRIG;
    _p459 : BOOL;
    _e460 : R_TRIG;
    _e461 : R_TRIG;
    _e462 : R_TRIG;
    _p463 : BOOL;
    _e464 : R_TRIG;
    _e465 : R_TRIG;
    _e466 : R_TRIG;
    _p467 : BOOL;
    _e468 : R_TRIG;
    _e469 : R_TRIG;
    _e470 : R_TRIG;
    _p471 : BOOL;
    _e472 : R_TRIG;
END_VAR

(* Section Input_入力: ladder, written here as Structured Text *)

